// TIA Portal project "整合" (V18)

(* hardware
DEVICE "S7-1200 station_2"  S7-1200 Station
   slot 0: "Rack_0"  S7-1200 Rack  Rack  V1.0
   slot 1: "PLC_1"  CPU 1214C DC/DC/DC  6ES7 214-1AG40-0XB0  V4.1
DEVICE "PC-System_1"  SIMATIC PC station
   slot 0: "SIMATIC PC station"  Rail  SIMATIC PC-Station  V1.0
      slot 125: "Stationmanager"  Station_Manager  V6.0.4
   slot 1: "HMI_RT_1"  WinCC RT Advanced  6AV2 104-0xxxx-xxxx  17.0.0.0
      slot 33792: "主机接口"  Host interface
   slot 2: "IE general_1"  IE General  IE_CP  V8.2.0
      slot 1: "PROFINET interface"  IEGeneral.Interface.8.2.0
*)

// ===== PLC "PLC_1"  CPU 1214C DC/DC/DC =====

DATA_BLOCK "初始化用"   // DB2
{ S7_Optimized_Access := 'TRUE' }
VERSION : 0.1
// stored: InstanceOfName 初始化
"初始化"
BEGIN
END_DATA_BLOCK

DATA_BLOCK "中间变量2"   // DB3
{ S7_Optimized_Access := 'FALSE' }
VERSION : 0.1
   VAR
      "1梯1层最终调度距离" : Int;
      "2梯1层最终调度距离" : Int;
      "3梯1层最终调度距离" : Int;
      "1层上呼分配1" : Bool;
      "1层上呼分配2" : Bool;
      "1层上呼分配3" : Bool;
      "1层上呼分配4" : Bool;
      "1层上呼分配5" : Bool;
      "1层上呼分配6" : Bool;
      "1梯2层最终调度距离上" : Int;
      "1梯2层最终调度距离下" : Int;
      "2层上呼分配1" : Bool;
      "2层上呼分配2" : Bool;
      "2层上呼分配3" : Bool;
      "2层上呼分配4" : Bool;
      "2层上呼分配5" : Bool;
      "2层上呼分配6" : Bool;
      "2梯2层最终调度距离上" : Int;
      "2梯2层最终调度距离下" : Int;
      "3梯2层最终调度距离上" : Int;
      "3梯2层最终调度距离下" : Int;
      "1梯3层最终调度距离上" : Int;
      "1梯3层最终调度距离下" : Int;
      "2梯3层最终调度距离上" : Int;
      "2梯3层最终调度距离下" : Int;
      "3梯3层最终调度距离上" : Int;
      "3梯3层最终调度距离下" : Int;
      "1梯4层最终调度距离上" : Int;
      "1梯4层最终调度距离下" : Int;
      "2梯4层最终调度距离上" : Int;
      "2梯4层最终调度距离下" : Int;
      "3梯4层最终调度距离上" : Int;
      "3梯4层最终调度距离下" : Int;
      "2层下呼分配1" : Bool;
      "2层下呼分配2" : Bool;
      "2层下呼分配3" : Bool;
      "2层下呼分配4" : Bool;
      "2层下呼分配5" : Bool;
      "2层下呼分配6" : Bool;
      "3层上呼分配1" : Bool;
      "3层上呼分配2" : Bool;
      "3层上呼分配3" : Bool;
      "3层上呼分配4" : Bool;
      "3层上呼分配5" : Bool;
      "3层上呼分配6" : Bool;
      "3层下呼分配1" : Bool;
      "3层下呼分配2" : Bool;
      "3层下呼分配3" : Bool;
      "3层下呼分配4" : Bool;
      "3层下呼分配5" : Bool;
      "3层下呼分配6" : Bool;
      "4层上呼分配1" : Bool;
      "4层上呼分配2" : Bool;
      "4层上呼分配3" : Bool;
      "4层上呼分配4" : Bool;
      "4层上呼分配5" : Bool;
      "4层上呼分配6" : Bool;
      "4层下呼分配1" : Bool;
      "4层下呼分配2" : Bool;
      "4层下呼分配3" : Bool;
      "4层下呼分配4" : Bool;
      "4层下呼分配5" : Bool;
      "4层下呼分配6" : Bool;
      "1梯5层最终调度距离上" : Int;
      "1梯5层最终调度距离下" : Int;
      "2梯5层最终调度距离上" : Int;
      "2梯5层最终调度距离下" : Int;
      "3梯5层最终调度距离上" : Int;
      "3梯5层最终调度距离下" : Int;
      "5层上呼分配1" : Bool;
      "5层上呼分配2" : Bool;
      "5层上呼分配3" : Bool;
      "5层上呼分配4" : Bool;
      "5层上呼分配5" : Bool;
      "5层上呼分配6" : Bool;
      "5层下呼分配1" : Bool;
      "5层下呼分配2" : Bool;
      "5层下呼分配3" : Bool;
      "5层下呼分配4" : Bool;
      "5层下呼分配5" : Bool;
      "5层下呼分配6" : Bool;
      "1梯6层最终调度距离上" : Int;
      "1梯6层最终调度距离下" : Int;
      "2梯6层最终调度距离上" : Int;
      "2梯6层最终调度距离下" : Int;
      "3梯6层最终调度距离上" : Int;
      "3梯6层最终调度距离下" : Int;
      "6层上呼分配1" : Bool;
      "6层上呼分配2" : Bool;
      "6层上呼分配3" : Bool;
      "6层上呼分配4" : Bool;
      "6层上呼分配5" : Bool;
      "6层上呼分配6" : Bool;
      "6层下呼分配1" : Bool;
      "6层下呼分配2" : Bool;
      "6层下呼分配3" : Bool;
      "6层下呼分配4" : Bool;
      "6层下呼分配5" : Bool;
      "6层下呼分配6" : Bool;
      "1梯7层最终调度距离上" : Int;
      "1梯7层最终调度距离下" : Int;
      "2梯7层最终调度距离上" : Int;
      "2梯7层最终调度距离下" : Int;
      "3梯7层最终调度距离上" : Int;
      "3梯7层最终调度距离下" : Int;
      "7层上呼分配1" : Bool;
      "7层上呼分配2" : Bool;
      "7层上呼分配3" : Bool;
      "7层上呼分配4" : Bool;
      "7层上呼分配5" : Bool;
      "7层上呼分配6" : Bool;
      "7层下呼分配1" : Bool;
      "7层下呼分配2" : Bool;
      "7层下呼分配3" : Bool;
      "7层下呼分配4" : Bool;
      "7层下呼分配5" : Bool;
      "7层下呼分配6" : Bool;
      "1梯8层最终调度距离上" : Int;
      "1梯8层最终调度距离下" : Int;
      "2梯8层最终调度距离上" : Int;
      "2梯8层最终调度距离下" : Int;
      "3梯8层最终调度距离上" : Int;
      "3梯8层最终调度距离下" : Int;
      "8层上呼分配1" : Bool;
      "8层上呼分配2" : Bool;
      "8层上呼分配3" : Bool;
      "8层上呼分配4" : Bool;
      "8层上呼分配5" : Bool;
      "8层上呼分配6" : Bool;
      "8层下呼分配1" : Bool;
      "8层下呼分配2" : Bool;
      "8层下呼分配3" : Bool;
      "8层下呼分配4" : Bool;
      "8层下呼分配5" : Bool;
      "8层下呼分配6" : Bool;
      "1梯9层最终调度距离上" : Int;
      "1梯9层最终调度距离下" : Int;
      "2梯9层最终调度距离上" : Int;
      "2梯9层最终调度距离下" : Int;
      "3梯9层最终调度距离上" : Int;
      "3梯9层最终调度距离下" : Int;
      "9层上呼分配1" : Bool;
      "9层上呼分配2" : Bool;
      "9层上呼分配3" : Bool;
      "9层上呼分配4" : Bool;
      "9层上呼分配5" : Bool;
      "9层上呼分配6" : Bool;
      "9层下呼分配1" : Bool;
      "9层下呼分配2" : Bool;
      "9层下呼分配3" : Bool;
      "9层下呼分配4" : Bool;
      "9层下呼分配5" : Bool;
      "9层下呼分配6" : Bool;
      "1梯10层最终调度距离" : Int;
      "2梯10层最终调度距离" : Int;
      "3梯10层最终调度距离" : Int;
      "10层下呼分配1" : Bool;
      "10层下呼分配2" : Bool;
      "10层下呼分配3" : Bool;
      "10层下呼分配4" : Bool;
      "10层下呼分配5" : Bool;
      "10层下呼分配6" : Bool;
      "1号梯外呼上面无目标2" : Bool;
      "1号梯外呼上面无目标3" : Bool;
      "1号梯外呼上面无目标4" : Bool;
      "1号梯外呼上面无目标5" : Bool;
      "1号梯外呼上面无目标6" : Bool;
      "1号梯外呼上面无目标7" : Bool;
      "1号梯外呼上面无目标8" : Bool;
      "1号梯外呼上面无目标9" : Bool;
      "1号梯外呼下面无目标2" : Bool;
      "1号梯外呼下面无目标3" : Bool;
      "1号梯外呼下面无目标4" : Bool;
      "1号梯外呼下面无目标5" : Bool;
      "1号梯外呼下面无目标6" : Bool;
      "1号梯外呼下面无目标7" : Bool;
      "1号梯外呼下面无目标8" : Bool;
      "1号梯外呼下面无目标9" : Bool;
      "2号梯外呼上面无目标2" : Bool;
      "2号梯外呼上面无目标3" : Bool;
      "2号梯外呼上面无目标4" : Bool;
      "2号梯外呼上面无目标5" : Bool;
      "2号梯外呼上面无目标6" : Bool;
      "2号梯外呼上面无目标7" : Bool;
      "2号梯外呼上面无目标8" : Bool;
      "2号梯外呼上面无目标9" : Bool;
      "2号梯外呼下面无目标2" : Bool;
      "2号梯外呼下面无目标3" : Bool;
      "2号梯外呼下面无目标4" : Bool;
      "2号梯外呼下面无目标5" : Bool;
      "2号梯外呼下面无目标6" : Bool;
      "2号梯外呼下面无目标7" : Bool;
      "2号梯外呼下面无目标8" : Bool;
      "2号梯外呼下面无目标9" : Bool;
      "3号梯外呼上面无目标2" : Bool;
      "3号梯外呼上面无目标3" : Bool;
      "3号梯外呼上面无目标4" : Bool;
      "3号梯外呼上面无目标5" : Bool;
      "3号梯外呼上面无目标6" : Bool;
      "3号梯外呼上面无目标7" : Bool;
      "3号梯外呼上面无目标8" : Bool;
      "3号梯外呼上面无目标9" : Bool;
      "3号梯外呼下面无目标2" : Bool;
      "3号梯外呼下面无目标3" : Bool;
      "3号梯外呼下面无目标4" : Bool;
      "3号梯外呼下面无目标5" : Bool;
      "3号梯外呼下面无目标6" : Bool;
      "3号梯外呼下面无目标7" : Bool;
      "3号梯外呼下面无目标8" : Bool;
      "3号梯外呼下面无目标9" : Bool;
      "1号梯外呼上面有目标最大数1" : Int;
      "1号梯外呼上面有目标最大数2" : Int;
      "1号梯外呼上面有目标最大数3" : Int;
      "1号梯外呼上面有目标最大数4" : Int;
      "1号梯外呼上面有目标最大数5" : Int;
      "1号梯外呼上面有目标最大数6" : Int;
      "1号梯外呼上面有目标最大数7" : Int;
      "1号梯外呼上面有目标最大数8" : Int;
      "1号梯外呼上面有目标最大数9" : Int;
      "1号梯外呼下面有目标最小数2" : Int;
      "1号梯外呼下面有目标最小数3" : Int;
      "1号梯外呼下面有目标最小数4" : Int;
      "1号梯外呼下面有目标最小数5" : Int;
      "1号梯外呼下面有目标最小数6" : Int;
      "1号梯外呼下面有目标最小数7" : Int;
      "1号梯外呼下面有目标最小数8" : Int;
      "1号梯外呼下面有目标最小数9" : Int;
      "1号梯外呼下面有目标最小数10" : Int;
      "2号梯外呼上面有目标最大数1" : Int;
      "2号梯外呼上面有目标最大数2" : Int;
      "2号梯外呼上面有目标最大数3" : Int;
      "2号梯外呼上面有目标最大数4" : Int;
      "2号梯外呼上面有目标最大数5" : Int;
      "2号梯外呼上面有目标最大数6" : Int;
      "2号梯外呼上面有目标最大数7" : Int;
      "2号梯外呼上面有目标最大数8" : Int;
      "2号梯外呼上面有目标最大数9" : Int;
      "2号梯外呼下面有目标最小数2" : Int;
      "2号梯外呼下面有目标最小数3" : Int;
      "2号梯外呼下面有目标最小数4" : Int;
      "2号梯外呼下面有目标最小数5" : Int;
      "2号梯外呼下面有目标最小数6" : Int;
      "2号梯外呼下面有目标最小数7" : Int;
      "2号梯外呼下面有目标最小数8" : Int;
      "2号梯外呼下面有目标最小数9" : Int;
      "2号梯外呼下面有目标最小数10" : Int;
      "3号梯外呼上面有目标最大数1" : Int;
      "3号梯外呼上面有目标最大数2" : Int;
      "3号梯外呼上面有目标最大数3" : Int;
      "3号梯外呼上面有目标最大数4" : Int;
      "3号梯外呼上面有目标最大数5" : Int;
      "3号梯外呼上面有目标最大数6" : Int;
      "3号梯外呼上面有目标最大数7" : Int;
      "3号梯外呼上面有目标最大数8" : Int;
      "3号梯外呼上面有目标最大数9" : Int;
      "3号梯外呼下面有目标最小数2" : Int;
      "3号梯外呼下面有目标最小数3" : Int;
      "3号梯外呼下面有目标最小数4" : Int;
      "3号梯外呼下面有目标最小数5" : Int;
      "3号梯外呼下面有目标最小数6" : Int;
      "3号梯外呼下面有目标最小数7" : Int;
      "3号梯外呼下面有目标最小数8" : Int;
      "3号梯外呼下面有目标最小数9" : Int;
      "3号梯外呼下面有目标最小数10" : Int;
      "1号梯外呼上面有目标1" : Bool;
      "1号梯外呼上面有目标2" : Bool;
      "1号梯外呼上面有目标3" : Bool;
      "1号梯外呼上面有目标4" : Bool;
      "1号梯外呼上面有目标5" : Bool;
      "1号梯外呼上面有目标6" : Bool;
      "1号梯外呼上面有目标7" : Bool;
      "1号梯外呼上面有目标8" : Bool;
      "1号梯外呼上面有目标9" : Bool;
      "1号梯外呼下面有目标2" : Bool;
      "1号梯外呼下面有目标3" : Bool;
      "1号梯外呼下面有目标4" : Bool;
      "1号梯外呼下面有目标5" : Bool;
      "1号梯外呼下面有目标6" : Bool;
      "1号梯外呼下面有目标7" : Bool;
      "1号梯外呼下面有目标8" : Bool;
      "1号梯外呼下面有目标9" : Bool;
      "1号梯外呼下面有目标10" : Bool;
      "2号梯外呼上面有目标1" : Bool;
      "2号梯外呼上面有目标2" : Bool;
      "2号梯外呼上面有目标3" : Bool;
      "2号梯外呼上面有目标4" : Bool;
      "2号梯外呼上面有目标5" : Bool;
      "2号梯外呼上面有目标6" : Bool;
      "2号梯外呼上面有目标7" : Bool;
      "2号梯外呼上面有目标8" : Bool;
      "2号梯外呼上面有目标9" : Bool;
      "2号梯外呼下面有目标2" : Bool;
      "2号梯外呼下面有目标3" : Bool;
      "2号梯外呼下面有目标4" : Bool;
      "2号梯外呼下面有目标5" : Bool;
      "2号梯外呼下面有目标6" : Bool;
      "2号梯外呼下面有目标7" : Bool;
      "2号梯外呼下面有目标8" : Bool;
      "2号梯外呼下面有目标9" : Bool;
      "2号梯外呼下面有目标10" : Bool;
      "3号梯外呼上面有目标1" : Bool;
      "3号梯外呼上面有目标2" : Bool;
      "3号梯外呼上面有目标3" : Bool;
      "3号梯外呼上面有目标4" : Bool;
      "3号梯外呼上面有目标5" : Bool;
      "3号梯外呼上面有目标6" : Bool;
      "3号梯外呼上面有目标7" : Bool;
      "3号梯外呼上面有目标8" : Bool;
      "3号梯外呼上面有目标9" : Bool;
      "3号梯外呼下面有目标2" : Bool;
      "3号梯外呼下面有目标3" : Bool;
      "3号梯外呼下面有目标4" : Bool;
      "3号梯外呼下面有目标5" : Bool;
      "3号梯外呼下面有目标6" : Bool;
      "3号梯外呼下面有目标7" : Bool;
      "3号梯外呼下面有目标8" : Bool;
      "3号梯外呼下面有目标9" : Bool;
      "3号梯外呼下面有目标10" : Bool;
      "1号梯上行停站次数3" : Int;
      "1号梯上行停站次数4" : Int;
      "1号梯上行停站次数5" : Int;
      "1号梯上行停站次数6" : Int;
      "1号梯上行停站次数7" : Int;
      "1号梯上行停站次数8" : Int;
      "1号梯上行停站次数9" : Int;
      "1号梯上行停站次数10" : Int;
      "1号梯下行停站次数1" : Int;
      "1号梯下行停站次数2" : Int;
      "1号梯下行停站次数3" : Int;
      "1号梯下行停站次数4" : Int;
      "1号梯下行停站次数5" : Int;
      "1号梯下行停站次数6" : Int;
      "1号梯下行停站次数7" : Int;
      "1号梯下行停站次数8" : Int;
      "2号梯上行停站次数3" : Int;
      "2号梯上行停站次数4" : Int;
      "2号梯上行停站次数5" : Int;
      "2号梯上行停站次数6" : Int;
      "2号梯上行停站次数7" : Int;
      "2号梯上行停站次数8" : Int;
      "2号梯上行停站次数9" : Int;
      "2号梯上行停站次数10" : Int;
      "2号梯下行停站次数1" : Int;
      "2号梯下行停站次数2" : Int;
      "2号梯下行停站次数3" : Int;
      "2号梯下行停站次数4" : Int;
      "2号梯下行停站次数5" : Int;
      "2号梯下行停站次数6" : Int;
      "2号梯下行停站次数7" : Int;
      "2号梯下行停站次数8" : Int;
      "3号梯上行停站次数3" : Int;
      "3号梯上行停站次数4" : Int;
      "3号梯上行停站次数5" : Int;
      "3号梯上行停站次数6" : Int;
      "3号梯上行停站次数7" : Int;
      "3号梯上行停站次数8" : Int;
      "3号梯上行停站次数9" : Int;
      "3号梯上行停站次数10" : Int;
      "3号梯下行停站次数1" : Int;
      "3号梯下行停站次数2" : Int;
      "3号梯下行停站次数3" : Int;
      "3号梯下行停站次数4" : Int;
      "3号梯下行停站次数5" : Int;
      "3号梯下行停站次数6" : Int;
      "3号梯下行停站次数7" : Int;
      "3号梯下行停站次数8" : Int;
      "1号梯上行需折返停站次数10" : Int;
      "2号梯上行需折返停站次数10" : Int;
      "3号梯上行需折返停站次数10" : Int;
      "1号梯下行需折返停站次数1" : Int;
      "2号梯下行需折返停站次数1" : Int;
      "3号梯下行需折返停站次数1" : Int;
      "1号梯当前楼层数" : Int;
      "2号梯当前楼层数" : Int;
      "3号梯当前楼层数" : Int;
      "4号梯当前楼层数" : Int;
      "5号梯当前楼层数" : Int;
      "6号梯当前楼层数" : Int;
      "4梯1层最终调度距离" : Int;
      "4梯10层最终调度距离" : Int;
      "4梯2层最终调度距离上" : Int;
      "4梯2层最终调度距离下" : Int;
      "4梯3层最终调度距离上" : Int;
      "4梯3层最终调度距离下" : Int;
      "4梯4层最终调度距离上" : Int;
      "4梯4层最终调度距离下" : Int;
      "4梯5层最终调度距离上" : Int;
      "4梯5层最终调度距离下" : Int;
      "4梯6层最终调度距离上" : Int;
      "4梯6层最终调度距离下" : Int;
      "4梯7层最终调度距离上" : Int;
      "4梯7层最终调度距离下" : Int;
      "4梯8层最终调度距离上" : Int;
      "4梯8层最终调度距离下" : Int;
      "4梯9层最终调度距离上" : Int;
      "4梯9层最终调度距离下" : Int;
      "4号梯外呼上面无目标2" : Bool;
      "4号梯外呼上面无目标3" : Bool;
      "4号梯外呼上面无目标4" : Bool;
      "4号梯外呼上面无目标5" : Bool;
      "4号梯外呼上面无目标6" : Bool;
      "4号梯外呼上面无目标7" : Bool;
      "4号梯外呼上面无目标8" : Bool;
      "4号梯外呼上面无目标9" : Bool;
      "4号梯外呼下面无目标2" : Bool;
      "4号梯外呼下面无目标3" : Bool;
      "4号梯外呼下面无目标4" : Bool;
      "4号梯外呼下面无目标5" : Bool;
      "4号梯外呼下面无目标6" : Bool;
      "4号梯外呼下面无目标7" : Bool;
      "4号梯外呼下面无目标8" : Bool;
      "4号梯外呼下面无目标9" : Bool;
      "4号梯外呼上面有目标最大数1" : Int;
      "4号梯外呼上面有目标最大数2" : Int;
      "4号梯外呼上面有目标最大数3" : Int;
      "4号梯外呼上面有目标最大数4" : Int;
      "4号梯外呼上面有目标最大数5" : Int;
      "4号梯外呼上面有目标最大数6" : Int;
      "4号梯外呼上面有目标最大数7" : Int;
      "4号梯外呼上面有目标最大数8" : Int;
      "4号梯外呼上面有目标最大数9" : Int;
      "4号梯外呼下面有目标最小数2" : Int;
      "4号梯外呼下面有目标最小数3" : Int;
      "4号梯外呼下面有目标最小数4" : Int;
      "4号梯外呼下面有目标最小数5" : Int;
      "4号梯外呼下面有目标最小数6" : Int;
      "4号梯外呼下面有目标最小数7" : Int;
      "4号梯外呼下面有目标最小数8" : Int;
      "4号梯外呼下面有目标最小数9" : Int;
      "4号梯外呼下面有目标最小数10" : Int;
      "4号梯外呼上面有目标1" : Bool;
      "4号梯外呼上面有目标2" : Bool;
      "4号梯外呼上面有目标3" : Bool;
      "4号梯外呼上面有目标4" : Bool;
      "4号梯外呼上面有目标5" : Bool;
      "4号梯外呼上面有目标6" : Bool;
      "4号梯外呼上面有目标7" : Bool;
      "4号梯外呼上面有目标8" : Bool;
      "4号梯外呼上面有目标9" : Bool;
      "4号梯外呼下面有目标2" : Bool;
      "4号梯外呼下面有目标3" : Bool;
      "4号梯外呼下面有目标4" : Bool;
      "4号梯外呼下面有目标5" : Bool;
      "4号梯外呼下面有目标6" : Bool;
      "4号梯外呼下面有目标7" : Bool;
      "4号梯外呼下面有目标8" : Bool;
      "4号梯外呼下面有目标9" : Bool;
      "4号梯外呼下面有目标10" : Bool;
      "4号梯上行停站次数3" : Int;
      "4号梯上行停站次数4" : Int;
      "4号梯上行停站次数5" : Int;
      "4号梯上行停站次数6" : Int;
      "4号梯上行停站次数7" : Int;
      "4号梯上行停站次数8" : Int;
      "4号梯上行停站次数9" : Int;
      "4号梯上行停站次数10" : Int;
      "4号梯下行停站次数1" : Int;
      "4号梯下行停站次数2" : Int;
      "4号梯下行停站次数3" : Int;
      "4号梯下行停站次数4" : Int;
      "4号梯下行停站次数5" : Int;
      "4号梯下行停站次数6" : Int;
      "4号梯下行停站次数7" : Int;
      "4号梯下行停站次数8" : Int;
      "4号梯上行需折返停站次数10" : Int;
      "4号梯下行需折返停站次数1" : Int;
      "5梯1层最终调度距离" : Int;
      "5梯10层最终调度距离" : Int;
      "5梯2层最终调度距离上" : Int;
      "5梯2层最终调度距离下" : Int;
      "5梯3层最终调度距离上" : Int;
      "5梯3层最终调度距离下" : Int;
      "5梯4层最终调度距离上" : Int;
      "5梯4层最终调度距离下" : Int;
      "5梯5层最终调度距离上" : Int;
      "5梯5层最终调度距离下" : Int;
      "5梯6层最终调度距离上" : Int;
      "5梯6层最终调度距离下" : Int;
      "5梯7层最终调度距离上" : Int;
      "5梯7层最终调度距离下" : Int;
      "5梯8层最终调度距离上" : Int;
      "5梯8层最终调度距离下" : Int;
      "5梯9层最终调度距离上" : Int;
      "5梯9层最终调度距离下" : Int;
      "5号梯外呼上面无目标2" : Bool;
      "5号梯外呼上面无目标3" : Bool;
      "5号梯外呼上面无目标4" : Bool;
      "5号梯外呼上面无目标5" : Bool;
      "5号梯外呼上面无目标6" : Bool;
      "5号梯外呼上面无目标7" : Bool;
      "5号梯外呼上面无目标8" : Bool;
      "5号梯外呼上面无目标9" : Bool;
      "5号梯外呼下面无目标2" : Bool;
      "5号梯外呼下面无目标3" : Bool;
      "5号梯外呼下面无目标4" : Bool;
      "5号梯外呼下面无目标5" : Bool;
      "5号梯外呼下面无目标6" : Bool;
      "5号梯外呼下面无目标7" : Bool;
      "5号梯外呼下面无目标8" : Bool;
      "5号梯外呼下面无目标9" : Bool;
      "5号梯外呼上面有目标最大数1" : Int;
      "5号梯外呼上面有目标最大数2" : Int;
      "5号梯外呼上面有目标最大数3" : Int;
      "5号梯外呼上面有目标最大数4" : Int;
      "5号梯外呼上面有目标最大数5" : Int;
      "5号梯外呼上面有目标最大数6" : Int;
      "5号梯外呼上面有目标最大数7" : Int;
      "5号梯外呼上面有目标最大数8" : Int;
      "5号梯外呼上面有目标最大数9" : Int;
      "5号梯外呼下面有目标最小数2" : Int;
      "5号梯外呼下面有目标最小数3" : Int;
      "5号梯外呼下面有目标最小数4" : Int;
      "5号梯外呼下面有目标最小数5" : Int;
      "5号梯外呼下面有目标最小数6" : Int;
      "5号梯外呼下面有目标最小数7" : Int;
      "5号梯外呼下面有目标最小数8" : Int;
      "5号梯外呼下面有目标最小数9" : Int;
      "5号梯外呼下面有目标最小数10" : Int;
      "5号梯外呼上面有目标1" : Bool;
      "5号梯外呼上面有目标2" : Bool;
      "5号梯外呼上面有目标3" : Bool;
      "5号梯外呼上面有目标4" : Bool;
      "5号梯外呼上面有目标5" : Bool;
      "5号梯外呼上面有目标6" : Bool;
      "5号梯外呼上面有目标7" : Bool;
      "5号梯外呼上面有目标8" : Bool;
      "5号梯外呼上面有目标9" : Bool;
      "5号梯外呼下面有目标2" : Bool;
      "5号梯外呼下面有目标3" : Bool;
      "5号梯外呼下面有目标4" : Bool;
      "5号梯外呼下面有目标5" : Bool;
      "5号梯外呼下面有目标6" : Bool;
      "5号梯外呼下面有目标7" : Bool;
      "5号梯外呼下面有目标8" : Bool;
      "5号梯外呼下面有目标9" : Bool;
      "5号梯外呼下面有目标10" : Bool;
      "5号梯上行停站次数3" : Int;
      "5号梯上行停站次数4" : Int;
      "5号梯上行停站次数5" : Int;
      "5号梯上行停站次数6" : Int;
      "5号梯上行停站次数7" : Int;
      "5号梯上行停站次数8" : Int;
      "5号梯上行停站次数9" : Int;
      "5号梯上行停站次数10" : Int;
      "5号梯下行停站次数1" : Int;
      "5号梯下行停站次数2" : Int;
      "5号梯下行停站次数3" : Int;
      "5号梯下行停站次数4" : Int;
      "5号梯下行停站次数5" : Int;
      "5号梯下行停站次数6" : Int;
      "5号梯下行停站次数7" : Int;
      "5号梯下行停站次数8" : Int;
      "5号梯上行需折返停站次数10" : Int;
      "5号梯下行需折返停站次数1" : Int;
      "6梯1层最终调度距离" : Int;
      "6梯10层最终调度距离" : Int;
      "6梯2层最终调度距离上" : Int;
      "6梯2层最终调度距离下" : Int;
      "6梯3层最终调度距离上" : Int;
      "6梯3层最终调度距离下" : Int;
      "6梯4层最终调度距离上" : Int;
      "6梯4层最终调度距离下" : Int;
      "6梯5层最终调度距离上" : Int;
      "6梯5层最终调度距离下" : Int;
      "6梯6层最终调度距离上" : Int;
      "6梯6层最终调度距离下" : Int;
      "6梯7层最终调度距离上" : Int;
      "6梯7层最终调度距离下" : Int;
      "6梯8层最终调度距离上" : Int;
      "6梯8层最终调度距离下" : Int;
      "6梯9层最终调度距离上" : Int;
      "6梯9层最终调度距离下" : Int;
      "6号梯外呼上面无目标2" : Bool;
      "6号梯外呼上面无目标3" : Bool;
      "6号梯外呼上面无目标4" : Bool;
      "6号梯外呼上面无目标5" : Bool;
      "6号梯外呼上面无目标6" : Bool;
      "6号梯外呼上面无目标7" : Bool;
      "6号梯外呼上面无目标8" : Bool;
      "6号梯外呼上面无目标9" : Bool;
      "6号梯外呼下面无目标2" : Bool;
      "6号梯外呼下面无目标3" : Bool;
      "6号梯外呼下面无目标4" : Bool;
      "6号梯外呼下面无目标5" : Bool;
      "6号梯外呼下面无目标6" : Bool;
      "6号梯外呼下面无目标7" : Bool;
      "6号梯外呼下面无目标8" : Bool;
      "6号梯外呼下面无目标9" : Bool;
      "6号梯外呼上面有目标最大数1" : Int;
      "6号梯外呼上面有目标最大数2" : Int;
      "6号梯外呼上面有目标最大数3" : Int;
      "6号梯外呼上面有目标最大数4" : Int;
      "6号梯外呼上面有目标最大数5" : Int;
      "6号梯外呼上面有目标最大数6" : Int;
      "6号梯外呼上面有目标最大数7" : Int;
      "6号梯外呼上面有目标最大数8" : Int;
      "6号梯外呼上面有目标最大数9" : Int;
      "6号梯外呼下面有目标最小数2" : Int;
      "6号梯外呼下面有目标最小数3" : Int;
      "6号梯外呼下面有目标最小数4" : Int;
      "6号梯外呼下面有目标最小数5" : Int;
      "6号梯外呼下面有目标最小数6" : Int;
      "6号梯外呼下面有目标最小数7" : Int;
      "6号梯外呼下面有目标最小数8" : Int;
      "6号梯外呼下面有目标最小数9" : Int;
      "6号梯外呼下面有目标最小数10" : Int;
      "6号梯外呼上面有目标1" : Bool;
      "6号梯外呼上面有目标2" : Bool;
      "6号梯外呼上面有目标3" : Bool;
      "6号梯外呼上面有目标4" : Bool;
      "6号梯外呼上面有目标5" : Bool;
      "6号梯外呼上面有目标6" : Bool;
      "6号梯外呼上面有目标7" : Bool;
      "6号梯外呼上面有目标8" : Bool;
      "6号梯外呼上面有目标9" : Bool;
      "6号梯外呼下面有目标2" : Bool;
      "6号梯外呼下面有目标3" : Bool;
      "6号梯外呼下面有目标4" : Bool;
      "6号梯外呼下面有目标5" : Bool;
      "6号梯外呼下面有目标6" : Bool;
      "6号梯外呼下面有目标7" : Bool;
      "6号梯外呼下面有目标8" : Bool;
      "6号梯外呼下面有目标9" : Bool;
      "6号梯外呼下面有目标10" : Bool;
      "6号梯上行停站次数3" : Int;
      "6号梯上行停站次数4" : Int;
      "6号梯上行停站次数5" : Int;
      "6号梯上行停站次数6" : Int;
      "6号梯上行停站次数7" : Int;
      "6号梯上行停站次数8" : Int;
      "6号梯上行停站次数9" : Int;
      "6号梯上行停站次数10" : Int;
      "6号梯下行停站次数1" : Int;
      "6号梯下行停站次数2" : Int;
      "6号梯下行停站次数3" : Int;
      "6号梯下行停站次数4" : Int;
      "6号梯下行停站次数5" : Int;
      "6号梯下行停站次数6" : Int;
      "6号梯下行停站次数7" : Int;
      "6号梯下行停站次数8" : Int;
      "6号梯上行需折返停站次数10" : Int;
      "6号梯下行需折返停站次数1" : Int;
      "1号梯转换后载重量" : Int;
      "2号梯转换后载重量" : Int;
      "3号梯转换后载重量" : Int;
      "4号梯转换后载重量" : Int;
      "5号梯转换后载重量" : Int;
      "6号梯转换后载重量" : Int;
      限重分配1 : Int := 900;
      限重分配2 : Int := 1200;
      限重分配3 : Int := 1200;
      限重分配4 : Int := 1200;
      限重分配5 : Int := 1650;
      限重分配6 : Int := 1850;
      就近运动电梯1 : Bool;
      就近运动电梯2 : Bool;
      就近运动电梯3 : Bool;
      就近运动电梯4 : Bool;
      就近运动电梯5 : Bool;
      就近运动电梯6 : Bool;
   END_VAR
BEGIN
END_DATA_BLOCK

DATA_BLOCK "输入"   // DB10
{ S7_Optimized_Access := 'FALSE' }
VERSION : 0.1
   VAR
      "1层上行呼梯按钮" : Bool;
      "2层上行呼梯按钮" : Bool;
      "3层上行呼梯按钮" : Bool;
      "4层上行呼梯按钮" : Bool;
      "5层上行呼梯按钮" : Bool;
      "6层上行呼梯按钮" : Bool;
      "7层上行呼梯按钮" : Bool;
      "8层上行呼梯按钮" : Bool;
      "9层上行呼梯按钮" : Bool;
      "2层下行呼梯按钮" : Bool;
      "3层下行呼梯按钮" : Bool;
      "4层下行呼梯按钮" : Bool;
      "5层下行呼梯按钮" : Bool;
      "6层下行呼梯按钮" : Bool;
      "7层下行呼梯按钮" : Bool;
      "8层下行呼梯按钮" : Bool;
      "9层下行呼梯按钮" : Bool;
      "10层下行呼梯按钮" : Bool;
      "1号梯轿内选层按钮1" : Bool;
      "1号梯轿内选层按钮2" : Bool;
      "1号梯轿内选层按钮3" : Bool;
      "1号梯轿内选层按钮4" : Bool;
      "1号梯轿内选层按钮5" : Bool;
      "1号梯轿内选层按钮6" : Bool;
      "1号梯轿内选层按钮7" : Bool;
      "1号梯轿内选层按钮8" : Bool;
      "1号梯轿内选层按钮9" : Bool;
      "1号梯轿内选层按钮10" : Bool;
      "1号梯轿内开门按钮" : Bool;
      "1号梯轿内关门按钮" : Bool;
      "1号梯光幕信号" : Bool;
      "1号梯检修信号" : Bool;
      "1号梯轿厢门锁信号" : Bool;
      "1号梯1楼层门锁信号" : Bool;
      "1号梯2楼层门锁信号" : Bool;
      "1号梯3楼层门锁信号" : Bool;
      "1号梯4楼层门锁信号" : Bool;
      "1号梯5楼层门锁信号" : Bool;
      "1号梯6楼层门锁信号" : Bool;
      "1号梯7楼层门锁信号" : Bool;
      "1号梯8楼层门锁信号" : Bool;
      "1号梯9楼层门锁信号" : Bool;
      "1号梯10楼层门锁信号" : Bool;
      "1号梯开门到位" : Bool;
      "1号梯关门到位" : Bool;
      "1号梯上平层信号" : Bool;
      "1号梯下平层信号" : Bool;
      "1号梯上端站第1限位" : Bool;
      "1号梯上端站第2限位" : Bool;
      "1号梯下端站第1限位" : Bool;
      "1号梯下端站第2限位" : Bool;
      "2号梯轿内选层按钮1" : Bool;
      "2号梯轿内选层按钮2" : Bool;
      "2号梯轿内选层按钮3" : Bool;
      "2号梯轿内选层按钮4" : Bool;
      "2号梯轿内选层按钮5" : Bool;
      "2号梯轿内选层按钮6" : Bool;
      "2号梯轿内选层按钮7" : Bool;
      "2号梯轿内选层按钮8" : Bool;
      "2号梯轿内选层按钮9" : Bool;
      "2号梯轿内选层按钮10" : Bool;
      "2号梯轿内开门按钮" : Bool;
      "2号梯轿内关门按钮" : Bool;
      "2号梯光幕信号" : Bool;
      "2号梯检修信号" : Bool;
      "2号梯轿厢门锁信号" : Bool;
      "2号梯1楼层门锁信号" : Bool;
      "2号梯2楼层门锁信号" : Bool;
      "2号梯3楼层门锁信号" : Bool;
      "2号梯4楼层门锁信号" : Bool;
      "2号梯5楼层门锁信号" : Bool;
      "2号梯6楼层门锁信号" : Bool;
      "2号梯7楼层门锁信号" : Bool;
      "2号梯8楼层门锁信号" : Bool;
      "2号梯9楼层门锁信号" : Bool;
      "2号梯10楼层门锁信号" : Bool;
      "2号梯开门到位" : Bool;
      "2号梯关门到位" : Bool;
      "2号梯上平层信号" : Bool;
      "2号梯下平层信号" : Bool;
      "2号梯上端站第1限位" : Bool;
      "2号梯上端站第2限位" : Bool;
      "2号梯下端站第1限位" : Bool;
      "2号梯下端站第2限位" : Bool;
      "3号梯轿内选层按钮1" : Bool;
      "3号梯轿内选层按钮2" : Bool;
      "3号梯轿内选层按钮3" : Bool;
      "3号梯轿内选层按钮4" : Bool;
      "3号梯轿内选层按钮5" : Bool;
      "3号梯轿内选层按钮6" : Bool;
      "3号梯轿内选层按钮7" : Bool;
      "3号梯轿内选层按钮8" : Bool;
      "3号梯轿内选层按钮9" : Bool;
      "3号梯轿内选层按钮10" : Bool;
      "3号梯轿内开门按钮" : Bool;
      "3号梯轿内关门按钮" : Bool;
      "3号梯光幕信号" : Bool;
      "3号梯检修信号" : Bool;
      "3号梯轿厢门锁信号" : Bool;
      "3号梯1楼层门锁信号" : Bool;
      "3号梯2楼层门锁信号" : Bool;
      "3号梯3楼层门锁信号" : Bool;
      "3号梯4楼层门锁信号" : Bool;
      "3号梯5楼层门锁信号" : Bool;
      "3号梯6楼层门锁信号" : Bool;
      "3号梯7楼层门锁信号" : Bool;
      "3号梯8楼层门锁信号" : Bool;
      "3号梯9楼层门锁信号" : Bool;
      "3号梯10楼层门锁信号" : Bool;
      "3号梯开门到位" : Bool;
      "3号梯关门到位" : Bool;
      "3号梯上平层信号" : Bool;
      "3号梯下平层信号" : Bool;
      "3号梯上端站第1限位" : Bool;
      "3号梯上端站第2限位" : Bool;
      "3号梯下端站第1限位" : Bool;
      "3号梯下端站第2限位" : Bool;
      "4号梯轿内选层按钮1" : Bool;
      "4号梯轿内选层按钮2" : Bool;
      "4号梯轿内选层按钮3" : Bool;
      "4号梯轿内选层按钮4" : Bool;
      "4号梯轿内选层按钮5" : Bool;
      "4号梯轿内选层按钮6" : Bool;
      "4号梯轿内选层按钮7" : Bool;
      "4号梯轿内选层按钮8" : Bool;
      "4号梯轿内选层按钮9" : Bool;
      "4号梯轿内选层按钮10" : Bool;
      "4号梯轿内开门按钮" : Bool;
      "4号梯轿内关门按钮" : Bool;
      "4号梯光幕信号" : Bool;
      "4号梯检修信号" : Bool;
      "4号梯轿厢门锁信号" : Bool;
      "4号梯1楼层门锁信号" : Bool;
      "4号梯2楼层门锁信号" : Bool;
      "4号梯3楼层门锁信号" : Bool;
      "4号梯4楼层门锁信号" : Bool;
      "4号梯5楼层门锁信号" : Bool;
      "4号梯6楼层门锁信号" : Bool;
      "4号梯7楼层门锁信号" : Bool;
      "4号梯8楼层门锁信号" : Bool;
      "4号梯9楼层门锁信号" : Bool;
      "4号梯10楼层门锁信号" : Bool;
      "4号梯开门到位" : Bool;
      "4号梯关门到位" : Bool;
      "4号梯上平层信号" : Bool;
      "4号梯下平层信号" : Bool;
      "4号梯上端站第1限位" : Bool;
      "4号梯上端站第2限位" : Bool;
      "4号梯下端站第1限位" : Bool;
      "4号梯下端站第2限位" : Bool;
      "5号梯轿内选层按钮1" : Bool;
      "5号梯轿内选层按钮2" : Bool;
      "5号梯轿内选层按钮3" : Bool;
      "5号梯轿内选层按钮4" : Bool;
      "5号梯轿内选层按钮5" : Bool;
      "5号梯轿内选层按钮6" : Bool;
      "5号梯轿内选层按钮7" : Bool;
      "5号梯轿内选层按钮8" : Bool;
      "5号梯轿内选层按钮9" : Bool;
      "5号梯轿内选层按钮10" : Bool;
      "5号梯轿内开门按钮" : Bool;
      "5号梯轿内关门按钮" : Bool;
      "5号梯光幕信号" : Bool;
      "5号梯检修信号" : Bool;
      "5号梯轿厢门锁信号" : Bool;
      "5号梯1楼层门锁信号" : Bool;
      "5号梯2楼层门锁信号" : Bool;
      "5号梯3楼层门锁信号" : Bool;
      "5号梯4楼层门锁信号" : Bool;
      "5号梯5楼层门锁信号" : Bool;
      "5号梯6楼层门锁信号" : Bool;
      "5号梯7楼层门锁信号" : Bool;
      "5号梯8楼层门锁信号" : Bool;
      "5号梯9楼层门锁信号" : Bool;
      "5号梯10楼层门锁信号" : Bool;
      "5号梯开门到位" : Bool;
      "5号梯关门到位" : Bool;
      "5号梯上平层信号" : Bool;
      "5号梯下平层信号" : Bool;
      "5号梯上端站第1限位" : Bool;
      "5号梯上端站第2限位" : Bool;
      "5号梯下端站第1限位" : Bool;
      "5号梯下端站第2限位" : Bool;
      "6号梯轿内选层按钮1" : Bool;
      "6号梯轿内选层按钮2" : Bool;
      "6号梯轿内选层按钮3" : Bool;
      "6号梯轿内选层按钮4" : Bool;
      "6号梯轿内选层按钮5" : Bool;
      "6号梯轿内选层按钮6" : Bool;
      "6号梯轿内选层按钮7" : Bool;
      "6号梯轿内选层按钮8" : Bool;
      "6号梯轿内选层按钮9" : Bool;
      "6号梯轿内选层按钮10" : Bool;
      "6号梯轿内开门按钮" : Bool;
      "6号梯轿内关门按钮" : Bool;
      "6号梯光幕信号" : Bool;
      "6号梯检修信号" : Bool;
      "6号梯轿厢门锁信号" : Bool;
      "6号梯1楼层门锁信号" : Bool;
      "6号梯2楼层门锁信号" : Bool;
      "6号梯3楼层门锁信号" : Bool;
      "6号梯4楼层门锁信号" : Bool;
      "6号梯5楼层门锁信号" : Bool;
      "6号梯6楼层门锁信号" : Bool;
      "6号梯7楼层门锁信号" : Bool;
      "6号梯8楼层门锁信号" : Bool;
      "6号梯9楼层门锁信号" : Bool;
      "6号梯10楼层门锁信号" : Bool;
      "6号梯开门到位" : Bool;
      "6号梯关门到位" : Bool;
      "6号梯上平层信号" : Bool;
      "6号梯下平层信号" : Bool;
      "6号梯上端站第1限位" : Bool;
      "6号梯上端站第2限位" : Bool;
      "6号梯下端站第1限位" : Bool;
      "6号梯下端站第2限位" : Bool;
      自动运行信号 : Bool;
      "1号梯当前载重量" : Word;
      "2号梯当前载重量" : Word;
      "3号梯当前载重量" : Word;
      "4号梯当前载重量" : Word;
      "5号梯当前载重量" : Word;
      "6号梯当前载重量" : Word;
   END_VAR
BEGIN
END_DATA_BLOCK

DATA_BLOCK "输出"   // DB11
{ S7_Optimized_Access := 'FALSE' }
VERSION : 0.1
   VAR
      "1层上行呼梯按钮指示灯" : Bool;
      "2层上行呼梯按钮指示灯" : Bool;
      "3层上行呼梯按钮指示灯" : Bool;
      "4层上行呼梯按钮指示灯" : Bool;
      "5层上行呼梯按钮指示灯" : Bool;
      "6层上行呼梯按钮指示灯" : Bool;
      "7层上行呼梯按钮指示灯" : Bool;
      "8层上行呼梯按钮指示灯" : Bool;
      "9层上行呼梯按钮指示灯" : Bool;
      "2层下行呼梯按钮指示灯" : Bool;
      "3层下行呼梯按钮指示灯" : Bool;
      "4层下行呼梯按钮指示灯" : Bool;
      "5层下行呼梯按钮指示灯" : Bool;
      "6层下行呼梯按钮指示灯" : Bool;
      "7层下行呼梯按钮指示灯" : Bool;
      "8层下行呼梯按钮指示灯" : Bool;
      "9层下行呼梯按钮指示灯" : Bool;
      "10层下行呼梯按钮指示灯" : Bool;
      "1号梯1层按钮指示灯" : Bool;
      "1号梯2层按钮指示灯" : Bool;
      "1号梯3层按钮指示灯" : Bool;
      "1号梯4层按钮指示灯" : Bool;
      "1号梯5层按钮指示灯" : Bool;
      "1号梯6层按钮指示灯" : Bool;
      "1号梯7层按钮指示灯" : Bool;
      "1号梯8层按钮指示灯" : Bool;
      "1号梯9层按钮指示灯" : Bool;
      "1号梯10层按钮指示灯" : Bool;
      "1号梯LEDa" : Bool;
      "1号梯LEDb" : Bool;
      "1号梯LEDc" : Bool;
      "1号梯LEDd" : Bool;
      "1号梯LEDe" : Bool;
      "1号梯LEDf" : Bool;
      "1号梯LEDg" : Bool;
      "1号梯LEDh" : Bool;
      "1号梯LEDi" : Bool;
      "1号梯LEDj" : Bool;
      "1号梯LEDk" : Bool;
      "1号梯LEDl" : Bool;
      "1号梯LEDm" : Bool;
      "1号梯LEDn" : Bool;
      "1号梯上行指示" : Bool;
      "1号梯下行指示" : Bool;
      "1号梯故障指示" : Bool;
      "1号梯照明指示" : Bool;
      "1号梯风扇指示" : Bool;
      "1号梯满载指示" : Bool;
      "1号梯电机启动信号" : Bool;
      "1号梯上行接触器" : Bool;
      "1号梯下行接触器" : Bool;
      "1号梯高速接触器" : Bool;
      "1号梯低速接触器" : Bool;
      "1号梯开门继电器" : Bool;
      "1号梯关门继电器" : Bool;
      "1号梯1级减速制动" : Bool;
      "1号梯2级减速制动" : Bool;
      "1号梯3级减速制动" : Bool;
      "2号梯1层按钮指示灯" : Bool;
      "2号梯2层按钮指示灯" : Bool;
      "2号梯3层按钮指示灯" : Bool;
      "2号梯4层按钮指示灯" : Bool;
      "2号梯5层按钮指示灯" : Bool;
      "2号梯6层按钮指示灯" : Bool;
      "2号梯7层按钮指示灯" : Bool;
      "2号梯8层按钮指示灯" : Bool;
      "2号梯9层按钮指示灯" : Bool;
      "2号梯10层按钮指示灯" : Bool;
      "2号梯LEDa" : Bool;
      "2号梯LEDb" : Bool;
      "2号梯LEDc" : Bool;
      "2号梯LEDd" : Bool;
      "2号梯LEDe" : Bool;
      "2号梯LEDf" : Bool;
      "2号梯LEDg" : Bool;
      "2号梯LEDh" : Bool;
      "2号梯LEDi" : Bool;
      "2号梯LEDj" : Bool;
      "2号梯LEDk" : Bool;
      "2号梯LEDl" : Bool;
      "2号梯LEDm" : Bool;
      "2号梯LEDn" : Bool;
      "2号梯上行指示" : Bool;
      "2号梯下行指示" : Bool;
      "2号梯故障指示" : Bool;
      "2号梯照明指示" : Bool;
      "2号梯风扇指示" : Bool;
      "2号梯满载指示" : Bool;
      "2号梯电机启动信号" : Bool;
      "2号梯上行接触器" : Bool;
      "2号梯下行接触器" : Bool;
      "2号梯高速接触器" : Bool;
      "2号梯低速接触器" : Bool;
      "2号梯开门继电器" : Bool;
      "2号梯关门继电器" : Bool;
      "2号梯1级减速制动" : Bool;
      "2号梯2级减速制动" : Bool;
      "2号梯3级减速制动" : Bool;
      "3号梯1层按钮指示灯" : Bool;
      "3号梯2层按钮指示灯" : Bool;
      "3号梯3层按钮指示灯" : Bool;
      "3号梯4层按钮指示灯" : Bool;
      "3号梯5层按钮指示灯" : Bool;
      "3号梯6层按钮指示灯" : Bool;
      "3号梯7层按钮指示灯" : Bool;
      "3号梯8层按钮指示灯" : Bool;
      "3号梯9层按钮指示灯" : Bool;
      "3号梯10层按钮指示灯" : Bool;
      "3号梯LEDa" : Bool;
      "3号梯LEDb" : Bool;
      "3号梯LEDc" : Bool;
      "3号梯LEDd" : Bool;
      "3号梯LEDe" : Bool;
      "3号梯LEDf" : Bool;
      "3号梯LEDg" : Bool;
      "3号梯LEDh" : Bool;
      "3号梯LEDi" : Bool;
      "3号梯LEDj" : Bool;
      "3号梯LEDk" : Bool;
      "3号梯LEDl" : Bool;
      "3号梯LEDm" : Bool;
      "3号梯LEDn" : Bool;
      "3号梯上行指示" : Bool;
      "3号梯下行指示" : Bool;
      "3号梯故障指示" : Bool;
      "3号梯照明指示" : Bool;
      "3号梯风扇指示" : Bool;
      "3号梯满载指示" : Bool;
      "3号梯电机启动信号" : Bool;
      "3号梯上行接触器" : Bool;
      "3号梯下行接触器" : Bool;
      "3号梯高速接触器" : Bool;
      "3号梯低速接触器" : Bool;
      "3号梯开门继电器" : Bool;
      "3号梯关门继电器" : Bool;
      "3号梯1级减速制动" : Bool;
      "3号梯2级减速制动" : Bool;
      "3号梯3级减速制动" : Bool;
      "4号梯1层按钮指示灯" : Bool;
      "4号梯2层按钮指示灯" : Bool;
      "4号梯3层按钮指示灯" : Bool;
      "4号梯4层按钮指示灯" : Bool;
      "4号梯5层按钮指示灯" : Bool;
      "4号梯6层按钮指示灯" : Bool;
      "4号梯7层按钮指示灯" : Bool;
      "4号梯8层按钮指示灯" : Bool;
      "4号梯9层按钮指示灯" : Bool;
      "4号梯10层按钮指示灯" : Bool;
      "4号梯LEDa" : Bool;
      "4号梯LEDb" : Bool;
      "4号梯LEDc" : Bool;
      "4号梯LEDd" : Bool;
      "4号梯LEDe" : Bool;
      "4号梯LEDf" : Bool;
      "4号梯LEDg" : Bool;
      "4号梯LEDh" : Bool;
      "4号梯LEDi" : Bool;
      "4号梯LEDj" : Bool;
      "4号梯LEDk" : Bool;
      "4号梯LEDl" : Bool;
      "4号梯LEDm" : Bool;
      "4号梯LEDn" : Bool;
      "4号梯上行指示" : Bool;
      "4号梯下行指示" : Bool;
      "4号梯故障指示" : Bool;
      "4号梯照明指示" : Bool;
      "4号梯风扇指示" : Bool;
      "4号梯满载指示" : Bool;
      "4号梯电机启动信号" : Bool;
      "4号梯上行接触器" : Bool;
      "4号梯下行接触器" : Bool;
      "4号梯高速接触器" : Bool;
      "4号梯低速接触器" : Bool;
      "4号梯开门继电器" : Bool;
      "4号梯关门继电器" : Bool;
      "4号梯1级减速制动" : Bool;
      "4号梯2级减速制动" : Bool;
      "4号梯3级减速制动" : Bool;
      "5号梯1层按钮指示灯" : Bool;
      "5号梯2层按钮指示灯" : Bool;
      "5号梯3层按钮指示灯" : Bool;
      "5号梯4层按钮指示灯" : Bool;
      "5号梯5层按钮指示灯" : Bool;
      "5号梯6层按钮指示灯" : Bool;
      "5号梯7层按钮指示灯" : Bool;
      "5号梯8层按钮指示灯" : Bool;
      "5号梯9层按钮指示灯" : Bool;
      "5号梯10层按钮指示灯" : Bool;
      "5号梯LEDa" : Bool;
      "5号梯LEDb" : Bool;
      "5号梯LEDc" : Bool;
      "5号梯LEDd" : Bool;
      "5号梯LEDe" : Bool;
      "5号梯LEDf" : Bool;
      "5号梯LEDg" : Bool;
      "5号梯LEDh" : Bool;
      "5号梯LEDi" : Bool;
      "5号梯LEDj" : Bool;
      "5号梯LEDk" : Bool;
      "5号梯LEDl" : Bool;
      "5号梯LEDm" : Bool;
      "5号梯LEDn" : Bool;
      "5号梯上行指示" : Bool;
      "5号梯下行指示" : Bool;
      "5号梯故障指示" : Bool;
      "5号梯照明指示" : Bool;
      "5号梯风扇指示" : Bool;
      "5号梯满载指示" : Bool;
      "5号梯电机启动信号" : Bool;
      "5号梯上行接触器" : Bool;
      "5号梯下行接触器" : Bool;
      "5号梯高速接触器" : Bool;
      "5号梯低速接触器" : Bool;
      "5号梯开门继电器" : Bool;
      "5号梯关门继电器" : Bool;
      "5号梯1级减速制动" : Bool;
      "5号梯2级减速制动" : Bool;
      "5号梯3级减速制动" : Bool;
      "6号梯1层按钮指示灯" : Bool;
      "6号梯2层按钮指示灯" : Bool;
      "6号梯3层按钮指示灯" : Bool;
      "6号梯4层按钮指示灯" : Bool;
      "6号梯5层按钮指示灯" : Bool;
      "6号梯6层按钮指示灯" : Bool;
      "6号梯7层按钮指示灯" : Bool;
      "6号梯8层按钮指示灯" : Bool;
      "6号梯9层按钮指示灯" : Bool;
      "6号梯10层按钮指示灯" : Bool;
      "6号梯LEDa" : Bool;
      "6号梯LEDb" : Bool;
      "6号梯LEDc" : Bool;
      "6号梯LEDd" : Bool;
      "6号梯LEDe" : Bool;
      "6号梯LEDf" : Bool;
      "6号梯LEDg" : Bool;
      "6号梯LEDh" : Bool;
      "6号梯LEDi" : Bool;
      "6号梯LEDj" : Bool;
      "6号梯LEDk" : Bool;
      "6号梯LEDl" : Bool;
      "6号梯LEDm" : Bool;
      "6号梯LEDn" : Bool;
      "6号梯上行指示" : Bool;
      "6号梯下行指示" : Bool;
      "6号梯故障指示" : Bool;
      "6号梯照明指示" : Bool;
      "6号梯风扇指示" : Bool;
      "6号梯满载指示" : Bool;
      "6号梯电机启动信号" : Bool;
      "6号梯上行接触器" : Bool;
      "6号梯下行接触器" : Bool;
      "6号梯高速接触器" : Bool;
      "6号梯低速接触器" : Bool;
      "6号梯开门继电器" : Bool;
      "6号梯关门继电器" : Bool;
      "6号梯1级减速制动" : Bool;
      "6号梯2级减速制动" : Bool;
      "6号梯3级减速制动" : Bool;
      准备就绪信号 : Bool;
   END_VAR
BEGIN
END_DATA_BLOCK

DATA_BLOCK "中间变量1"   // DB13
{ S7_Optimized_Access := 'FALSE' }
VERSION : 0.1
   VAR
      "1号梯高速初始化" : Bool;
      "2号梯高速初始化" : Bool;
      "3号梯高速初始化" : Bool;
      "4号梯高速初始化" : Bool;
      "5号梯高速初始化" : Bool;
      "6号梯高速初始化" : Bool;
      是否高速1 : Bool;
      是否高速2 : Bool;
      是否高速3 : Bool;
      是否高速4 : Bool;
      是否高速5 : Bool;
      是否高速6 : Bool;
      高速延时1 : Time;
      高速延时2 : Time;
      高速延时3 : Time;
      高速延时4 : Time;
      高速延时5 : Time;
      高速延时6 : Time;
      上下平层同时为1梯1 : Bool;
      上下平层同时为1梯2 : Bool;
      上下平层同时为1梯3 : Bool;
      上下平层同时为1梯4 : Bool;
      上下平层同时为1梯5 : Bool;
      上下平层同时为1梯6 : Bool;
      特殊上行将要停梯1 : Bool;
      特殊上行将要停梯2 : Bool;
      特殊上行将要停梯3 : Bool;
      特殊上行将要停梯4 : Bool;
      特殊上行将要停梯5 : Bool;
      特殊上行将要停梯6 : Bool;
      特殊下行将要停梯1 : Bool;
      特殊下行将要停梯2 : Bool;
      特殊下行将要停梯3 : Bool;
      特殊下行将要停梯4 : Bool;
      特殊下行将要停梯5 : Bool;
      特殊下行将要停梯6 : Bool;
      "1号梯正处于故障中" : Bool;
      "2号梯正处于故障中" : Bool;
      "3号梯正处于故障中" : Bool;
      "4号梯正处于故障中" : Bool;
      "5号梯正处于故障中" : Bool;
      "6号梯正处于故障中" : Bool;
      "1号梯存在安全隐患（光幕）" : Bool;
      "2号梯存在安全隐患（光幕）" : Bool;
      "3号梯存在安全隐患（光幕）" : Bool;
      "4号梯存在安全隐患（光幕）" : Bool;
      "5号梯存在安全隐患（光幕）" : Bool;
      "6号梯存在安全隐患（光幕）" : Bool;
      "1号梯当前楼层数" : Int;
      "2号梯当前楼层数" : Int;
      "3号梯当前楼层数" : Int;
      "4号梯当前楼层数" : Int;
      "5号梯当前楼层数" : Int;
      "6号梯当前楼层数" : Int;
      "1号梯初始化楼层数" : Int := 1;
      "2号梯初始化楼层数" : Int := 1;
      "3号梯初始化楼层数" : Int := 10;
      "4号梯初始化楼层数" : Int := 10;
      "5号梯初始化楼层数" : Int := 10;
      "6号梯初始化楼层数" : Int := 10;
      "1号梯是否到达端限" : Bool;
      "2号梯是否到达端限" : Bool;
      "3号梯是否到达端限" : Bool;
      "4号梯是否到达端限" : Bool;
      "5号梯是否到达端限" : Bool;
      "6号梯是否到达端限" : Bool;
      "1号梯初始化方向上行" : Bool;
      "2号梯初始化方向上行" : Bool;
      "3号梯初始化方向上行" : Bool;
      "4号梯初始化方向上行" : Bool;
      "5号梯初始化方向上行" : Bool;
      "6号梯初始化方向上行" : Bool;
      "1号梯初始化方向下行" : Bool;
      "2号梯初始化方向下行" : Bool;
      "3号梯初始化方向下行" : Bool;
      "4号梯初始化方向下行" : Bool;
      "5号梯初始化方向下行" : Bool;
      "6号梯初始化方向下行" : Bool;
      检修方向上行1 : Bool;
      检修方向上行2 : Bool;
      检修方向上行3 : Bool;
      检修方向上行4 : Bool;
      检修方向上行5 : Bool;
      检修方向上行6 : Bool;
      检修方向下行1 : Bool;
      检修方向下行2 : Bool;
      检修方向下行3 : Bool;
      检修方向下行4 : Bool;
      检修方向下行5 : Bool;
      检修方向下行6 : Bool;
      "1号梯初始化低速运行" : Bool;
      "2号梯初始化低速运行" : Bool;
      "3号梯初始化低速运行" : Bool;
      "4号梯初始化低速运行" : Bool;
      "5号梯初始化低速运行" : Bool;
      "6号梯初始化低速运行" : Bool;
      "1号梯初始化上行接触器" : Bool;
      "2号梯初始化上行接触器" : Bool;
      "3号梯初始化上行接触器" : Bool;
      "4号梯初始化上行接触器" : Bool;
      "5号梯初始化上行接触器" : Bool;
      "6号梯初始化上行接触器" : Bool;
      "1号梯初始化下行接触器" : Bool;
      "2号梯初始化下行接触器" : Bool;
      "3号梯初始化下行接触器" : Bool;
      "4号梯初始化下行接触器" : Bool;
      "5号梯初始化下行接触器" : Bool;
      "6号梯初始化下行接触器" : Bool;
      "1号梯停梯截断(置0完成关门）" : Bool;
      "2号梯停梯截断(置0完成关门）" : Bool;
      "3号梯停梯截断(置0完成关门）" : Bool;
      "4号梯停梯截断(置0完成关门）" : Bool;
      "5号梯停梯截断(置0完成关门）" : Bool;
      "6号梯停梯截断(置0完成关门）" : Bool;
      "1号梯停梯截断(置0完成开门）" : Bool;
      "2号梯停梯截断(置0完成开门）" : Bool;
      "3号梯停梯截断(置0完成开门）" : Bool;
      "4号梯停梯截断(置0完成开门）" : Bool;
      "5号梯停梯截断(置0完成开门）" : Bool;
      "6号梯停梯截断(置0完成开门）" : Bool;
      "1号梯置0为完成开门" : Bool;
      "2号梯置0为完成开门" : Bool;
      "3号梯置0为完成开门" : Bool;
      "4号梯置0为完成开门" : Bool;
      "5号梯置0为完成开门" : Bool;
      "6号梯置0为完成开门" : Bool;
      "1号梯置0为完成关门" : Bool;
      "2号梯置0为完成关门" : Bool;
      "3号梯置0为完成关门" : Bool;
      "4号梯置0为完成关门" : Bool;
      "5号梯置0为完成关门" : Bool;
      "6号梯置0为完成关门" : Bool;
      "1号梯转换" : Real;
      "2号梯转换" : Real;
      "3号梯转换" : Real;
      "4号梯转换" : Real;
      "5号梯转换" : Real;
      "6号梯转换" : Real;
      "1号梯载重限额" : Int := 1050;
      "2号梯载重限额" : Int := 1350;
      "3号梯载重限额" : Int := 1350;
      "4号梯载重限额" : Int := 1350;
      "5号梯载重限额" : Int := 1800;
      "6号梯载重限额" : Int := 2000;
      "1号梯准备就绪" : Bool;
      "2号梯准备就绪" : Bool;
      "3号梯准备就绪" : Bool;
      "4号梯准备就绪" : Bool;
      "5号梯准备就绪" : Bool;
      "6号梯准备就绪" : Bool;
      "1号梯将要停梯" : Bool;
      "2号梯将要停梯" : Bool;
      "3号梯将要停梯" : Bool;
      "4号梯将要停梯" : Bool;
      "5号梯将要停梯" : Bool;
      "6号梯将要停梯" : Bool;
      "1号梯初始化将要停梯" : Bool;
      "2号梯初始化将要停梯" : Bool;
      "3号梯初始化将要停梯" : Bool;
      "4号梯初始化将要停梯" : Bool;
      "5号梯初始化将要停梯" : Bool;
      "6号梯初始化将要停梯" : Bool;
      初始化1级制动 : Bool;
      初始化2级制动 : Bool;
      初始化3级制动 : Bool;
      卡顿上行1 : Bool;
      卡顿上行2 : Bool;
      卡顿上行3 : Bool;
      卡顿上行4 : Bool;
      卡顿上行5 : Bool;
      卡顿上行6 : Bool;
      卡顿下行1 : Bool;
      卡顿下行2 : Bool;
      卡顿下行3 : Bool;
      卡顿下行4 : Bool;
      卡顿下行5 : Bool;
      卡顿下行6 : Bool;
      卡顿制速1 : Bool;
      卡顿制速2 : Bool;
      卡顿制速3 : Bool;
      卡顿制速4 : Bool;
      卡顿制速5 : Bool;
      卡顿制速6 : Bool;
      到达初始化楼层1号梯 : Bool;
      到达初始化楼层2号梯 : Bool;
      到达初始化楼层3号梯 : Bool;
      到达初始化楼层4号梯 : Bool;
      到达初始化楼层5号梯 : Bool;
      到达初始化楼层6号梯 : Bool;
      死机1 : Bool;
      死机2 : Bool;
      死机3 : Bool;
      死机4 : Bool;
      死机5 : Bool;
      死机6 : Bool;
      截下 : Bool;
      截上 : Bool;
      疑似满载1 : Int;
      疑似满载2 : Int;
      疑似满载3 : Int;
      疑似满载4 : Int;
      疑似满载5 : Int;
      "1号梯初始化方向位" : Int;
      "2号梯初始化方向位" : Int;
      "3号梯初始化方向位" : Int;
      "4号梯初始化方向位" : Int;
      "5号梯初始化方向位" : Int;
      "6号梯初始化方向位" : Int;
      "1号梯初始化方向位选择" : Bool;
      "2号梯初始化方向位选择" : Bool;
      "3号梯初始化方向位选择" : Bool;
      "4号梯初始化方向位选择" : Bool;
      "5号梯初始化方向位选择" : Bool;
      "6号梯初始化方向位选择" : Bool;
      疑似满载6 : Int;
      "1号梯正确楼层数" : Int;
      "2号梯正确楼层数" : Int;
      "3号梯正确楼层数" : Int;
      "4号梯正确楼层数" : Int;
      "5号梯正确楼层数" : Int;
      "6号梯正确楼层数" : Int;
      程序运行时长秒 : Int;
      程序运行时长分钟 : Int;
      程序运行时长小时 : Int;
      程序运行时长 : Time_Of_Day;
      程序运行时长初始量 : Time_Of_Day;
      时间累加器最长时长 : Time := T#99999999ms;
      小时复位 : Bool;
      分钟复位 : Bool;
      秒复位 : Bool;
   END_VAR
BEGIN
END_DATA_BLOCK

// folder: 1号梯

DATA_BLOCK "1号梯初始化"   // DB1
{ S7_Optimized_Access := 'TRUE' }
VERSION : 0.1
// stored: InstanceOfName 初始化
"初始化"
BEGIN
END_DATA_BLOCK

DATA_BLOCK "1号梯距离调度"   // DB4
{ S7_Optimized_Access := 'TRUE' }
VERSION : 0.1
// stored: InstanceOfName 距离调度
"距离调度"
BEGIN
END_DATA_BLOCK

DATA_BLOCK "1号梯指示灯"   // DB6
{ S7_Optimized_Access := 'TRUE' }
VERSION : 0.1
// stored: InstanceOfName 照明，风扇，数码管
"照明，风扇，数码管"
BEGIN
END_DATA_BLOCK

DATA_BLOCK "1号梯停层次数"   // DB7
{ S7_Optimized_Access := 'TRUE' }
VERSION : 0.1
// stored: InstanceOfName 停层次数判断
"停层次数判断"
BEGIN
END_DATA_BLOCK

DATA_BLOCK "1号梯高低速转换"   // DB9
{ S7_Optimized_Access := 'TRUE' }
VERSION : 0.1
// stored: InstanceOfName 高低速转换
"高低速转换"
BEGIN
END_DATA_BLOCK

DATA_BLOCK "1号梯上下行与制动"   // DB16
{ S7_Optimized_Access := 'TRUE' }
VERSION : 0.1
// stored: InstanceOfName 上下行和制动
"上下行和制动"
BEGIN
END_DATA_BLOCK

DATA_BLOCK "1号梯优先级"   // DB18
{ S7_Optimized_Access := 'TRUE' }
VERSION : 0.1
// stored: InstanceOfName 优先级响应开关门
"优先级响应开关门"
BEGIN
END_DATA_BLOCK

DATA_BLOCK "1号梯楼层计算"   // DB20
{ S7_Optimized_Access := 'TRUE' }
VERSION : 0.1
// stored: InstanceOfName 楼层计算
"楼层计算"
BEGIN
END_DATA_BLOCK

DATA_BLOCK "1号梯有无目标判断"   // DB24
{ S7_Optimized_Access := 'TRUE' }
VERSION : 0.1
// stored: InstanceOfName 目标判断
"目标判断"
BEGIN
END_DATA_BLOCK

// folder: 2号梯

DATA_BLOCK "2号梯初始化"   // DB14
{ S7_Optimized_Access := 'TRUE' }
VERSION : 0.1
// stored: InstanceOfName 初始化
"初始化"
BEGIN
END_DATA_BLOCK

DATA_BLOCK "2号梯高低速转换"   // DB15
{ S7_Optimized_Access := 'TRUE' }
VERSION : 0.1
// stored: InstanceOfName 高低速转换
"高低速转换"
BEGIN
END_DATA_BLOCK

DATA_BLOCK "2号梯上下行与制动"   // DB44
{ S7_Optimized_Access := 'TRUE' }
VERSION : 0.1
// stored: InstanceOfName 上下行和制动
"上下行和制动"
BEGIN
END_DATA_BLOCK

DATA_BLOCK "2号梯距离调度"   // DB49
{ S7_Optimized_Access := 'TRUE' }
VERSION : 0.1
// stored: InstanceOfName 距离调度
"距离调度"
BEGIN
END_DATA_BLOCK

DATA_BLOCK "2号梯停层次数"   // DB54
{ S7_Optimized_Access := 'TRUE' }
VERSION : 0.1
// stored: InstanceOfName 停层次数判断
"停层次数判断"
BEGIN
END_DATA_BLOCK

DATA_BLOCK "2号梯楼层计算"   // DB59
{ S7_Optimized_Access := 'TRUE' }
VERSION : 0.1
// stored: InstanceOfName 楼层计算
"楼层计算"
BEGIN
END_DATA_BLOCK

DATA_BLOCK "2号梯优先级"   // DB64
{ S7_Optimized_Access := 'TRUE' }
VERSION : 0.1
// stored: InstanceOfName 优先级响应开关门
"优先级响应开关门"
BEGIN
END_DATA_BLOCK

DATA_BLOCK "2号梯指示灯"   // DB69
{ S7_Optimized_Access := 'TRUE' }
VERSION : 0.1
// stored: InstanceOfName 照明，风扇，数码管
"照明，风扇，数码管"
BEGIN
END_DATA_BLOCK

DATA_BLOCK "2号梯有无目标判断"   // DB74
{ S7_Optimized_Access := 'TRUE' }
VERSION : 0.1
// stored: InstanceOfName 目标判断
"目标判断"
BEGIN
END_DATA_BLOCK

// folder: 3号梯

DATA_BLOCK "3号梯初始化"   // DB17
{ S7_Optimized_Access := 'TRUE' }
VERSION : 0.1
// stored: InstanceOfName 初始化
"初始化"
BEGIN
END_DATA_BLOCK

DATA_BLOCK "3号梯高低速转换"   // DB40
{ S7_Optimized_Access := 'TRUE' }
VERSION : 0.1
// stored: InstanceOfName 高低速转换
"高低速转换"
BEGIN
END_DATA_BLOCK

DATA_BLOCK "3号梯上下行与制动"   // DB45
{ S7_Optimized_Access := 'TRUE' }
VERSION : 0.1
// stored: InstanceOfName 上下行和制动
"上下行和制动"
BEGIN
END_DATA_BLOCK

DATA_BLOCK "3号梯距离调度"   // DB50
{ S7_Optimized_Access := 'TRUE' }
VERSION : 0.1
// stored: InstanceOfName 距离调度
"距离调度"
BEGIN
END_DATA_BLOCK

DATA_BLOCK "3号梯停层次数"   // DB55
{ S7_Optimized_Access := 'TRUE' }
VERSION : 0.1
// stored: InstanceOfName 停层次数判断
"停层次数判断"
BEGIN
END_DATA_BLOCK

DATA_BLOCK "3号梯楼层计算"   // DB60
{ S7_Optimized_Access := 'TRUE' }
VERSION : 0.1
// stored: InstanceOfName 楼层计算
"楼层计算"
BEGIN
END_DATA_BLOCK

DATA_BLOCK "3号梯优先级"   // DB65
{ S7_Optimized_Access := 'TRUE' }
VERSION : 0.1
// stored: InstanceOfName 优先级响应开关门
"优先级响应开关门"
BEGIN
END_DATA_BLOCK

DATA_BLOCK "3号梯指示灯"   // DB70
{ S7_Optimized_Access := 'TRUE' }
VERSION : 0.1
// stored: InstanceOfName 照明，风扇，数码管
"照明，风扇，数码管"
BEGIN
END_DATA_BLOCK

DATA_BLOCK "3号梯有无目标判断"   // DB75
{ S7_Optimized_Access := 'TRUE' }
VERSION : 0.1
// stored: InstanceOfName 目标判断
"目标判断"
BEGIN
END_DATA_BLOCK

// folder: 4号梯

DATA_BLOCK "4号梯初始化"   // DB19
{ S7_Optimized_Access := 'TRUE' }
VERSION : 0.1
// stored: InstanceOfName 初始化
"初始化"
BEGIN
END_DATA_BLOCK

DATA_BLOCK "4号梯高低速转换"   // DB41
{ S7_Optimized_Access := 'TRUE' }
VERSION : 0.1
// stored: InstanceOfName 高低速转换
"高低速转换"
BEGIN
END_DATA_BLOCK

DATA_BLOCK "4号梯上下行与制动"   // DB46
{ S7_Optimized_Access := 'TRUE' }
VERSION : 0.1
// stored: InstanceOfName 上下行和制动
"上下行和制动"
BEGIN
END_DATA_BLOCK

DATA_BLOCK "4号梯距离调度"   // DB51
{ S7_Optimized_Access := 'TRUE' }
VERSION : 0.1
// stored: InstanceOfName 距离调度
"距离调度"
BEGIN
END_DATA_BLOCK

DATA_BLOCK "4号梯停层次数"   // DB56
{ S7_Optimized_Access := 'TRUE' }
VERSION : 0.1
// stored: InstanceOfName 停层次数判断
"停层次数判断"
BEGIN
END_DATA_BLOCK

DATA_BLOCK "4号梯楼层计算"   // DB61
{ S7_Optimized_Access := 'TRUE' }
VERSION : 0.1
// stored: InstanceOfName 楼层计算
"楼层计算"
BEGIN
END_DATA_BLOCK

DATA_BLOCK "4号梯优先级"   // DB66
{ S7_Optimized_Access := 'TRUE' }
VERSION : 0.1
// stored: InstanceOfName 优先级响应开关门
"优先级响应开关门"
BEGIN
END_DATA_BLOCK

DATA_BLOCK "4号梯指示灯"   // DB71
{ S7_Optimized_Access := 'TRUE' }
VERSION : 0.1
// stored: InstanceOfName 照明，风扇，数码管
"照明，风扇，数码管"
BEGIN
END_DATA_BLOCK

DATA_BLOCK "4号梯有无目标判断"   // DB76
{ S7_Optimized_Access := 'TRUE' }
VERSION : 0.1
// stored: InstanceOfName 目标判断
"目标判断"
BEGIN
END_DATA_BLOCK

// folder: 5号梯

DATA_BLOCK "5号梯初始化"   // DB22
{ S7_Optimized_Access := 'TRUE' }
VERSION : 0.1
// stored: InstanceOfName 初始化
"初始化"
BEGIN
END_DATA_BLOCK

DATA_BLOCK "5号梯高低速转换"   // DB42
{ S7_Optimized_Access := 'TRUE' }
VERSION : 0.1
// stored: InstanceOfName 初始化低速模式
"初始化低速模式"
BEGIN
END_DATA_BLOCK

DATA_BLOCK "5号梯上下行与制动"   // DB47
{ S7_Optimized_Access := 'TRUE' }
VERSION : 0.1
// stored: InstanceOfName 上下行和制动
"上下行和制动"
BEGIN
END_DATA_BLOCK

DATA_BLOCK "5号梯距离调度"   // DB52
{ S7_Optimized_Access := 'TRUE' }
VERSION : 0.1
// stored: InstanceOfName 距离调度
"距离调度"
BEGIN
END_DATA_BLOCK

DATA_BLOCK "5号梯停层次数"   // DB57
{ S7_Optimized_Access := 'TRUE' }
VERSION : 0.1
// stored: InstanceOfName 停层次数判断
"停层次数判断"
BEGIN
END_DATA_BLOCK

DATA_BLOCK "5号梯楼层计算"   // DB62
{ S7_Optimized_Access := 'TRUE' }
VERSION : 0.1
// stored: InstanceOfName 楼层计算
"楼层计算"
BEGIN
END_DATA_BLOCK

DATA_BLOCK "5号梯优先级"   // DB67
{ S7_Optimized_Access := 'TRUE' }
VERSION : 0.1
// stored: InstanceOfName 优先级响应开关门
"优先级响应开关门"
BEGIN
END_DATA_BLOCK

DATA_BLOCK "5号梯指示灯"   // DB72
{ S7_Optimized_Access := 'TRUE' }
VERSION : 0.1
// stored: InstanceOfName 照明，风扇，数码管
"照明，风扇，数码管"
BEGIN
END_DATA_BLOCK

DATA_BLOCK "5号梯有无目标判断"   // DB77
{ S7_Optimized_Access := 'TRUE' }
VERSION : 0.1
// stored: InstanceOfName 目标判断
"目标判断"
BEGIN
END_DATA_BLOCK

DATA_BLOCK "5号梯高低速切换"   // DB80
{ S7_Optimized_Access := 'TRUE' }
VERSION : 0.1
// stored: InstanceOfName 高低速转换
"高低速转换"
BEGIN
END_DATA_BLOCK

// folder: 6号梯

DATA_BLOCK "6号梯初始化"   // DB23
{ S7_Optimized_Access := 'TRUE' }
VERSION : 0.1
// stored: InstanceOfName 初始化
"初始化"
BEGIN
END_DATA_BLOCK

DATA_BLOCK "6号梯高低速转换"   // DB43
{ S7_Optimized_Access := 'TRUE' }
VERSION : 0.1
// stored: InstanceOfName 初始化低速模式
"初始化低速模式"
BEGIN
END_DATA_BLOCK

DATA_BLOCK "6号梯上下行与制动"   // DB48
{ S7_Optimized_Access := 'TRUE' }
VERSION : 0.1
// stored: InstanceOfName 上下行和制动
"上下行和制动"
BEGIN
END_DATA_BLOCK

DATA_BLOCK "6号梯距离调度"   // DB53
{ S7_Optimized_Access := 'TRUE' }
VERSION : 0.1
// stored: InstanceOfName 距离调度
"距离调度"
BEGIN
END_DATA_BLOCK

DATA_BLOCK "6号梯停层次数"   // DB58
{ S7_Optimized_Access := 'TRUE' }
VERSION : 0.1
// stored: InstanceOfName 停层次数判断
"停层次数判断"
BEGIN
END_DATA_BLOCK

DATA_BLOCK "6号梯楼层计算"   // DB63
{ S7_Optimized_Access := 'TRUE' }
VERSION : 0.1
// stored: InstanceOfName 楼层计算
"楼层计算"
BEGIN
END_DATA_BLOCK

DATA_BLOCK "6号梯优先级"   // DB68
{ S7_Optimized_Access := 'TRUE' }
VERSION : 0.1
// stored: InstanceOfName 优先级响应开关门
"优先级响应开关门"
BEGIN
END_DATA_BLOCK

DATA_BLOCK "6号梯指示灯"   // DB73
{ S7_Optimized_Access := 'TRUE' }
VERSION : 0.1
// stored: InstanceOfName 照明，风扇，数码管
"照明，风扇，数码管"
BEGIN
END_DATA_BLOCK

DATA_BLOCK "6号梯有无目标判断"   // DB78
{ S7_Optimized_Access := 'TRUE' }
VERSION : 0.1
// stored: InstanceOfName 目标判断
"目标判断"
BEGIN
END_DATA_BLOCK

DATA_BLOCK "6号梯高低速切换"   // DB82
{ S7_Optimized_Access := 'TRUE' }
VERSION : 0.1
// stored: InstanceOfName 高低速转换
"高低速转换"
BEGIN
END_DATA_BLOCK

// folder: System blocks/Program resources

DATA_BLOCK "1号梯初始化置位延时"   // DB21
{ S7_Optimized_Access := 'TRUE' }
AUTHOR : Simatic
FAMILY : IEC
NAME : IEC_TMR
VERSION : 1.0
// stored: InstanceOfName IEC_TIMER
"IEC_TIMER"
BEGIN
END_DATA_BLOCK

DATA_BLOCK "2号梯初始化置位延时"   // DB79
{ S7_Optimized_Access := 'TRUE' }
AUTHOR : Simatic
FAMILY : IEC
NAME : IEC_TMR
VERSION : 1.0
// stored: InstanceOfName IEC_TIMER
"IEC_TIMER"
BEGIN
END_DATA_BLOCK

DATA_BLOCK "3号梯初始化置位延时"   // DB81
{ S7_Optimized_Access := 'TRUE' }
AUTHOR : Simatic
FAMILY : IEC
NAME : IEC_TMR
VERSION : 1.0
// stored: InstanceOfName IEC_TIMER
"IEC_TIMER"
BEGIN
END_DATA_BLOCK

DATA_BLOCK "4号梯初始化置位延时"   // DB83
{ S7_Optimized_Access := 'TRUE' }
AUTHOR : Simatic
FAMILY : IEC
NAME : IEC_TMR
VERSION : 1.0
// stored: InstanceOfName IEC_TIMER
"IEC_TIMER"
BEGIN
END_DATA_BLOCK

DATA_BLOCK "接通延时"   // DB84
{ S7_Optimized_Access := 'TRUE' }
AUTHOR : Simatic
FAMILY : IEC
NAME : IEC_TMR
VERSION : 1.0
// stored: InstanceOfName IEC_TIMER
"IEC_TIMER"
BEGIN
END_DATA_BLOCK

DATA_BLOCK "5号梯初始化置位延时"   // DB85
{ S7_Optimized_Access := 'TRUE' }
AUTHOR : Simatic
FAMILY : IEC
NAME : IEC_TMR
VERSION : 1.0
// stored: InstanceOfName IEC_TIMER
"IEC_TIMER"
BEGIN
END_DATA_BLOCK

DATA_BLOCK "6号梯初始化置位延时"   // DB87
{ S7_Optimized_Access := 'TRUE' }
AUTHOR : Simatic
FAMILY : IEC
NAME : IEC_TMR
VERSION : 1.0
// stored: InstanceOfName IEC_TIMER
"IEC_TIMER"
BEGIN
END_DATA_BLOCK

DATA_BLOCK "每秒脉冲生成器"   // DB91
{ S7_Optimized_Access := 'TRUE' }
AUTHOR : Simatic
FAMILY : IEC
NAME : IEC_TMR
VERSION : 1.0
// stored: InstanceOfName IEC_TIMER
"IEC_TIMER"
BEGIN
END_DATA_BLOCK

DATA_BLOCK "脉冲计数小时"   // DB93
{ S7_Optimized_Access := 'TRUE' }
AUTHOR : Simatic
FAMILY : IEC
NAME : CNTR
VERSION : 1.0
// stored: InstanceOfName IEC_COUNTER
"IEC_COUNTER"
BEGIN
END_DATA_BLOCK

DATA_BLOCK "脉冲计数秒"   // DB94
{ S7_Optimized_Access := 'TRUE' }
AUTHOR : Simatic
FAMILY : IEC
NAME : CNTR
VERSION : 1.0
// stored: InstanceOfName IEC_COUNTER
"IEC_COUNTER"
BEGIN
END_DATA_BLOCK

DATA_BLOCK "脉冲计数分钟"   // DB95
{ S7_Optimized_Access := 'TRUE' }
AUTHOR : Simatic
FAMILY : IEC
NAME : CNTR
VERSION : 1.0
// stored: InstanceOfName IEC_COUNTER
"IEC_COUNTER"
BEGIN
END_DATA_BLOCK

// folder: 距离比较

DATA_BLOCK "1层上呼距离比较"   // DB5
{ S7_Optimized_Access := 'TRUE' }
VERSION : 0.1
// stored: InstanceOfName 距离比较
"距离比较"
BEGIN
END_DATA_BLOCK

DATA_BLOCK "2层上呼距离比较"   // DB8
{ S7_Optimized_Access := 'TRUE' }
VERSION : 0.1
// stored: InstanceOfName 距离比较
"距离比较"
BEGIN
END_DATA_BLOCK

DATA_BLOCK "2层下呼距离比较"   // DB12
{ S7_Optimized_Access := 'TRUE' }
VERSION : 0.1
// stored: InstanceOfName 距离比较
"距离比较"
BEGIN
END_DATA_BLOCK

DATA_BLOCK "3层上呼距离比较"   // DB25
{ S7_Optimized_Access := 'TRUE' }
VERSION : 0.1
// stored: InstanceOfName 距离比较
"距离比较"
BEGIN
END_DATA_BLOCK

DATA_BLOCK "3层下呼距离比较"   // DB26
{ S7_Optimized_Access := 'TRUE' }
VERSION : 0.1
// stored: InstanceOfName 距离比较
"距离比较"
BEGIN
END_DATA_BLOCK

DATA_BLOCK "4层上呼距离比较"   // DB27
{ S7_Optimized_Access := 'TRUE' }
VERSION : 0.1
// stored: InstanceOfName 距离比较
"距离比较"
BEGIN
END_DATA_BLOCK

DATA_BLOCK "4层下呼距离比较"   // DB28
{ S7_Optimized_Access := 'TRUE' }
VERSION : 0.1
// stored: InstanceOfName 距离比较
"距离比较"
BEGIN
END_DATA_BLOCK

DATA_BLOCK "5层上呼距离比较"   // DB29
{ S7_Optimized_Access := 'TRUE' }
VERSION : 0.1
// stored: InstanceOfName 距离比较
"距离比较"
BEGIN
END_DATA_BLOCK

DATA_BLOCK "5层下呼距离比较"   // DB30
{ S7_Optimized_Access := 'TRUE' }
VERSION : 0.1
// stored: InstanceOfName 距离比较
"距离比较"
BEGIN
END_DATA_BLOCK

DATA_BLOCK "6层上呼距离比较"   // DB31
{ S7_Optimized_Access := 'TRUE' }
VERSION : 0.1
// stored: InstanceOfName 距离比较
"距离比较"
BEGIN
END_DATA_BLOCK

DATA_BLOCK "6层下呼距离比较"   // DB32
{ S7_Optimized_Access := 'TRUE' }
VERSION : 0.1
// stored: InstanceOfName 距离比较
"距离比较"
BEGIN
END_DATA_BLOCK

DATA_BLOCK "7层上呼距离比较"   // DB33
{ S7_Optimized_Access := 'TRUE' }
VERSION : 0.1
// stored: InstanceOfName 距离比较
"距离比较"
BEGIN
END_DATA_BLOCK

DATA_BLOCK "7层下呼距离比较"   // DB34
{ S7_Optimized_Access := 'TRUE' }
VERSION : 0.1
// stored: InstanceOfName 距离比较
"距离比较"
BEGIN
END_DATA_BLOCK

DATA_BLOCK "8层上呼距离比较"   // DB35
{ S7_Optimized_Access := 'TRUE' }
VERSION : 0.1
// stored: InstanceOfName 距离比较
"距离比较"
BEGIN
END_DATA_BLOCK

DATA_BLOCK "8层下行距离比较"   // DB36
{ S7_Optimized_Access := 'TRUE' }
VERSION : 0.1
// stored: InstanceOfName 距离比较
"距离比较"
BEGIN
END_DATA_BLOCK

DATA_BLOCK "9层上呼距离比较"   // DB37
{ S7_Optimized_Access := 'TRUE' }
VERSION : 0.1
// stored: InstanceOfName 距离比较
"距离比较"
BEGIN
END_DATA_BLOCK

DATA_BLOCK "9层下呼距离比较"   // DB38
{ S7_Optimized_Access := 'TRUE' }
VERSION : 0.1
// stored: InstanceOfName 距离比较
"距离比较"
BEGIN
END_DATA_BLOCK

DATA_BLOCK "10层下行距离比较"   // DB39
{ S7_Optimized_Access := 'TRUE' }
VERSION : 0.1
// stored: InstanceOfName 距离比较
"距离比较"
BEGIN
END_DATA_BLOCK

// folder: (top level)

FUNCTION_BLOCK "距离比较"   // FB1, LAD
{ S7_Optimized_Access := 'TRUE' }
VERSION : 0.1
   VAR_INPUT
      上下平层同时为1梯1 : Bool;
      上下平层同时为1梯2 : Bool;
      上下平层同时为1梯3 : Bool;
      上下平层同时为1梯4 : Bool;
      上下平层同时为1梯5 : Bool;
      上下平层同时为1梯6 : Bool;
      有外呼楼层内选1 : Bool;
      有外呼楼层内选2 : Bool;
      有外呼楼层内选3 : Bool;
      有外呼楼层内选4 : Bool;
      有外呼楼层内选5 : Bool;
      有外呼楼层内选6 : Bool;
      就近运动电梯1 : Bool;
      就近运动电梯2 : Bool;
      就近运动电梯3 : Bool;
      就近运动电梯4 : Bool;
      就近运动电梯5 : Bool;
      就近运动电梯6 : Bool;
      呼灯 : Bool;
      调度距离1 : Int;
      调度距离2 : Int;
      调度距离3 : Int;
      调度距离4 : Int;
      调度距离5 : Int;
      调度距离6 : Int;
   END_VAR
   VAR_OUTPUT
      最小调度距离 : Int;
      分配给1 : Bool;
      分配给2 : Bool;
      分配给3 : Bool;
      分配给4 : Bool;
      分配给5 : Bool;
      分配给6 : Bool;
   END_VAR
   VAR
      追击1 : Bool;
      追击2 : Bool;
      追击3 : Bool;
      追击4 : Bool;
      追击5 : Bool;
      追击6 : Bool;
      中间分配1 : Bool;
      中间分配2 : Bool;
      中间分配3 : Bool;
      中间分配4 : Bool;
      中间分配5 : Bool;
      中间分配6 : Bool;
      内外呼重合1 : Bool;
      内外呼重合2 : Bool;
      内外呼重合3 : Bool;
      内外呼重合4 : Bool;
      内外呼重合5 : Bool;
      内外呼重合6 : Bool;
      与最小调度距离差值1 : Int;
      与最小调度距离差值2 : Int;
      与最小调度距离差值3 : Int;
      与最小调度距离差值4 : Int;
      与最小调度距离差值5 : Int;
      与最小调度距离差值6 : Int;
      IEC_Timer_0_Instance : TON_TIME;
      IEC_Timer_0_Instance_1 : TOF_TIME;
      "IEC_Ti me_0_Instance_3" : TOF_TIME;
      IEC_Timer_0_Instance_2 : TON_TIME;
      "IEC_Timer_0_Instance 5" : TOF_TIME;
      IEC_Timer_0_Instance_4 : TON_TIME;
      "IEC_Timer_0_Instance 7" : TOF_TIME;
      IEC_Timer_0_Instance_6 : TON_TIME;
      IEC_Timer_0_Instance_9 : TON_TIME;
      IEC_Timer_0_Instance11 : TON_TIME;
      "IEC_Timer_0_Instance 8" : TOF_TIME;
      IEC_Timer_0_Instance10 : TOF_TIME;
      IEC_Timer_0_Instance_3 : TOF_TIME;
      IEC_Timer_0_Instance_44 : TOF_TIME;
      IEC_Timer_0_Instance_45 : TOF_TIME;
      IEC_Timer_0_Instance_46 : TOF_TIME;
      IEC_Timer_0_Instance_47 : TOF_TIME;
   END_VAR
BEGIN

REGION Network 1: 比较计算
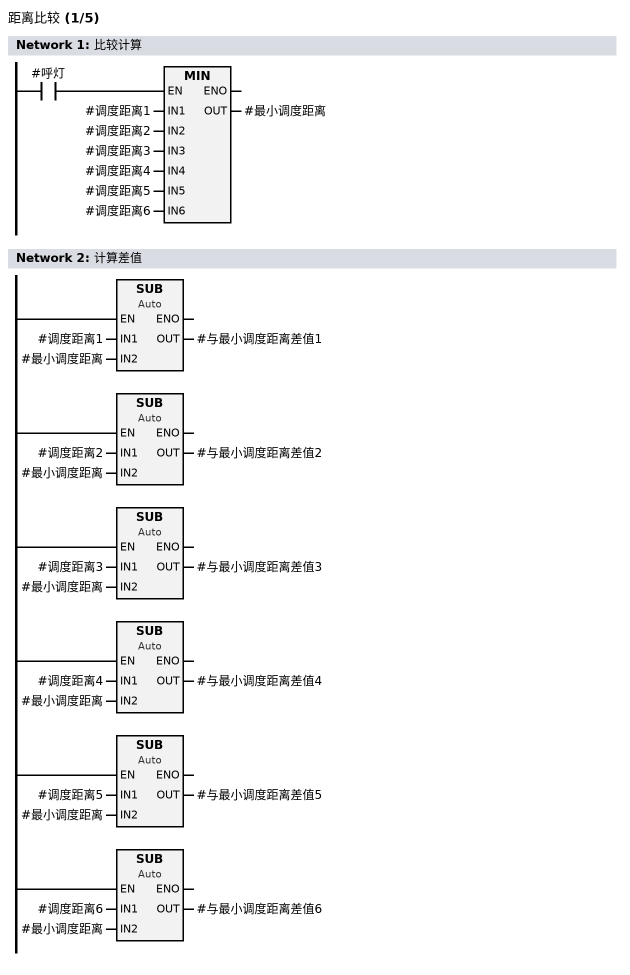
   IF #呼灯 THEN
       #最小调度距离 := MIN(IN1 := #调度距离1, IN2 := #调度距离2, IN3 := #调度距离3, IN4 := #调度距离4, IN5 := #调度距离5, IN6 := #调度距离6);
   END_IF;
END_REGION

REGION Network 2: 计算差值
   RUNG wire#powerrail
      Sub(in1 := #调度距离1, in2 := #最小调度距离, out => #与最小调度距离差值1)
   END_RUNG
   RUNG wire#powerrail
      Sub(in1 := #调度距离2, in2 := #最小调度距离, out => #与最小调度距离差值2)
   END_RUNG
   RUNG wire#powerrail
      Sub(in1 := #调度距离3, in2 := #最小调度距离, out => #与最小调度距离差值3)
   END_RUNG
   RUNG wire#powerrail
      Sub(in1 := #调度距离4, in2 := #最小调度距离, out => #与最小调度距离差值4)
   END_RUNG
   RUNG wire#powerrail
      Sub(in1 := #调度距离5, in2 := #最小调度距离, out => #与最小调度距离差值5)
   END_RUNG
   RUNG wire#powerrail
      Sub(in1 := #调度距离6, in2 := #最小调度距离, out => #与最小调度距离差值6)
   END_RUNG
   // the same network as SCL:
   #与最小调度距离差值1 := #调度距离1 - #最小调度距离;
   #与最小调度距离差值2 := #调度距离2 - #最小调度距离;
   #与最小调度距离差值3 := #调度距离3 - #最小调度距离;
   #与最小调度距离差值4 := #调度距离4 - #最小调度距离;
   #与最小调度距离差值5 := #调度距离5 - #最小调度距离;
   #与最小调度距离差值6 := #调度距离6 - #最小调度距离;
END_REGION

REGION Network 3: 追击
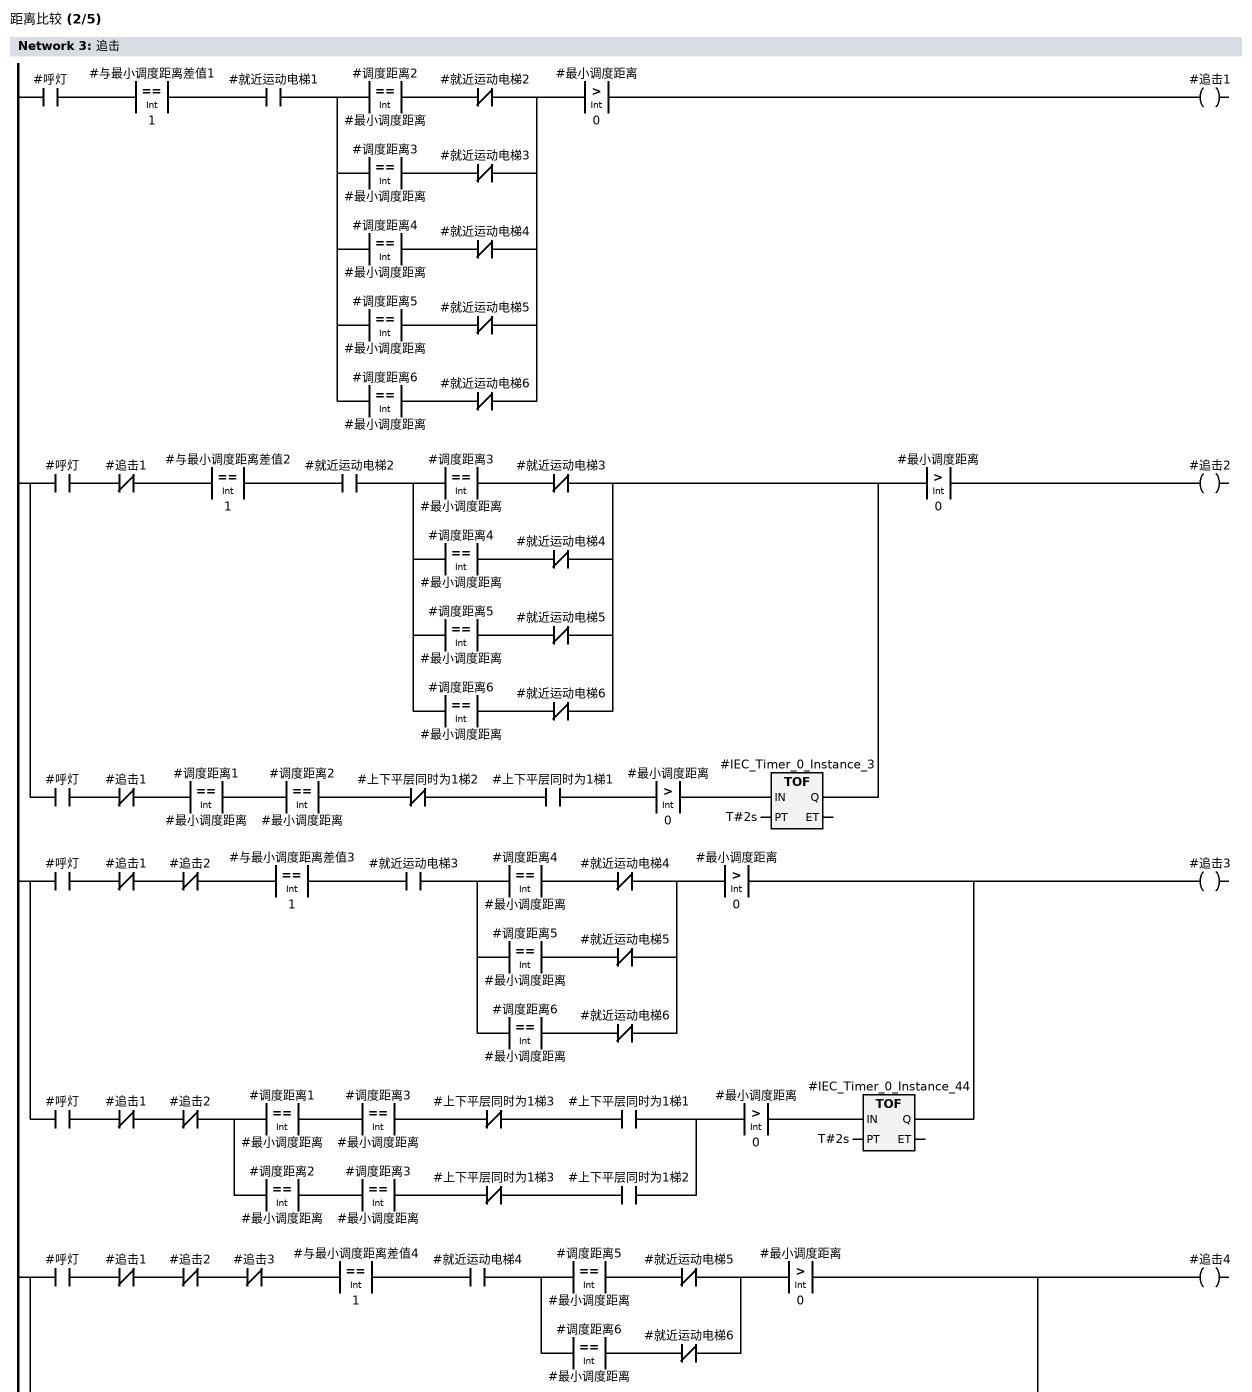
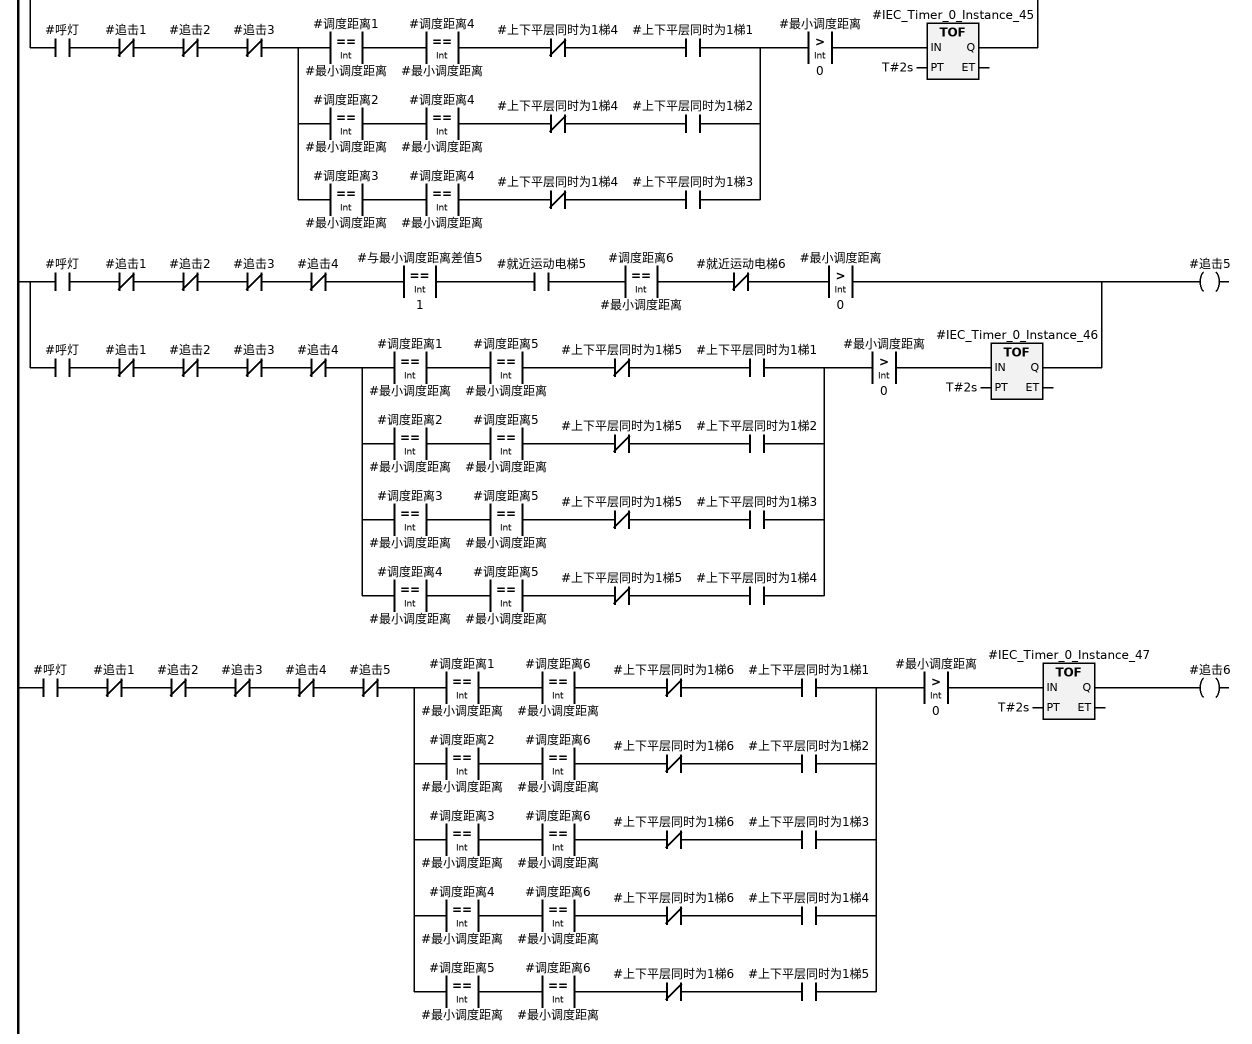
   #追击1 := #呼灯 AND (#与最小调度距离差值1 = 1) AND #就近运动电梯1 AND (((#调度距离2 = #最小调度距离) AND NOT #就近运动电梯2) OR ((#调度距离3 = #最小调度距离) AND NOT #就近运动电梯3) OR ((#调度距离4 = #最小调度距离) AND NOT #就近运动电梯4) OR ((#调度距离5 = #最小调度距离) AND NOT #就近运动电梯5) OR ((#调度距离6 = #最小调度距离) AND NOT #就近运动电梯6)) AND (#最小调度距离 > 0);
   #IEC_Timer_0_Instance_3(IN := #呼灯 AND NOT #追击1 AND (#调度距离1 = #最小调度距离) AND (#调度距离2 = #最小调度距离) AND NOT #上下平层同时为1梯2 AND #上下平层同时为1梯1 AND (#最小调度距离 > 0),   // TOF
                           PT := T#2s);
   #追击2 := ((#呼灯 AND NOT #追击1 AND (#与最小调度距离差值2 = 1) AND #就近运动电梯2 AND (((#调度距离3 = #最小调度距离) AND NOT #就近运动电梯3) OR ((#调度距离4 = #最小调度距离) AND NOT #就近运动电梯4) OR ((#调度距离5 = #最小调度距离) AND NOT #就近运动电梯5) OR ((#调度距离6 = #最小调度距离) AND NOT #就近运动电梯6))) OR #IEC_Timer_0_Instance_3.Q) AND (#最小调度距离 > 0);
   #IEC_Timer_0_Instance_44(IN := #呼灯 AND NOT #追击1 AND NOT #追击2 AND (((#调度距离1 = #最小调度距离) AND (#调度距离3 = #最小调度距离) AND NOT #上下平层同时为1梯3 AND #上下平层同时为1梯1) OR ((#调度距离2 = #最小调度距离) AND (#调度距离3 = #最小调度距离) AND NOT #上下平层同时为1梯3 AND #上下平层同时为1梯2)) AND (#最小调度距离 > 0),   // TOF
                           PT := T#2s);
   #追击3 := (#呼灯 AND NOT #追击1 AND NOT #追击2 AND (#与最小调度距离差值3 = 1) AND #就近运动电梯3 AND (((#调度距离4 = #最小调度距离) AND NOT #就近运动电梯4) OR ((#调度距离5 = #最小调度距离) AND NOT #就近运动电梯5) OR ((#调度距离6 = #最小调度距离) AND NOT #就近运动电梯6)) AND (#最小调度距离 > 0)) OR #IEC_Timer_0_Instance_44.Q;
   #IEC_Timer_0_Instance_45(IN := #呼灯 AND NOT #追击1 AND NOT #追击2 AND NOT #追击3 AND (((#调度距离1 = #最小调度距离) AND (#调度距离4 = #最小调度距离) AND NOT #上下平层同时为1梯4 AND #上下平层同时为1梯1) OR ((#调度距离2 = #最小调度距离) AND (#调度距离4 = #最小调度距离) AND NOT #上下平层同时为1梯4 AND #上下平层同时为1梯2) OR ((#调度距离3 = #最小调度距离) AND (#调度距离4 = #最小调度距离) AND NOT #上下平层同时为1梯4 AND #上下平层同时为1梯3)) AND (#最小调度距离 > 0),   // TOF
                           PT := T#2s);
   #追击4 := (#呼灯 AND NOT #追击1 AND NOT #追击2 AND NOT #追击3 AND (#与最小调度距离差值4 = 1) AND #就近运动电梯4 AND (((#调度距离5 = #最小调度距离) AND NOT #就近运动电梯5) OR ((#调度距离6 = #最小调度距离) AND NOT #就近运动电梯6)) AND (#最小调度距离 > 0)) OR #IEC_Timer_0_Instance_45.Q;
   #IEC_Timer_0_Instance_46(IN := #呼灯 AND NOT #追击1 AND NOT #追击2 AND NOT #追击3 AND NOT #追击4 AND (((#调度距离1 = #最小调度距离) AND (#调度距离5 = #最小调度距离) AND NOT #上下平层同时为1梯5 AND #上下平层同时为1梯1) OR ((#调度距离2 = #最小调度距离) AND (#调度距离5 = #最小调度距离) AND NOT #上下平层同时为1梯5 AND #上下平层同时为1梯2) OR ((#调度距离3 = #最小调度距离) AND (#调度距离5 = #最小调度距离) AND NOT #上下平层同时为1梯5 AND #上下平层同时为1梯3) OR ((#调度距离4 = #最小调度距离) AND (#调度距离5 = #最小调度距离) AND NOT #上下平层同时为1梯5 AND #上下平层同时为1梯4)) AND (#最小调度距离 > 0),   // TOF
                           PT := T#2s);
   #追击5 := (#呼灯 AND NOT #追击1 AND NOT #追击2 AND NOT #追击3 AND NOT #追击4 AND (#与最小调度距离差值5 = 1) AND #就近运动电梯5 AND (#调度距离6 = #最小调度距离) AND NOT #就近运动电梯6 AND (#最小调度距离 > 0)) OR #IEC_Timer_0_Instance_46.Q;
   #IEC_Timer_0_Instance_47(IN := #呼灯 AND NOT #追击1 AND NOT #追击2 AND NOT #追击3 AND NOT #追击4 AND NOT #追击5 AND (((#调度距离1 = #最小调度距离) AND (#调度距离6 = #最小调度距离) AND NOT #上下平层同时为1梯6 AND #上下平层同时为1梯1) OR ((#调度距离2 = #最小调度距离) AND (#调度距离6 = #最小调度距离) AND NOT #上下平层同时为1梯6 AND #上下平层同时为1梯2) OR ((#调度距离3 = #最小调度距离) AND (#调度距离6 = #最小调度距离) AND NOT #上下平层同时为1梯6 AND #上下平层同时为1梯3) OR ((#调度距离4 = #最小调度距离) AND (#调度距离6 = #最小调度距离) AND NOT #上下平层同时为1梯6 AND #上下平层同时为1梯4) OR ((#调度距离5 = #最小调度距离) AND (#调度距离6 = #最小调度距离) AND NOT #上下平层同时为1梯6 AND #上下平层同时为1梯5)) AND (#最小调度距离 > 0),   // TOF
                           PT := T#2s);
   #追击6 := #IEC_Timer_0_Instance_47.Q;
END_REGION

REGION Network 4: 判断内外呼是否重合
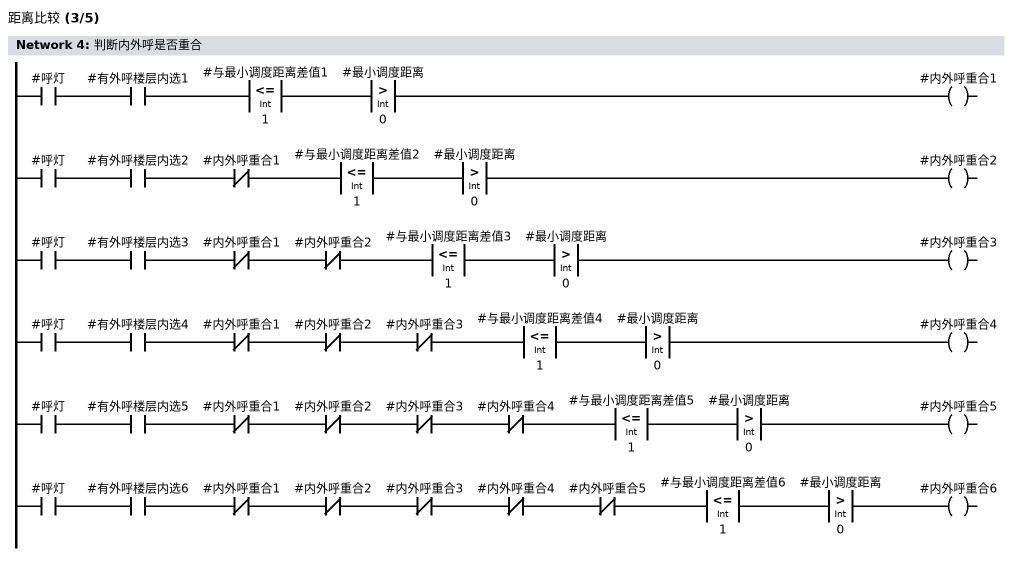
   RUNG wire#powerrail
      Contact( #呼灯 )
      Contact( #有外呼楼层内选1 )
      { S7_Templates := "SrcType := Int" } LE_Contact(in1 := #与最小调度距离差值1, in2 := 1)
      { S7_Templates := "SrcType := Int" } GT_Contact(in1 := #最小调度距离, in2 := 0)
      Coil( #内外呼重合1 )
   END_RUNG
   RUNG wire#powerrail
      Contact( #呼灯 )
      Contact( #有外呼楼层内选2 )
      I_Contact( #内外呼重合1 )
      { S7_Templates := "SrcType := Int" } LE_Contact(in1 := #与最小调度距离差值2, in2 := 1)
      { S7_Templates := "SrcType := Int" } GT_Contact(in1 := #最小调度距离, in2 := 0)
      Coil( #内外呼重合2 )
   END_RUNG
   RUNG wire#powerrail
      Contact( #呼灯 )
      Contact( #有外呼楼层内选3 )
      I_Contact( #内外呼重合1 )
      I_Contact( #内外呼重合2 )
      { S7_Templates := "SrcType := Int" } LE_Contact(in1 := #与最小调度距离差值3, in2 := 1)
      { S7_Templates := "SrcType := Int" } GT_Contact(in1 := #最小调度距离, in2 := 0)
      Coil( #内外呼重合3 )
   END_RUNG
   RUNG wire#powerrail
      Contact( #呼灯 )
      Contact( #有外呼楼层内选4 )
      I_Contact( #内外呼重合1 )
      I_Contact( #内外呼重合2 )
      I_Contact( #内外呼重合3 )
      { S7_Templates := "SrcType := Int" } LE_Contact(in1 := #与最小调度距离差值4, in2 := 1)
      { S7_Templates := "SrcType := Int" } GT_Contact(in1 := #最小调度距离, in2 := 0)
      Coil( #内外呼重合4 )
   END_RUNG
   RUNG wire#powerrail
      Contact( #呼灯 )
      Contact( #有外呼楼层内选5 )
      I_Contact( #内外呼重合1 )
      I_Contact( #内外呼重合2 )
      I_Contact( #内外呼重合3 )
      I_Contact( #内外呼重合4 )
      { S7_Templates := "SrcType := Int" } LE_Contact(in1 := #与最小调度距离差值5, in2 := 1)
      { S7_Templates := "SrcType := Int" } GT_Contact(in1 := #最小调度距离, in2 := 0)
      Coil( #内外呼重合5 )
   END_RUNG
   RUNG wire#powerrail
      Contact( #呼灯 )
      Contact( #有外呼楼层内选6 )
      I_Contact( #内外呼重合1 )
      I_Contact( #内外呼重合2 )
      I_Contact( #内外呼重合3 )
      I_Contact( #内外呼重合4 )
      I_Contact( #内外呼重合5 )
      { S7_Templates := "SrcType := Int" } LE_Contact(in1 := #与最小调度距离差值6, in2 := 1)
      { S7_Templates := "SrcType := Int" } GT_Contact(in1 := #最小调度距离, in2 := 0)
      Coil( #内外呼重合6 )
   END_RUNG
   // the same network as SCL:
   #内外呼重合1 := #呼灯 AND #有外呼楼层内选1 AND (#与最小调度距离差值1 <= 1) AND (#最小调度距离 > 0);
   #内外呼重合2 := #呼灯 AND #有外呼楼层内选2 AND NOT #内外呼重合1 AND (#与最小调度距离差值2 <= 1) AND (#最小调度距离 > 0);
   #内外呼重合3 := #呼灯 AND #有外呼楼层内选3 AND NOT #内外呼重合1 AND NOT #内外呼重合2 AND (#与最小调度距离差值3 <= 1) AND (#最小调度距离 > 0);
   #内外呼重合4 := #呼灯 AND #有外呼楼层内选4 AND NOT #内外呼重合1 AND NOT #内外呼重合2 AND NOT #内外呼重合3 AND (#与最小调度距离差值4 <= 1) AND (#最小调度距离 > 0);
   #内外呼重合5 := #呼灯 AND #有外呼楼层内选5 AND NOT #内外呼重合1 AND NOT #内外呼重合2 AND NOT #内外呼重合3 AND NOT #内外呼重合4 AND (#与最小调度距离差值5 <= 1) AND (#最小调度距离 > 0);
   #内外呼重合6 := #呼灯 AND #有外呼楼层内选6 AND NOT #内外呼重合1 AND NOT #内外呼重合2 AND NOT #内外呼重合3 AND NOT #内外呼重合4 AND NOT #内外呼重合5 AND (#与最小调度距离差值6 <= 1) AND (#最小调度距离 > 0);
END_REGION

REGION Network 5: 中间分配123456
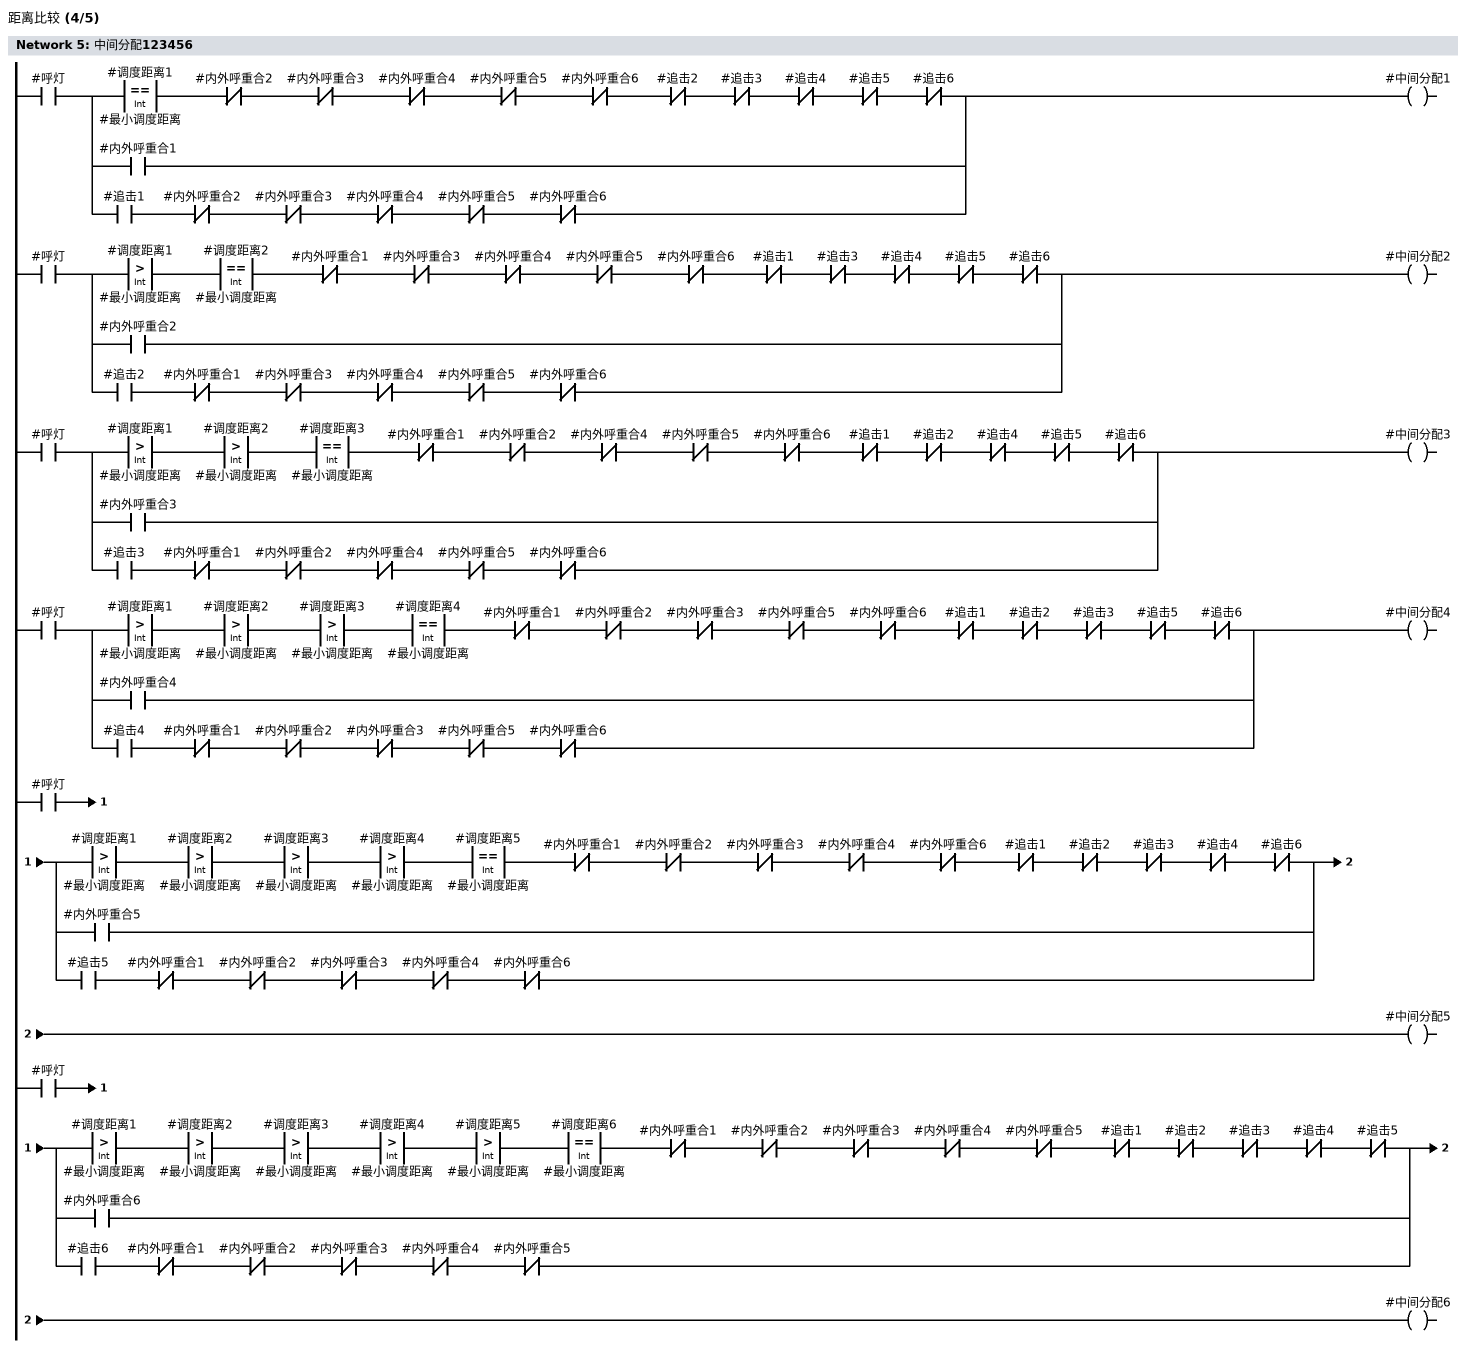
   RUNG wire#powerrail
      Contact( #呼灯 )
      wire#w1
      { S7_Templates := "SrcType := Int" } EQ_Contact(in1 := #调度距离1, in2 := #最小调度距离)
      I_Contact( #内外呼重合2 )
      I_Contact( #内外呼重合3 )
      I_Contact( #内外呼重合4 )
      I_Contact( #内外呼重合5 )
      I_Contact( #内外呼重合6 )
      I_Contact( #追击2 )
      I_Contact( #追击3 )
      I_Contact( #追击4 )
      I_Contact( #追击5 )
      I_Contact( #追击6 )
      wire#w2
      Coil( #中间分配1 )
   END_RUNG
   RUNG wire#w1
      Contact( #内外呼重合1 )
   END_RUNG wire#w2
   RUNG wire#w1
      Contact( #追击1 )
      I_Contact( #内外呼重合2 )
      I_Contact( #内外呼重合3 )
      I_Contact( #内外呼重合4 )
      I_Contact( #内外呼重合5 )
      I_Contact( #内外呼重合6 )
   END_RUNG wire#w2
   RUNG wire#powerrail
      Contact( #呼灯 )
      wire#w3
      { S7_Templates := "SrcType := Int" } GT_Contact(in1 := #调度距离1, in2 := #最小调度距离)
      { S7_Templates := "SrcType := Int" } EQ_Contact(in1 := #调度距离2, in2 := #最小调度距离)
      I_Contact( #内外呼重合1 )
      I_Contact( #内外呼重合3 )
      I_Contact( #内外呼重合4 )
      I_Contact( #内外呼重合5 )
      I_Contact( #内外呼重合6 )
      I_Contact( #追击1 )
      I_Contact( #追击3 )
      I_Contact( #追击4 )
      I_Contact( #追击5 )
      I_Contact( #追击6 )
      wire#w4
      Coil( #中间分配2 )
   END_RUNG
   RUNG wire#w3
      Contact( #内外呼重合2 )
   END_RUNG wire#w4
   RUNG wire#w3
      Contact( #追击2 )
      I_Contact( #内外呼重合1 )
      I_Contact( #内外呼重合3 )
      I_Contact( #内外呼重合4 )
      I_Contact( #内外呼重合5 )
      I_Contact( #内外呼重合6 )
   END_RUNG wire#w4
   RUNG wire#powerrail
      Contact( #呼灯 )
      wire#w5
      { S7_Templates := "SrcType := Int" } GT_Contact(in1 := #调度距离1, in2 := #最小调度距离)
      { S7_Templates := "SrcType := Int" } GT_Contact(in1 := #调度距离2, in2 := #最小调度距离)
      { S7_Templates := "SrcType := Int" } EQ_Contact(in1 := #调度距离3, in2 := #最小调度距离)
      I_Contact( #内外呼重合1 )
      I_Contact( #内外呼重合2 )
      I_Contact( #内外呼重合4 )
      I_Contact( #内外呼重合5 )
      I_Contact( #内外呼重合6 )
      I_Contact( #追击1 )
      I_Contact( #追击2 )
      I_Contact( #追击4 )
      I_Contact( #追击5 )
      I_Contact( #追击6 )
      wire#w6
      Coil( #中间分配3 )
   END_RUNG
   RUNG wire#w5
      Contact( #内外呼重合3 )
   END_RUNG wire#w6
   RUNG wire#w5
      Contact( #追击3 )
      I_Contact( #内外呼重合1 )
      I_Contact( #内外呼重合2 )
      I_Contact( #内外呼重合4 )
      I_Contact( #内外呼重合5 )
      I_Contact( #内外呼重合6 )
   END_RUNG wire#w6
   RUNG wire#powerrail
      Contact( #呼灯 )
      wire#w7
      { S7_Templates := "SrcType := Int" } GT_Contact(in1 := #调度距离1, in2 := #最小调度距离)
      { S7_Templates := "SrcType := Int" } GT_Contact(in1 := #调度距离2, in2 := #最小调度距离)
      { S7_Templates := "SrcType := Int" } GT_Contact(in1 := #调度距离3, in2 := #最小调度距离)
      { S7_Templates := "SrcType := Int" } EQ_Contact(in1 := #调度距离4, in2 := #最小调度距离)
      I_Contact( #内外呼重合1 )
      I_Contact( #内外呼重合2 )
      I_Contact( #内外呼重合3 )
      I_Contact( #内外呼重合5 )
      I_Contact( #内外呼重合6 )
      I_Contact( #追击1 )
      I_Contact( #追击2 )
      I_Contact( #追击3 )
      I_Contact( #追击5 )
      I_Contact( #追击6 )
      wire#w8
      Coil( #中间分配4 )
   END_RUNG
   RUNG wire#w7
      Contact( #内外呼重合4 )
   END_RUNG wire#w8
   RUNG wire#w7
      Contact( #追击4 )
      I_Contact( #内外呼重合1 )
      I_Contact( #内外呼重合2 )
      I_Contact( #内外呼重合3 )
      I_Contact( #内外呼重合5 )
      I_Contact( #内外呼重合6 )
   END_RUNG wire#w8
   RUNG wire#powerrail
      Contact( #呼灯 )
      wire#w9
      { S7_Templates := "SrcType := Int" } GT_Contact(in1 := #调度距离1, in2 := #最小调度距离)
      { S7_Templates := "SrcType := Int" } GT_Contact(in1 := #调度距离2, in2 := #最小调度距离)
      { S7_Templates := "SrcType := Int" } GT_Contact(in1 := #调度距离3, in2 := #最小调度距离)
      { S7_Templates := "SrcType := Int" } GT_Contact(in1 := #调度距离4, in2 := #最小调度距离)
      { S7_Templates := "SrcType := Int" } EQ_Contact(in1 := #调度距离5, in2 := #最小调度距离)
      I_Contact( #内外呼重合1 )
      I_Contact( #内外呼重合2 )
      I_Contact( #内外呼重合3 )
      I_Contact( #内外呼重合4 )
      I_Contact( #内外呼重合6 )
      I_Contact( #追击1 )
      I_Contact( #追击2 )
      I_Contact( #追击3 )
      I_Contact( #追击4 )
      I_Contact( #追击6 )
      wire#w10
      Coil( #中间分配5 )
   END_RUNG
   RUNG wire#w9
      Contact( #内外呼重合5 )
   END_RUNG wire#w10
   RUNG wire#w9
      Contact( #追击5 )
      I_Contact( #内外呼重合1 )
      I_Contact( #内外呼重合2 )
      I_Contact( #内外呼重合3 )
      I_Contact( #内外呼重合4 )
      I_Contact( #内外呼重合6 )
   END_RUNG wire#w10
   RUNG wire#powerrail
      Contact( #呼灯 )
      wire#w11
      { S7_Templates := "SrcType := Int" } GT_Contact(in1 := #调度距离1, in2 := #最小调度距离)
      { S7_Templates := "SrcType := Int" } GT_Contact(in1 := #调度距离2, in2 := #最小调度距离)
      { S7_Templates := "SrcType := Int" } GT_Contact(in1 := #调度距离3, in2 := #最小调度距离)
      { S7_Templates := "SrcType := Int" } GT_Contact(in1 := #调度距离4, in2 := #最小调度距离)
      { S7_Templates := "SrcType := Int" } GT_Contact(in1 := #调度距离5, in2 := #最小调度距离)
      { S7_Templates := "SrcType := Int" } EQ_Contact(in1 := #调度距离6, in2 := #最小调度距离)
      I_Contact( #内外呼重合1 )
      I_Contact( #内外呼重合2 )
      I_Contact( #内外呼重合3 )
      I_Contact( #内外呼重合4 )
      I_Contact( #内外呼重合5 )
      I_Contact( #追击1 )
      I_Contact( #追击2 )
      I_Contact( #追击3 )
      I_Contact( #追击4 )
      I_Contact( #追击5 )
      wire#w12
      Coil( #中间分配6 )
   END_RUNG
   RUNG wire#w11
      Contact( #内外呼重合6 )
   END_RUNG wire#w12
   RUNG wire#w11
      Contact( #追击6 )
      I_Contact( #内外呼重合1 )
      I_Contact( #内外呼重合2 )
      I_Contact( #内外呼重合3 )
      I_Contact( #内外呼重合4 )
      I_Contact( #内外呼重合5 )
   END_RUNG wire#w12
   // the same network as SCL:
   #中间分配1 := #呼灯 AND (((#调度距离1 = #最小调度距离) AND NOT #内外呼重合2 AND NOT #内外呼重合3 AND NOT #内外呼重合4 AND NOT #内外呼重合5 AND NOT #内外呼重合6 AND NOT #追击2 AND NOT #追击3 AND NOT #追击4 AND NOT #追击5 AND NOT #追击6) OR #内外呼重合1 OR (#追击1 AND NOT #内外呼重合2 AND NOT #内外呼重合3 AND NOT #内外呼重合4 AND NOT #内外呼重合5 AND NOT #内外呼重合6));
   #中间分配2 := #呼灯 AND (((#调度距离1 > #最小调度距离) AND (#调度距离2 = #最小调度距离) AND NOT #内外呼重合1 AND NOT #内外呼重合3 AND NOT #内外呼重合4 AND NOT #内外呼重合5 AND NOT #内外呼重合6 AND NOT #追击1 AND NOT #追击3 AND NOT #追击4 AND NOT #追击5 AND NOT #追击6) OR #内外呼重合2 OR (#追击2 AND NOT #内外呼重合1 AND NOT #内外呼重合3 AND NOT #内外呼重合4 AND NOT #内外呼重合5 AND NOT #内外呼重合6));
   #中间分配3 := #呼灯 AND (((#调度距离1 > #最小调度距离) AND (#调度距离2 > #最小调度距离) AND (#调度距离3 = #最小调度距离) AND NOT #内外呼重合1 AND NOT #内外呼重合2 AND NOT #内外呼重合4 AND NOT #内外呼重合5 AND NOT #内外呼重合6 AND NOT #追击1 AND NOT #追击2 AND NOT #追击4 AND NOT #追击5 AND NOT #追击6) OR #内外呼重合3 OR (#追击3 AND NOT #内外呼重合1 AND NOT #内外呼重合2 AND NOT #内外呼重合4 AND NOT #内外呼重合5 AND NOT #内外呼重合6));
   #中间分配4 := #呼灯 AND (((#调度距离1 > #最小调度距离) AND (#调度距离2 > #最小调度距离) AND (#调度距离3 > #最小调度距离) AND (#调度距离4 = #最小调度距离) AND NOT #内外呼重合1 AND NOT #内外呼重合2 AND NOT #内外呼重合3 AND NOT #内外呼重合5 AND NOT #内外呼重合6 AND NOT #追击1 AND NOT #追击2 AND NOT #追击3 AND NOT #追击5 AND NOT #追击6) OR #内外呼重合4 OR (#追击4 AND NOT #内外呼重合1 AND NOT #内外呼重合2 AND NOT #内外呼重合3 AND NOT #内外呼重合5 AND NOT #内外呼重合6));
   #中间分配5 := #呼灯 AND (((#调度距离1 > #最小调度距离) AND (#调度距离2 > #最小调度距离) AND (#调度距离3 > #最小调度距离) AND (#调度距离4 > #最小调度距离) AND (#调度距离5 = #最小调度距离) AND NOT #内外呼重合1 AND NOT #内外呼重合2 AND NOT #内外呼重合3 AND NOT #内外呼重合4 AND NOT #内外呼重合6 AND NOT #追击1 AND NOT #追击2 AND NOT #追击3 AND NOT #追击4 AND NOT #追击6) OR #内外呼重合5 OR (#追击5 AND NOT #内外呼重合1 AND NOT #内外呼重合2 AND NOT #内外呼重合3 AND NOT #内外呼重合4 AND NOT #内外呼重合6));
   #中间分配6 := #呼灯 AND (((#调度距离1 > #最小调度距离) AND (#调度距离2 > #最小调度距离) AND (#调度距离3 > #最小调度距离) AND (#调度距离4 > #最小调度距离) AND (#调度距离5 > #最小调度距离) AND (#调度距离6 = #最小调度距离) AND NOT #内外呼重合1 AND NOT #内外呼重合2 AND NOT #内外呼重合3 AND NOT #内外呼重合4 AND NOT #内外呼重合5 AND NOT #追击1 AND NOT #追击2 AND NOT #追击3 AND NOT #追击4 AND NOT #追击5) OR #内外呼重合6 OR (#追击6 AND NOT #内外呼重合1 AND NOT #内外呼重合2 AND NOT #内外呼重合3 AND NOT #内外呼重合4 AND NOT #内外呼重合5));
END_REGION

REGION Network 6: 分配1梯
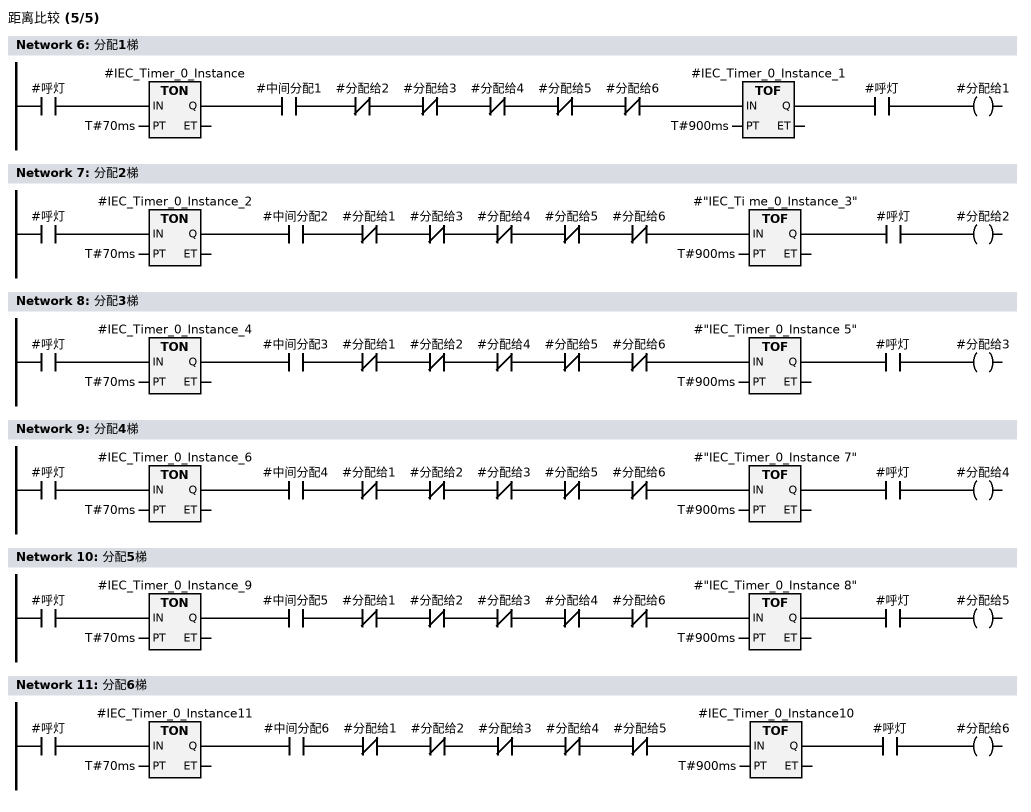
   #IEC_Timer_0_Instance(IN := #呼灯, PT := T#70ms);   // TON
   #IEC_Timer_0_Instance_1(IN := #IEC_Timer_0_Instance.Q AND #中间分配1 AND NOT #分配给2 AND NOT #分配给3 AND NOT #分配给4 AND NOT #分配给5 AND NOT #分配给6,   // TOF
                           PT := T#900ms);
   #分配给1 := #IEC_Timer_0_Instance_1.Q AND #呼灯;
END_REGION

REGION Network 7: 分配2梯
   #IEC_Timer_0_Instance_2(IN := #呼灯, PT := T#70ms);   // TON
   #"IEC_Ti me_0_Instance_3"(IN := #IEC_Timer_0_Instance_2.Q AND #中间分配2 AND NOT #分配给1 AND NOT #分配给3 AND NOT #分配给4 AND NOT #分配给5 AND NOT #分配给6,   // TOF
                           PT := T#900ms);
   #分配给2 := #"IEC_Ti me_0_Instance_3".Q AND #呼灯;
END_REGION

REGION Network 8: 分配3梯
   #IEC_Timer_0_Instance_4(IN := #呼灯, PT := T#70ms);   // TON
   #"IEC_Timer_0_Instance 5"(IN := #IEC_Timer_0_Instance_4.Q AND #中间分配3 AND NOT #分配给1 AND NOT #分配给2 AND NOT #分配给4 AND NOT #分配给5 AND NOT #分配给6,   // TOF
                           PT := T#900ms);
   #分配给3 := #"IEC_Timer_0_Instance 5".Q AND #呼灯;
END_REGION

REGION Network 9: 分配4梯
   #IEC_Timer_0_Instance_6(IN := #呼灯, PT := T#70ms);   // TON
   #"IEC_Timer_0_Instance 7"(IN := #IEC_Timer_0_Instance_6.Q AND #中间分配4 AND NOT #分配给1 AND NOT #分配给2 AND NOT #分配给3 AND NOT #分配给5 AND NOT #分配给6,   // TOF
                           PT := T#900ms);
   #分配给4 := #"IEC_Timer_0_Instance 7".Q AND #呼灯;
END_REGION

REGION Network 10: 分配5梯
   #IEC_Timer_0_Instance_9(IN := #呼灯, PT := T#70ms);   // TON
   #"IEC_Timer_0_Instance 8"(IN := #IEC_Timer_0_Instance_9.Q AND #中间分配5 AND NOT #分配给1 AND NOT #分配给2 AND NOT #分配给3 AND NOT #分配给4 AND NOT #分配给6,   // TOF
                           PT := T#900ms);
   #分配给5 := #"IEC_Timer_0_Instance 8".Q AND #呼灯;
END_REGION

REGION Network 11: 分配6梯
   #IEC_Timer_0_Instance11(IN := #呼灯, PT := T#70ms);   // TON
   #IEC_Timer_0_Instance10(IN := #IEC_Timer_0_Instance11.Q AND #中间分配6 AND NOT #分配给1 AND NOT #分配给2 AND NOT #分配给3 AND NOT #分配给4 AND NOT #分配给5,   // TOF
                           PT := T#900ms);
   #分配给6 := #IEC_Timer_0_Instance10.Q AND #呼灯;
END_REGION
END_FUNCTION_BLOCK

FUNCTION_BLOCK "目标判断"   // FB2, LAD
{ S7_Optimized_Access := 'TRUE' }
VERSION : 0.1
   VAR_INPUT
      "1层上呼分配" : Bool;
      "2层上呼分配" : Bool;
      "2层下呼分配" : Bool;
      "3层上呼分配" : Bool;
      "3层下呼分配" : Bool;
      "4层上呼分配" : Bool;
      "4层下呼分配" : Bool;
      "5层上呼分配" : Bool;
      "5层下呼分配" : Bool;
      "6层上呼分配" : Bool;
      "6层下呼分配" : Bool;
      "7层上呼分配" : Bool;
      "7层下呼分配" : Bool;
      "8层上呼分配" : Bool;
      "8层下呼分配" : Bool;
      "9层上呼分配" : Bool;
      "9层下呼分配" : Bool;
      "10层下呼分配" : Bool;
      内呼按钮1 : Bool;
      内呼按钮2 : Bool;
      内呼按钮3 : Bool;
      内呼按钮4 : Bool;
      内呼按钮5 : Bool;
      内呼按钮6 : Bool;
      内呼按钮7 : Bool;
      内呼按钮8 : Bool;
      内呼按钮9 : Bool;
      内呼按钮10 : Bool;
   END_VAR
   VAR_OUTPUT
      外呼下面无目标2 : Bool;
      外呼下面无目标3 : Bool;
      外呼下面无目标4 : Bool;
      外呼下面无目标5 : Bool;
      外呼下面无目标6 : Bool;
      外呼下面无目标7 : Bool;
      外呼下面无目标8 : Bool;
      外呼下面无目标9 : Bool;
      外呼上面无目标2 : Bool;
      外呼上面无目标3 : Bool;
      外呼上面无目标4 : Bool;
      外呼上面无目标5 : Bool;
      外呼上面无目标6 : Bool;
      外呼上面无目标7 : Bool;
      外呼上面无目标8 : Bool;
      外呼上面无目标9 : Bool;
      外呼上面有目标1 : Bool;
      外呼上面有目标2 : Bool;
      外呼上面有目标3 : Bool;
      外呼上面有目标4 : Bool;
      外呼上面有目标5 : Bool;
      外呼上面有目标6 : Bool;
      外呼上面有目标7 : Bool;
      外呼上面有目标8 : Bool;
      外呼上面有目标9 : Bool;
      外呼下面有目标2 : Bool;
      外呼下面有目标3 : Bool;
      外呼下面有目标4 : Bool;
      外呼下面有目标5 : Bool;
      外呼下面有目标6 : Bool;
      外呼下面有目标7 : Bool;
      外呼下面有目标8 : Bool;
      外呼下面有目标9 : Bool;
      外呼下面有目标10 : Bool;
      外呼上面有最大目标数1 : Int;
      外呼上面有最大目标数2 : Int;
      外呼上面有最大目标数3 : Int;
      外呼上面有最大目标数4 : Int;
      外呼上面有最大目标数5 : Int;
      外呼上面有最大目标数6 : Int;
      外呼上面有最大目标数7 : Int;
      外呼上面有最大目标数8 : Int;
      外呼上面有最大目标数9 : Int;
      外呼下面有最小目标数2 : Int;
      外呼下面有最小目标数3 : Int;
      外呼下面有最小目标数4 : Int;
      外呼下面有最小目标数5 : Int;
      外呼下面有最小目标数6 : Int;
      外呼下面有最小目标数7 : Int;
      外呼下面有最小目标数8 : Int;
      外呼下面有最小目标数9 : Int;
      外呼下面有最小目标数10 : Int;
   END_VAR
   VAR
      目标楼层数1 : Int;
      目标楼层数2 : Int;
      目标楼层数3 : Int;
      目标楼层数4 : Int;
      目标楼层数5 : Int;
      目标楼层数6 : Int;
      目标楼层数7 : Int;
      目标楼层数8 : Int;
      目标楼层数9 : Int;
      目标楼层数10 : Int;
      无目标 : Bool;
   END_VAR
BEGIN

REGION Network 1: 外呼下面无目标
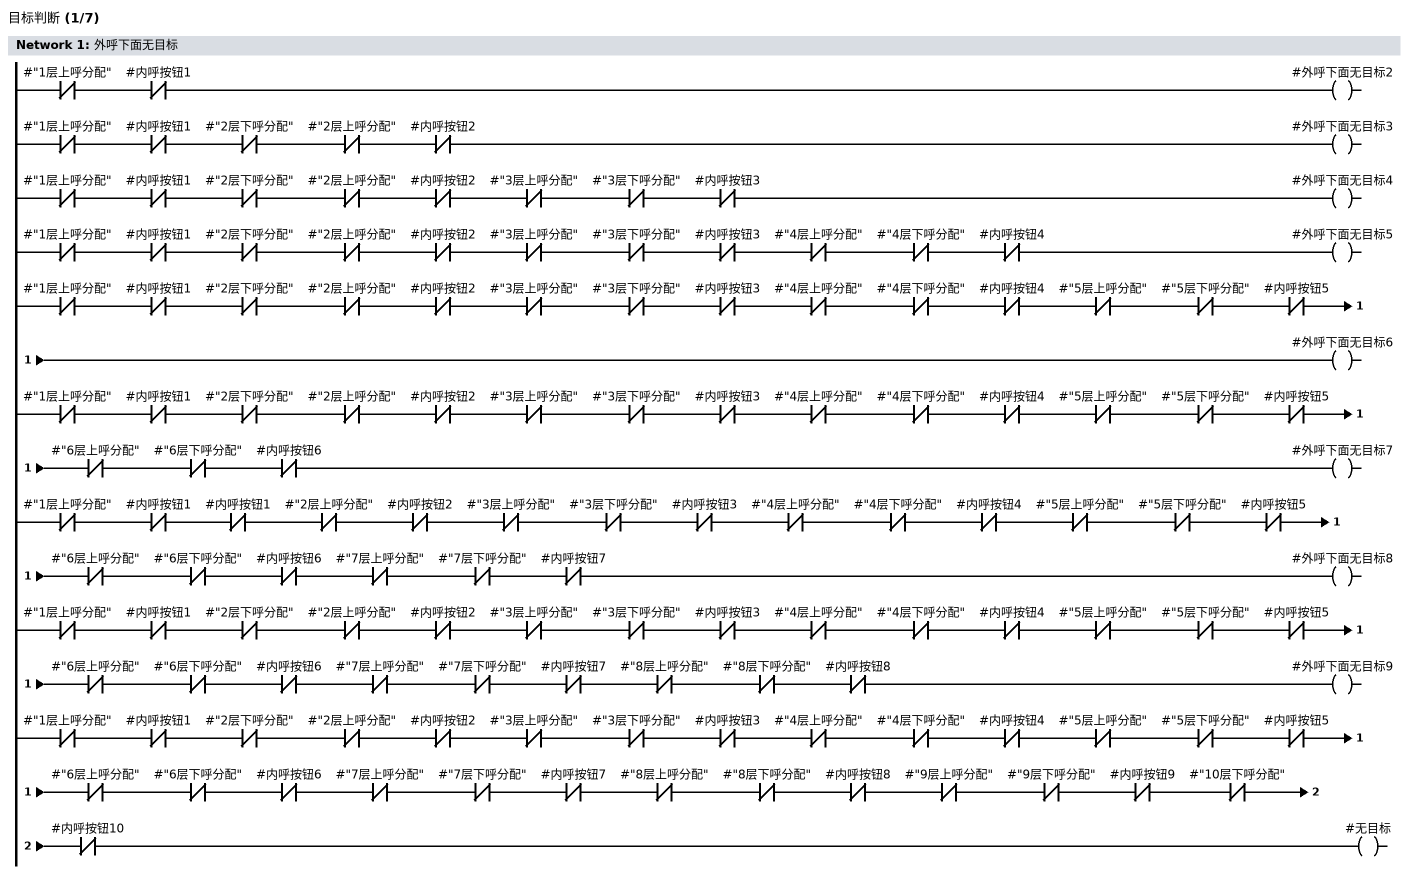
   RUNG wire#powerrail
      I_Contact( #"1层上呼分配" )
      I_Contact( #内呼按钮1 )
      Coil( #外呼下面无目标2 )
   END_RUNG
   RUNG wire#powerrail
      I_Contact( #"1层上呼分配" )
      I_Contact( #内呼按钮1 )
      I_Contact( #"2层下呼分配" )
      I_Contact( #"2层上呼分配" )
      I_Contact( #内呼按钮2 )
      Coil( #外呼下面无目标3 )
   END_RUNG
   RUNG wire#powerrail
      I_Contact( #"1层上呼分配" )
      I_Contact( #内呼按钮1 )
      I_Contact( #"2层下呼分配" )
      I_Contact( #"2层上呼分配" )
      I_Contact( #内呼按钮2 )
      I_Contact( #"3层上呼分配" )
      I_Contact( #"3层下呼分配" )
      I_Contact( #内呼按钮3 )
      Coil( #外呼下面无目标4 )
   END_RUNG
   RUNG wire#powerrail
      I_Contact( #"1层上呼分配" )
      I_Contact( #内呼按钮1 )
      I_Contact( #"2层下呼分配" )
      I_Contact( #"2层上呼分配" )
      I_Contact( #内呼按钮2 )
      I_Contact( #"3层上呼分配" )
      I_Contact( #"3层下呼分配" )
      I_Contact( #内呼按钮3 )
      I_Contact( #"4层上呼分配" )
      I_Contact( #"4层下呼分配" )
      I_Contact( #内呼按钮4 )
      Coil( #外呼下面无目标5 )
   END_RUNG
   RUNG wire#powerrail
      I_Contact( #"1层上呼分配" )
      I_Contact( #内呼按钮1 )
      I_Contact( #"2层下呼分配" )
      I_Contact( #"2层上呼分配" )
      I_Contact( #内呼按钮2 )
      I_Contact( #"3层上呼分配" )
      I_Contact( #"3层下呼分配" )
      I_Contact( #内呼按钮3 )
      I_Contact( #"4层上呼分配" )
      I_Contact( #"4层下呼分配" )
      I_Contact( #内呼按钮4 )
      I_Contact( #"5层上呼分配" )
      I_Contact( #"5层下呼分配" )
      I_Contact( #内呼按钮5 )
      Coil( #外呼下面无目标6 )
   END_RUNG
   RUNG wire#powerrail
      I_Contact( #"1层上呼分配" )
      I_Contact( #内呼按钮1 )
      I_Contact( #"2层下呼分配" )
      I_Contact( #"2层上呼分配" )
      I_Contact( #内呼按钮2 )
      I_Contact( #"3层上呼分配" )
      I_Contact( #"3层下呼分配" )
      I_Contact( #内呼按钮3 )
      I_Contact( #"4层上呼分配" )
      I_Contact( #"4层下呼分配" )
      I_Contact( #内呼按钮4 )
      I_Contact( #"5层上呼分配" )
      I_Contact( #"5层下呼分配" )
      I_Contact( #内呼按钮5 )
      I_Contact( #"6层上呼分配" )
      I_Contact( #"6层下呼分配" )
      I_Contact( #内呼按钮6 )
      Coil( #外呼下面无目标7 )
   END_RUNG
   RUNG wire#powerrail
      I_Contact( #"1层上呼分配" )
      I_Contact( #内呼按钮1 )
      I_Contact( #内呼按钮1 )
      I_Contact( #"2层上呼分配" )
      I_Contact( #内呼按钮2 )
      I_Contact( #"3层上呼分配" )
      I_Contact( #"3层下呼分配" )
      I_Contact( #内呼按钮3 )
      I_Contact( #"4层上呼分配" )
      I_Contact( #"4层下呼分配" )
      I_Contact( #内呼按钮4 )
      I_Contact( #"5层上呼分配" )
      I_Contact( #"5层下呼分配" )
      I_Contact( #内呼按钮5 )
      I_Contact( #"6层上呼分配" )
      I_Contact( #"6层下呼分配" )
      I_Contact( #内呼按钮6 )
      I_Contact( #"7层上呼分配" )
      I_Contact( #"7层下呼分配" )
      I_Contact( #内呼按钮7 )
      Coil( #外呼下面无目标8 )
   END_RUNG
   RUNG wire#powerrail
      I_Contact( #"1层上呼分配" )
      I_Contact( #内呼按钮1 )
      I_Contact( #"2层下呼分配" )
      I_Contact( #"2层上呼分配" )
      I_Contact( #内呼按钮2 )
      I_Contact( #"3层上呼分配" )
      I_Contact( #"3层下呼分配" )
      I_Contact( #内呼按钮3 )
      I_Contact( #"4层上呼分配" )
      I_Contact( #"4层下呼分配" )
      I_Contact( #内呼按钮4 )
      I_Contact( #"5层上呼分配" )
      I_Contact( #"5层下呼分配" )
      I_Contact( #内呼按钮5 )
      I_Contact( #"6层上呼分配" )
      I_Contact( #"6层下呼分配" )
      I_Contact( #内呼按钮6 )
      I_Contact( #"7层上呼分配" )
      I_Contact( #"7层下呼分配" )
      I_Contact( #内呼按钮7 )
      I_Contact( #"8层上呼分配" )
      I_Contact( #"8层下呼分配" )
      I_Contact( #内呼按钮8 )
      Coil( #外呼下面无目标9 )
   END_RUNG
   RUNG wire#powerrail
      I_Contact( #"1层上呼分配" )
      I_Contact( #内呼按钮1 )
      I_Contact( #"2层下呼分配" )
      I_Contact( #"2层上呼分配" )
      I_Contact( #内呼按钮2 )
      I_Contact( #"3层上呼分配" )
      I_Contact( #"3层下呼分配" )
      I_Contact( #内呼按钮3 )
      I_Contact( #"4层上呼分配" )
      I_Contact( #"4层下呼分配" )
      I_Contact( #内呼按钮4 )
      I_Contact( #"5层上呼分配" )
      I_Contact( #"5层下呼分配" )
      I_Contact( #内呼按钮5 )
      I_Contact( #"6层上呼分配" )
      I_Contact( #"6层下呼分配" )
      I_Contact( #内呼按钮6 )
      I_Contact( #"7层上呼分配" )
      I_Contact( #"7层下呼分配" )
      I_Contact( #内呼按钮7 )
      I_Contact( #"8层上呼分配" )
      I_Contact( #"8层下呼分配" )
      I_Contact( #内呼按钮8 )
      I_Contact( #"9层上呼分配" )
      I_Contact( #"9层下呼分配" )
      I_Contact( #内呼按钮9 )
      I_Contact( #"10层下呼分配" )
      I_Contact( #内呼按钮10 )
      Coil( #无目标 )
   END_RUNG
   // the same network as SCL:
   #外呼下面无目标2 := NOT #"1层上呼分配" AND NOT #内呼按钮1;
   #外呼下面无目标3 := NOT #"1层上呼分配" AND NOT #内呼按钮1 AND NOT #"2层下呼分配" AND NOT #"2层上呼分配" AND NOT #内呼按钮2;
   #外呼下面无目标4 := NOT #"1层上呼分配" AND NOT #内呼按钮1 AND NOT #"2层下呼分配" AND NOT #"2层上呼分配" AND NOT #内呼按钮2 AND NOT #"3层上呼分配" AND NOT #"3层下呼分配" AND NOT #内呼按钮3;
   #外呼下面无目标5 := NOT #"1层上呼分配" AND NOT #内呼按钮1 AND NOT #"2层下呼分配" AND NOT #"2层上呼分配" AND NOT #内呼按钮2 AND NOT #"3层上呼分配" AND NOT #"3层下呼分配" AND NOT #内呼按钮3 AND NOT #"4层上呼分配" AND NOT #"4层下呼分配" AND NOT #内呼按钮4;
   #外呼下面无目标6 := NOT #"1层上呼分配" AND NOT #内呼按钮1 AND NOT #"2层下呼分配" AND NOT #"2层上呼分配" AND NOT #内呼按钮2 AND NOT #"3层上呼分配" AND NOT #"3层下呼分配" AND NOT #内呼按钮3 AND NOT #"4层上呼分配" AND NOT #"4层下呼分配" AND NOT #内呼按钮4 AND NOT #"5层上呼分配" AND NOT #"5层下呼分配" AND NOT #内呼按钮5;
   #外呼下面无目标7 := NOT #"1层上呼分配" AND NOT #内呼按钮1 AND NOT #"2层下呼分配" AND NOT #"2层上呼分配" AND NOT #内呼按钮2 AND NOT #"3层上呼分配" AND NOT #"3层下呼分配" AND NOT #内呼按钮3 AND NOT #"4层上呼分配" AND NOT #"4层下呼分配" AND NOT #内呼按钮4 AND NOT #"5层上呼分配" AND NOT #"5层下呼分配" AND NOT #内呼按钮5 AND NOT #"6层上呼分配" AND NOT #"6层下呼分配" AND NOT #内呼按钮6;
   #外呼下面无目标8 := NOT #"1层上呼分配" AND NOT #内呼按钮1 AND NOT #内呼按钮1 AND NOT #"2层上呼分配" AND NOT #内呼按钮2 AND NOT #"3层上呼分配" AND NOT #"3层下呼分配" AND NOT #内呼按钮3 AND NOT #"4层上呼分配" AND NOT #"4层下呼分配" AND NOT #内呼按钮4 AND NOT #"5层上呼分配" AND NOT #"5层下呼分配" AND NOT #内呼按钮5 AND NOT #"6层上呼分配" AND NOT #"6层下呼分配" AND NOT #内呼按钮6 AND NOT #"7层上呼分配" AND NOT #"7层下呼分配" AND NOT #内呼按钮7;
   #外呼下面无目标9 := NOT #"1层上呼分配" AND NOT #内呼按钮1 AND NOT #"2层下呼分配" AND NOT #"2层上呼分配" AND NOT #内呼按钮2 AND NOT #"3层上呼分配" AND NOT #"3层下呼分配" AND NOT #内呼按钮3 AND NOT #"4层上呼分配" AND NOT #"4层下呼分配" AND NOT #内呼按钮4 AND NOT #"5层上呼分配" AND NOT #"5层下呼分配" AND NOT #内呼按钮5 AND NOT #"6层上呼分配" AND NOT #"6层下呼分配" AND NOT #内呼按钮6 AND NOT #"7层上呼分配" AND NOT #"7层下呼分配" AND NOT #内呼按钮7 AND NOT #"8层上呼分配" AND NOT #"8层下呼分配" AND NOT #内呼按钮8;
   #无目标 := NOT #"1层上呼分配" AND NOT #内呼按钮1 AND NOT #"2层下呼分配" AND NOT #"2层上呼分配" AND NOT #内呼按钮2 AND NOT #"3层上呼分配" AND NOT #"3层下呼分配" AND NOT #内呼按钮3 AND NOT #"4层上呼分配" AND NOT #"4层下呼分配" AND NOT #内呼按钮4 AND NOT #"5层上呼分配" AND NOT #"5层下呼分配" AND NOT #内呼按钮5 AND NOT #"6层上呼分配" AND NOT #"6层下呼分配" AND NOT #内呼按钮6 AND NOT #"7层上呼分配" AND NOT #"7层下呼分配" AND NOT #内呼按钮7 AND NOT #"8层上呼分配" AND NOT #"8层下呼分配" AND NOT #内呼按钮8 AND NOT #"9层上呼分配" AND NOT #"9层下呼分配" AND NOT #内呼按钮9 AND NOT #"10层下呼分配" AND NOT #内呼按钮10;
END_REGION

REGION Network 2: 外呼上面无目标
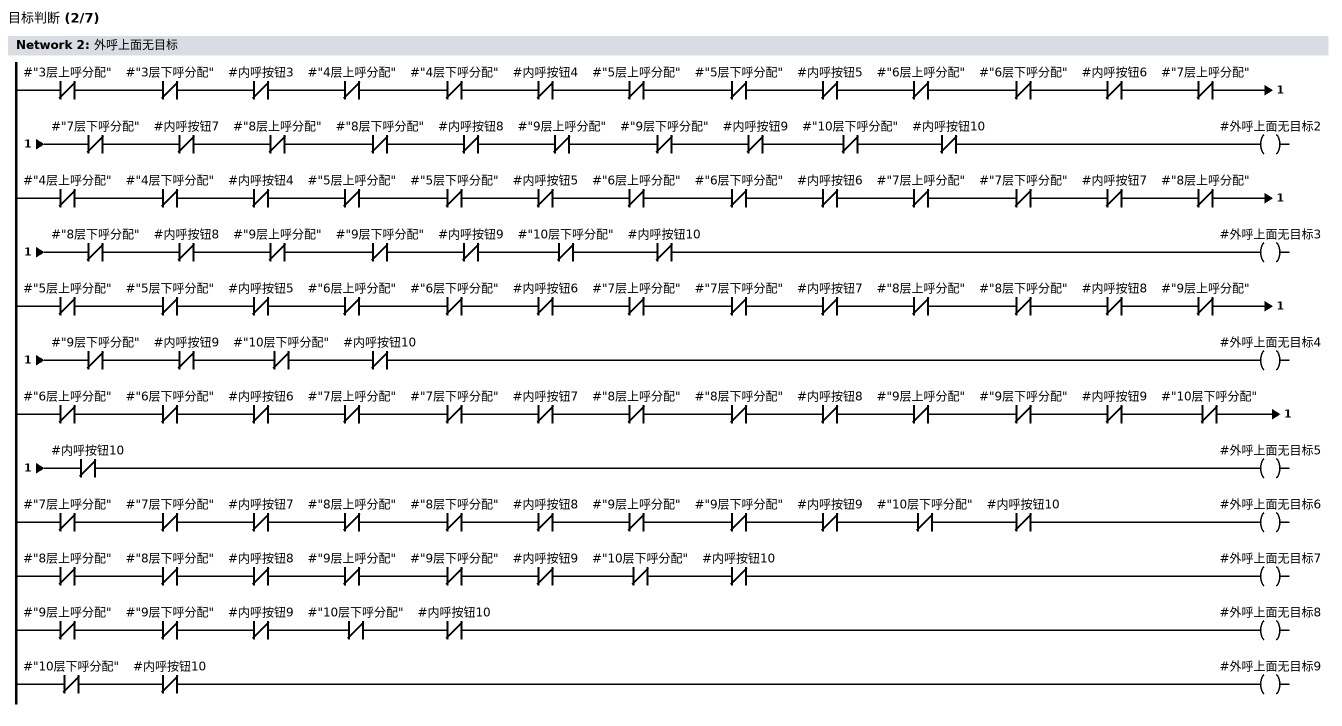
   RUNG wire#powerrail
      I_Contact( #"3层上呼分配" )
      I_Contact( #"3层下呼分配" )
      I_Contact( #内呼按钮3 )
      I_Contact( #"4层上呼分配" )
      I_Contact( #"4层下呼分配" )
      I_Contact( #内呼按钮4 )
      I_Contact( #"5层上呼分配" )
      I_Contact( #"5层下呼分配" )
      I_Contact( #内呼按钮5 )
      I_Contact( #"6层上呼分配" )
      I_Contact( #"6层下呼分配" )
      I_Contact( #内呼按钮6 )
      I_Contact( #"7层上呼分配" )
      I_Contact( #"7层下呼分配" )
      I_Contact( #内呼按钮7 )
      I_Contact( #"8层上呼分配" )
      I_Contact( #"8层下呼分配" )
      I_Contact( #内呼按钮8 )
      I_Contact( #"9层上呼分配" )
      I_Contact( #"9层下呼分配" )
      I_Contact( #内呼按钮9 )
      I_Contact( #"10层下呼分配" )
      I_Contact( #内呼按钮10 )
      Coil( #外呼上面无目标2 )
   END_RUNG
   RUNG wire#powerrail
      I_Contact( #"4层上呼分配" )
      I_Contact( #"4层下呼分配" )
      I_Contact( #内呼按钮4 )
      I_Contact( #"5层上呼分配" )
      I_Contact( #"5层下呼分配" )
      I_Contact( #内呼按钮5 )
      I_Contact( #"6层上呼分配" )
      I_Contact( #"6层下呼分配" )
      I_Contact( #内呼按钮6 )
      I_Contact( #"7层上呼分配" )
      I_Contact( #"7层下呼分配" )
      I_Contact( #内呼按钮7 )
      I_Contact( #"8层上呼分配" )
      I_Contact( #"8层下呼分配" )
      I_Contact( #内呼按钮8 )
      I_Contact( #"9层上呼分配" )
      I_Contact( #"9层下呼分配" )
      I_Contact( #内呼按钮9 )
      I_Contact( #"10层下呼分配" )
      I_Contact( #内呼按钮10 )
      Coil( #外呼上面无目标3 )
   END_RUNG
   RUNG wire#powerrail
      I_Contact( #"5层上呼分配" )
      I_Contact( #"5层下呼分配" )
      I_Contact( #内呼按钮5 )
      I_Contact( #"6层上呼分配" )
      I_Contact( #"6层下呼分配" )
      I_Contact( #内呼按钮6 )
      I_Contact( #"7层上呼分配" )
      I_Contact( #"7层下呼分配" )
      I_Contact( #内呼按钮7 )
      I_Contact( #"8层上呼分配" )
      I_Contact( #"8层下呼分配" )
      I_Contact( #内呼按钮8 )
      I_Contact( #"9层上呼分配" )
      I_Contact( #"9层下呼分配" )
      I_Contact( #内呼按钮9 )
      I_Contact( #"10层下呼分配" )
      I_Contact( #内呼按钮10 )
      Coil( #外呼上面无目标4 )
   END_RUNG
   RUNG wire#powerrail
      I_Contact( #"6层上呼分配" )
      I_Contact( #"6层下呼分配" )
      I_Contact( #内呼按钮6 )
      I_Contact( #"7层上呼分配" )
      I_Contact( #"7层下呼分配" )
      I_Contact( #内呼按钮7 )
      I_Contact( #"8层上呼分配" )
      I_Contact( #"8层下呼分配" )
      I_Contact( #内呼按钮8 )
      I_Contact( #"9层上呼分配" )
      I_Contact( #"9层下呼分配" )
      I_Contact( #内呼按钮9 )
      I_Contact( #"10层下呼分配" )
      I_Contact( #内呼按钮10 )
      Coil( #外呼上面无目标5 )
   END_RUNG
   RUNG wire#powerrail
      I_Contact( #"7层上呼分配" )
      I_Contact( #"7层下呼分配" )
      I_Contact( #内呼按钮7 )
      I_Contact( #"8层上呼分配" )
      I_Contact( #"8层下呼分配" )
      I_Contact( #内呼按钮8 )
      I_Contact( #"9层上呼分配" )
      I_Contact( #"9层下呼分配" )
      I_Contact( #内呼按钮9 )
      I_Contact( #"10层下呼分配" )
      I_Contact( #内呼按钮10 )
      Coil( #外呼上面无目标6 )
   END_RUNG
   RUNG wire#powerrail
      I_Contact( #"8层上呼分配" )
      I_Contact( #"8层下呼分配" )
      I_Contact( #内呼按钮8 )
      I_Contact( #"9层上呼分配" )
      I_Contact( #"9层下呼分配" )
      I_Contact( #内呼按钮9 )
      I_Contact( #"10层下呼分配" )
      I_Contact( #内呼按钮10 )
      Coil( #外呼上面无目标7 )
   END_RUNG
   RUNG wire#powerrail
      I_Contact( #"9层上呼分配" )
      I_Contact( #"9层下呼分配" )
      I_Contact( #内呼按钮9 )
      I_Contact( #"10层下呼分配" )
      I_Contact( #内呼按钮10 )
      Coil( #外呼上面无目标8 )
   END_RUNG
   RUNG wire#powerrail
      I_Contact( #"10层下呼分配" )
      I_Contact( #内呼按钮10 )
      Coil( #外呼上面无目标9 )
   END_RUNG
   // the same network as SCL:
   #外呼上面无目标2 := NOT #"3层上呼分配" AND NOT #"3层下呼分配" AND NOT #内呼按钮3 AND NOT #"4层上呼分配" AND NOT #"4层下呼分配" AND NOT #内呼按钮4 AND NOT #"5层上呼分配" AND NOT #"5层下呼分配" AND NOT #内呼按钮5 AND NOT #"6层上呼分配" AND NOT #"6层下呼分配" AND NOT #内呼按钮6 AND NOT #"7层上呼分配" AND NOT #"7层下呼分配" AND NOT #内呼按钮7 AND NOT #"8层上呼分配" AND NOT #"8层下呼分配" AND NOT #内呼按钮8 AND NOT #"9层上呼分配" AND NOT #"9层下呼分配" AND NOT #内呼按钮9 AND NOT #"10层下呼分配" AND NOT #内呼按钮10;
   #外呼上面无目标3 := NOT #"4层上呼分配" AND NOT #"4层下呼分配" AND NOT #内呼按钮4 AND NOT #"5层上呼分配" AND NOT #"5层下呼分配" AND NOT #内呼按钮5 AND NOT #"6层上呼分配" AND NOT #"6层下呼分配" AND NOT #内呼按钮6 AND NOT #"7层上呼分配" AND NOT #"7层下呼分配" AND NOT #内呼按钮7 AND NOT #"8层上呼分配" AND NOT #"8层下呼分配" AND NOT #内呼按钮8 AND NOT #"9层上呼分配" AND NOT #"9层下呼分配" AND NOT #内呼按钮9 AND NOT #"10层下呼分配" AND NOT #内呼按钮10;
   #外呼上面无目标4 := NOT #"5层上呼分配" AND NOT #"5层下呼分配" AND NOT #内呼按钮5 AND NOT #"6层上呼分配" AND NOT #"6层下呼分配" AND NOT #内呼按钮6 AND NOT #"7层上呼分配" AND NOT #"7层下呼分配" AND NOT #内呼按钮7 AND NOT #"8层上呼分配" AND NOT #"8层下呼分配" AND NOT #内呼按钮8 AND NOT #"9层上呼分配" AND NOT #"9层下呼分配" AND NOT #内呼按钮9 AND NOT #"10层下呼分配" AND NOT #内呼按钮10;
   #外呼上面无目标5 := NOT #"6层上呼分配" AND NOT #"6层下呼分配" AND NOT #内呼按钮6 AND NOT #"7层上呼分配" AND NOT #"7层下呼分配" AND NOT #内呼按钮7 AND NOT #"8层上呼分配" AND NOT #"8层下呼分配" AND NOT #内呼按钮8 AND NOT #"9层上呼分配" AND NOT #"9层下呼分配" AND NOT #内呼按钮9 AND NOT #"10层下呼分配" AND NOT #内呼按钮10;
   #外呼上面无目标6 := NOT #"7层上呼分配" AND NOT #"7层下呼分配" AND NOT #内呼按钮7 AND NOT #"8层上呼分配" AND NOT #"8层下呼分配" AND NOT #内呼按钮8 AND NOT #"9层上呼分配" AND NOT #"9层下呼分配" AND NOT #内呼按钮9 AND NOT #"10层下呼分配" AND NOT #内呼按钮10;
   #外呼上面无目标7 := NOT #"8层上呼分配" AND NOT #"8层下呼分配" AND NOT #内呼按钮8 AND NOT #"9层上呼分配" AND NOT #"9层下呼分配" AND NOT #内呼按钮9 AND NOT #"10层下呼分配" AND NOT #内呼按钮10;
   #外呼上面无目标8 := NOT #"9层上呼分配" AND NOT #"9层下呼分配" AND NOT #内呼按钮9 AND NOT #"10层下呼分配" AND NOT #内呼按钮10;
   #外呼上面无目标9 := NOT #"10层下呼分配" AND NOT #内呼按钮10;
END_REGION

REGION Network 3: 目标转数字
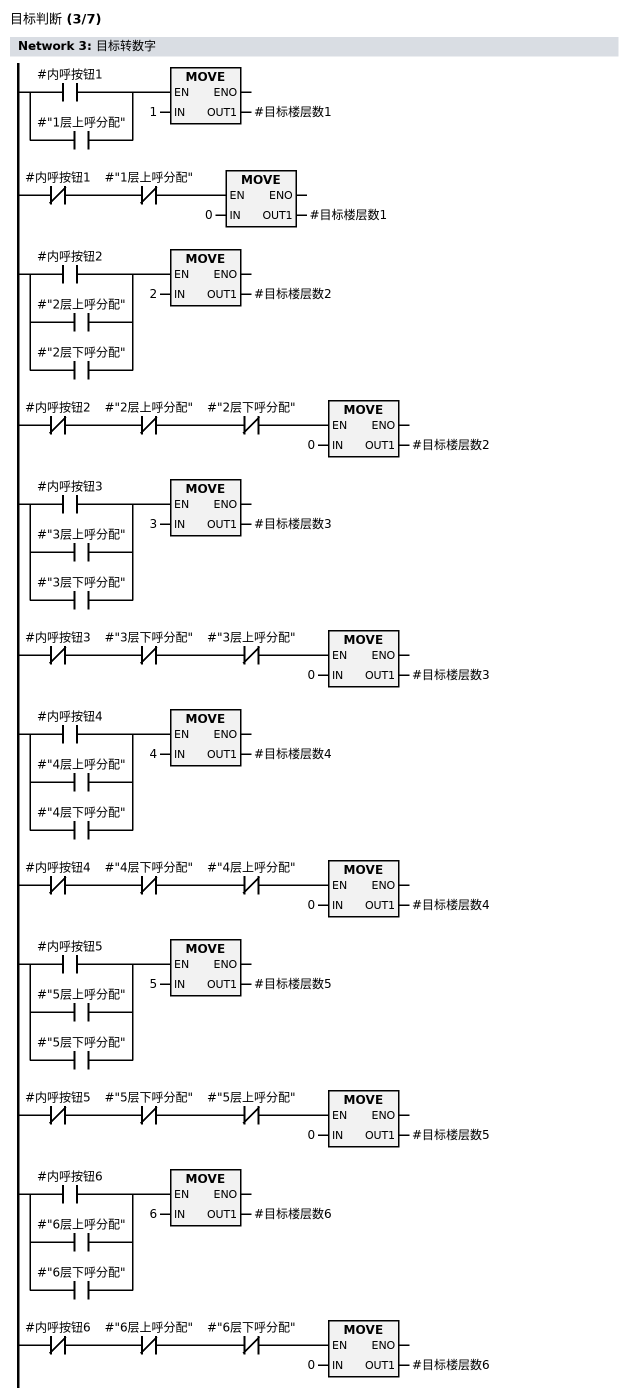
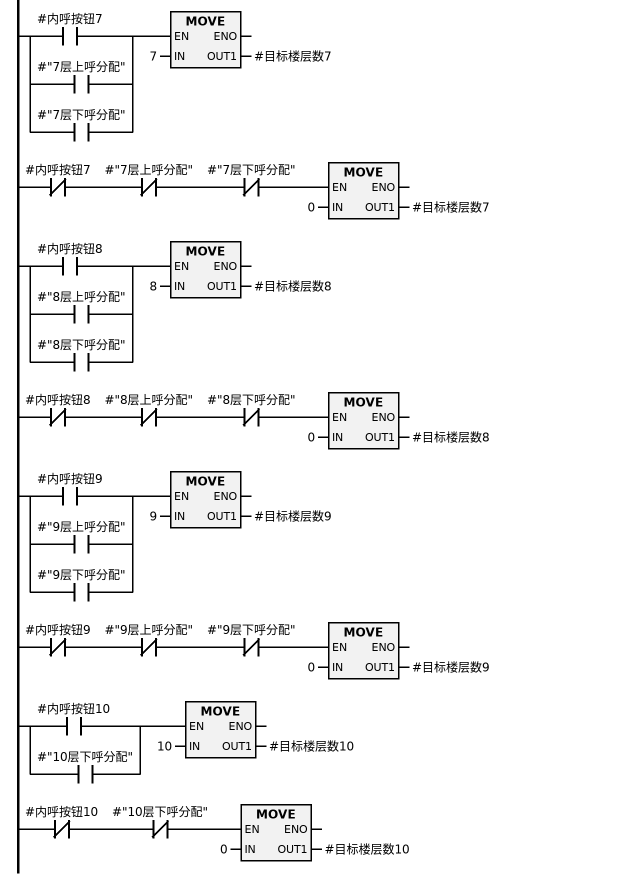
   RUNG wire#powerrail
      Contact( #内呼按钮1 )
      wire#w1
      Move(in := 1, out1 => #目标楼层数1)
   END_RUNG
   RUNG wire#powerrail
      Contact( #"1层上呼分配" )
   END_RUNG wire#w1
   RUNG wire#powerrail
      I_Contact( #内呼按钮1 )
      I_Contact( #"1层上呼分配" )
      Move(in := 0, out1 => #目标楼层数1)
   END_RUNG
   RUNG wire#powerrail
      Contact( #内呼按钮2 )
      wire#w2
      Move(in := 2, out1 => #目标楼层数2)
   END_RUNG
   RUNG wire#powerrail
      Contact( #"2层上呼分配" )
   END_RUNG wire#w2
   RUNG wire#powerrail
      Contact( #"2层下呼分配" )
   END_RUNG wire#w2
   RUNG wire#powerrail
      I_Contact( #内呼按钮2 )
      I_Contact( #"2层上呼分配" )
      I_Contact( #"2层下呼分配" )
      Move(in := 0, out1 => #目标楼层数2)
   END_RUNG
   RUNG wire#powerrail
      Contact( #内呼按钮3 )
      wire#w3
      Move(in := 3, out1 => #目标楼层数3)
   END_RUNG
   RUNG wire#powerrail
      Contact( #"3层上呼分配" )
   END_RUNG wire#w3
   RUNG wire#powerrail
      Contact( #"3层下呼分配" )
   END_RUNG wire#w3
   RUNG wire#powerrail
      I_Contact( #内呼按钮3 )
      I_Contact( #"3层下呼分配" )
      I_Contact( #"3层上呼分配" )
      Move(in := 0, out1 => #目标楼层数3)
   END_RUNG
   RUNG wire#powerrail
      Contact( #内呼按钮4 )
      wire#w4
      Move(in := 4, out1 => #目标楼层数4)
   END_RUNG
   RUNG wire#powerrail
      Contact( #"4层上呼分配" )
   END_RUNG wire#w4
   RUNG wire#powerrail
      Contact( #"4层下呼分配" )
   END_RUNG wire#w4
   RUNG wire#powerrail
      I_Contact( #内呼按钮4 )
      I_Contact( #"4层下呼分配" )
      I_Contact( #"4层上呼分配" )
      Move(in := 0, out1 => #目标楼层数4)
   END_RUNG
   RUNG wire#powerrail
      Contact( #内呼按钮5 )
      wire#w5
      Move(in := 5, out1 => #目标楼层数5)
   END_RUNG
   RUNG wire#powerrail
      Contact( #"5层上呼分配" )
   END_RUNG wire#w5
   RUNG wire#powerrail
      Contact( #"5层下呼分配" )
   END_RUNG wire#w5
   RUNG wire#powerrail
      I_Contact( #内呼按钮5 )
      I_Contact( #"5层下呼分配" )
      I_Contact( #"5层上呼分配" )
      Move(in := 0, out1 => #目标楼层数5)
   END_RUNG
   RUNG wire#powerrail
      Contact( #内呼按钮6 )
      wire#w6
      Move(in := 6, out1 => #目标楼层数6)
   END_RUNG
   RUNG wire#powerrail
      Contact( #"6层上呼分配" )
   END_RUNG wire#w6
   RUNG wire#powerrail
      Contact( #"6层下呼分配" )
   END_RUNG wire#w6
   RUNG wire#powerrail
      I_Contact( #内呼按钮6 )
      I_Contact( #"6层上呼分配" )
      I_Contact( #"6层下呼分配" )
      Move(in := 0, out1 => #目标楼层数6)
   END_RUNG
   RUNG wire#powerrail
      Contact( #内呼按钮7 )
      wire#w7
      Move(in := 7, out1 => #目标楼层数7)
   END_RUNG
   RUNG wire#powerrail
      Contact( #"7层上呼分配" )
   END_RUNG wire#w7
   RUNG wire#powerrail
      Contact( #"7层下呼分配" )
   END_RUNG wire#w7
   RUNG wire#powerrail
      I_Contact( #内呼按钮7 )
      I_Contact( #"7层上呼分配" )
      I_Contact( #"7层下呼分配" )
      Move(in := 0, out1 => #目标楼层数7)
   END_RUNG
   RUNG wire#powerrail
      Contact( #内呼按钮8 )
      wire#w8
      Move(in := 8, out1 => #目标楼层数8)
   END_RUNG
   RUNG wire#powerrail
      Contact( #"8层上呼分配" )
   END_RUNG wire#w8
   RUNG wire#powerrail
      Contact( #"8层下呼分配" )
   END_RUNG wire#w8
   RUNG wire#powerrail
      I_Contact( #内呼按钮8 )
      I_Contact( #"8层上呼分配" )
      I_Contact( #"8层下呼分配" )
      Move(in := 0, out1 => #目标楼层数8)
   END_RUNG
   RUNG wire#powerrail
      Contact( #内呼按钮9 )
      wire#w9
      Move(in := 9, out1 => #目标楼层数9)
   END_RUNG
   RUNG wire#powerrail
      Contact( #"9层上呼分配" )
   END_RUNG wire#w9
   RUNG wire#powerrail
      Contact( #"9层下呼分配" )
   END_RUNG wire#w9
   RUNG wire#powerrail
      I_Contact( #内呼按钮9 )
      I_Contact( #"9层上呼分配" )
      I_Contact( #"9层下呼分配" )
      Move(in := 0, out1 => #目标楼层数9)
   END_RUNG
   RUNG wire#powerrail
      Contact( #内呼按钮10 )
      wire#w10
      Move(in := 10, out1 => #目标楼层数10)
   END_RUNG
   RUNG wire#powerrail
      Contact( #"10层下呼分配" )
   END_RUNG wire#w10
   RUNG wire#powerrail
      I_Contact( #内呼按钮10 )
      I_Contact( #"10层下呼分配" )
      Move(in := 0, out1 => #目标楼层数10)
   END_RUNG
   // the same network as SCL:
   IF #内呼按钮1 OR #"1层上呼分配" THEN #目标楼层数1 := 1; END_IF;
   IF NOT #内呼按钮1 AND NOT #"1层上呼分配" THEN #目标楼层数1 := 0; END_IF;
   IF #内呼按钮2 OR #"2层上呼分配" OR #"2层下呼分配" THEN #目标楼层数2 := 2; END_IF;
   IF NOT #内呼按钮2 AND NOT #"2层上呼分配" AND NOT #"2层下呼分配" THEN #目标楼层数2 := 0; END_IF;
   IF #内呼按钮3 OR #"3层上呼分配" OR #"3层下呼分配" THEN #目标楼层数3 := 3; END_IF;
   IF NOT #内呼按钮3 AND NOT #"3层下呼分配" AND NOT #"3层上呼分配" THEN #目标楼层数3 := 0; END_IF;
   IF #内呼按钮4 OR #"4层上呼分配" OR #"4层下呼分配" THEN #目标楼层数4 := 4; END_IF;
   IF NOT #内呼按钮4 AND NOT #"4层下呼分配" AND NOT #"4层上呼分配" THEN #目标楼层数4 := 0; END_IF;
   IF #内呼按钮5 OR #"5层上呼分配" OR #"5层下呼分配" THEN #目标楼层数5 := 5; END_IF;
   IF NOT #内呼按钮5 AND NOT #"5层下呼分配" AND NOT #"5层上呼分配" THEN #目标楼层数5 := 0; END_IF;
   IF #内呼按钮6 OR #"6层上呼分配" OR #"6层下呼分配" THEN #目标楼层数6 := 6; END_IF;
   IF NOT #内呼按钮6 AND NOT #"6层上呼分配" AND NOT #"6层下呼分配" THEN #目标楼层数6 := 0; END_IF;
   IF #内呼按钮7 OR #"7层上呼分配" OR #"7层下呼分配" THEN #目标楼层数7 := 7; END_IF;
   IF NOT #内呼按钮7 AND NOT #"7层上呼分配" AND NOT #"7层下呼分配" THEN #目标楼层数7 := 0; END_IF;
   IF #内呼按钮8 OR #"8层上呼分配" OR #"8层下呼分配" THEN #目标楼层数8 := 8; END_IF;
   IF NOT #内呼按钮8 AND NOT #"8层上呼分配" AND NOT #"8层下呼分配" THEN #目标楼层数8 := 0; END_IF;
   IF #内呼按钮9 OR #"9层上呼分配" OR #"9层下呼分配" THEN #目标楼层数9 := 9; END_IF;
   IF NOT #内呼按钮9 AND NOT #"9层上呼分配" AND NOT #"9层下呼分配" THEN #目标楼层数9 := 0; END_IF;
   IF #内呼按钮10 OR #"10层下呼分配" THEN #目标楼层数10 := 10; END_IF;
   IF NOT #内呼按钮10 AND NOT #"10层下呼分配" THEN #目标楼层数10 := 0; END_IF;
END_REGION

REGION Network 4: 外呼上面有目标
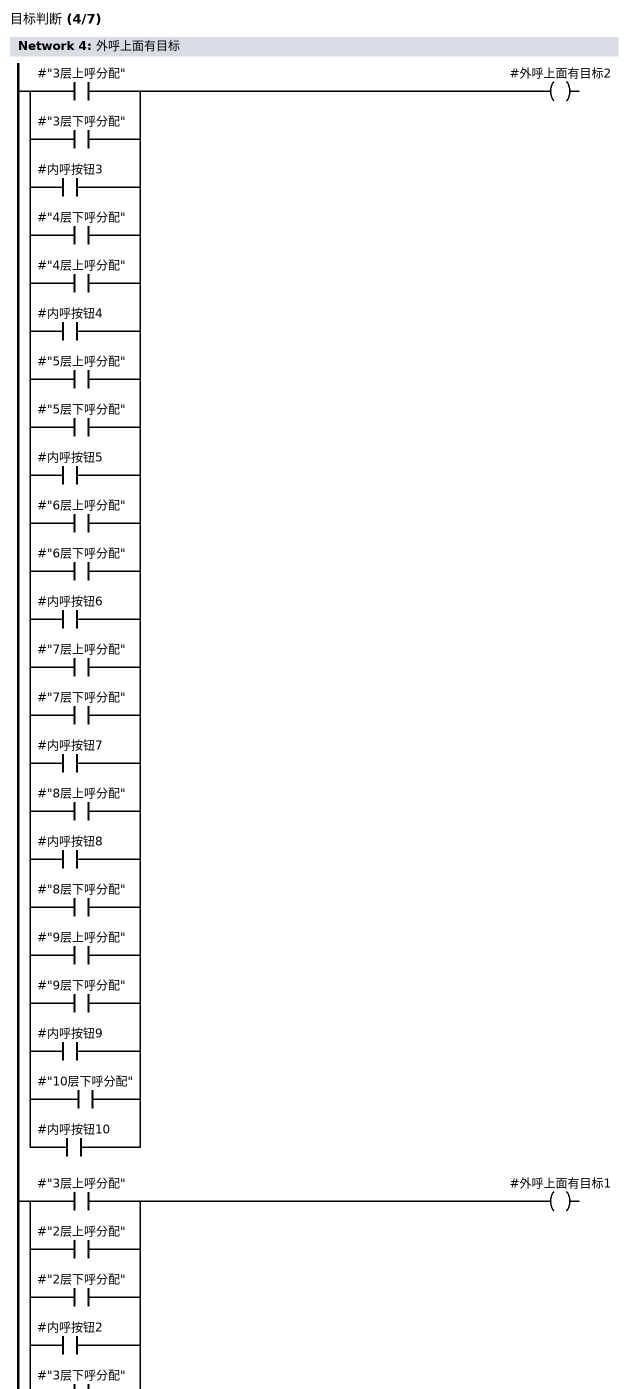
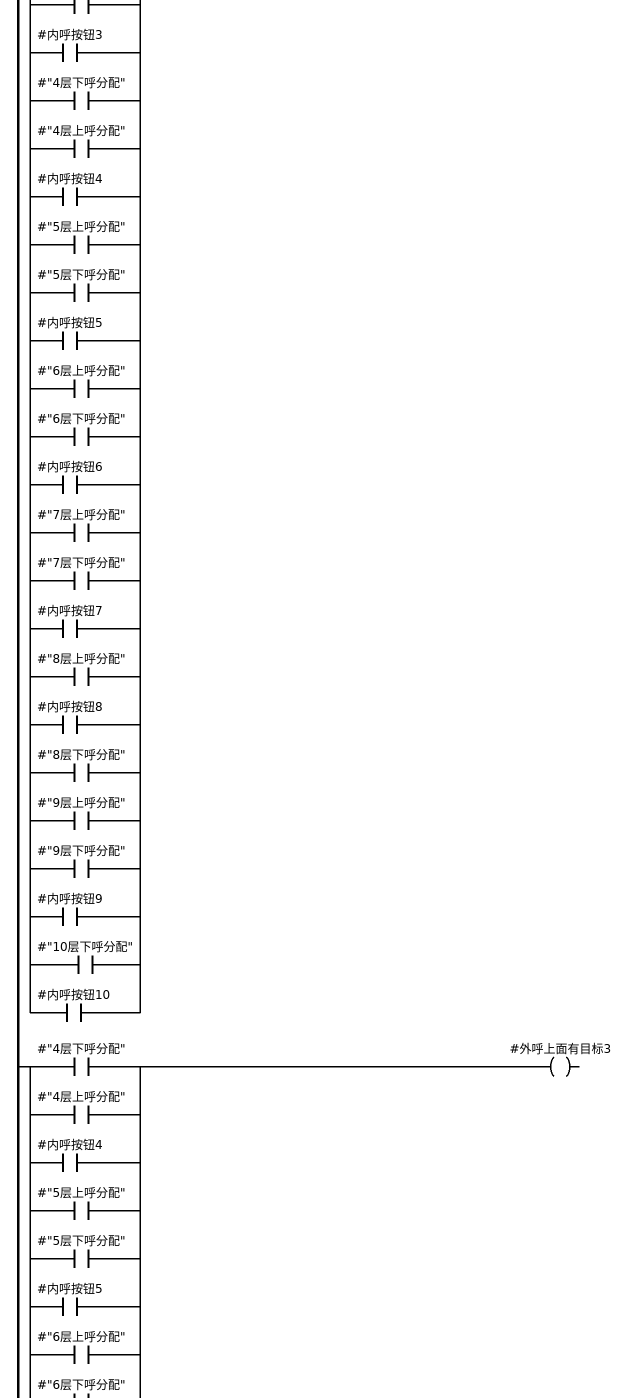
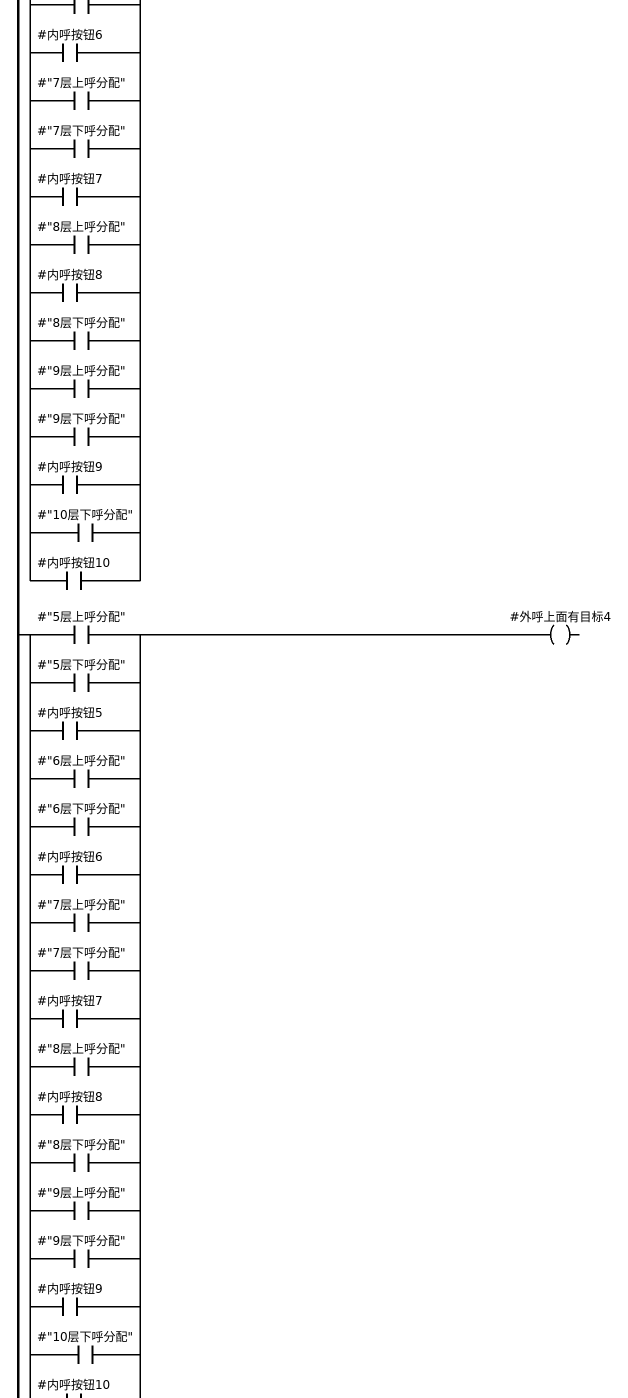
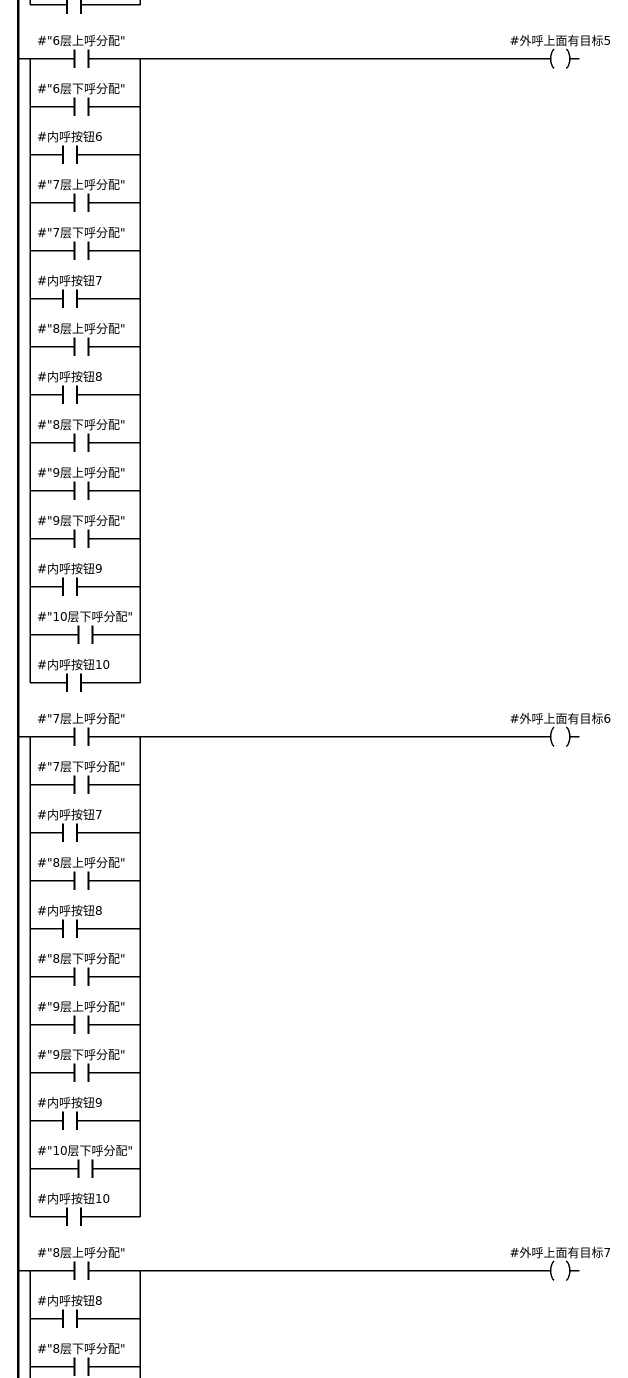
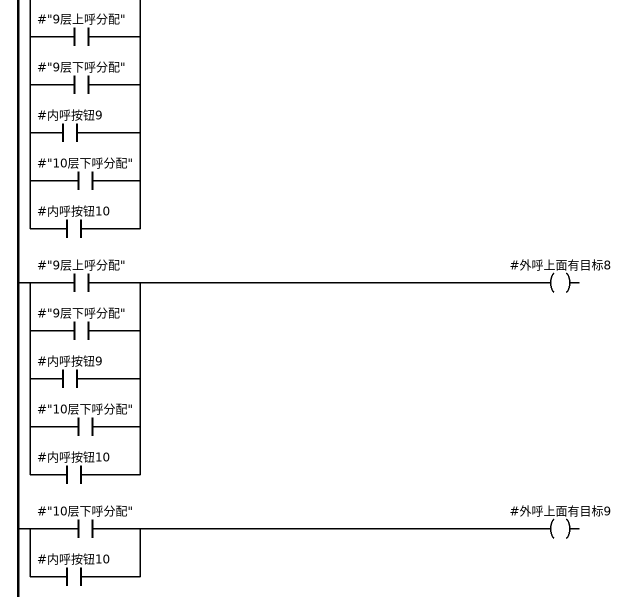
   RUNG wire#powerrail
      Contact( #"3层上呼分配" )
      wire#w1
      Coil( #外呼上面有目标2 )
   END_RUNG
   RUNG wire#powerrail
      Contact( #"3层下呼分配" )
   END_RUNG wire#w1
   RUNG wire#powerrail
      Contact( #内呼按钮3 )
   END_RUNG wire#w1
   RUNG wire#powerrail
      Contact( #"4层下呼分配" )
   END_RUNG wire#w1
   RUNG wire#powerrail
      Contact( #"4层上呼分配" )
   END_RUNG wire#w1
   RUNG wire#powerrail
      Contact( #内呼按钮4 )
   END_RUNG wire#w1
   RUNG wire#powerrail
      Contact( #"5层上呼分配" )
   END_RUNG wire#w1
   RUNG wire#powerrail
      Contact( #"5层下呼分配" )
   END_RUNG wire#w1
   RUNG wire#powerrail
      Contact( #内呼按钮5 )
   END_RUNG wire#w1
   RUNG wire#powerrail
      Contact( #"6层上呼分配" )
   END_RUNG wire#w1
   RUNG wire#powerrail
      Contact( #"6层下呼分配" )
   END_RUNG wire#w1
   RUNG wire#powerrail
      Contact( #内呼按钮6 )
   END_RUNG wire#w1
   RUNG wire#powerrail
      Contact( #"7层上呼分配" )
   END_RUNG wire#w1
   RUNG wire#powerrail
      Contact( #"7层下呼分配" )
   END_RUNG wire#w1
   RUNG wire#powerrail
      Contact( #内呼按钮7 )
   END_RUNG wire#w1
   RUNG wire#powerrail
      Contact( #"8层上呼分配" )
   END_RUNG wire#w1
   RUNG wire#powerrail
      Contact( #内呼按钮8 )
   END_RUNG wire#w1
   RUNG wire#powerrail
      Contact( #"8层下呼分配" )
   END_RUNG wire#w1
   RUNG wire#powerrail
      Contact( #"9层上呼分配" )
   END_RUNG wire#w1
   RUNG wire#powerrail
      Contact( #"9层下呼分配" )
   END_RUNG wire#w1
   RUNG wire#powerrail
      Contact( #内呼按钮9 )
   END_RUNG wire#w1
   RUNG wire#powerrail
      Contact( #"10层下呼分配" )
   END_RUNG wire#w1
   RUNG wire#powerrail
      Contact( #内呼按钮10 )
   END_RUNG wire#w1
   RUNG wire#powerrail
      Contact( #"3层上呼分配" )
      wire#w2
      Coil( #外呼上面有目标1 )
   END_RUNG
   RUNG wire#powerrail
      Contact( #"2层上呼分配" )
   END_RUNG wire#w2
   RUNG wire#powerrail
      Contact( #"2层下呼分配" )
   END_RUNG wire#w2
   RUNG wire#powerrail
      Contact( #内呼按钮2 )
   END_RUNG wire#w2
   RUNG wire#powerrail
      Contact( #"3层下呼分配" )
   END_RUNG wire#w2
   RUNG wire#powerrail
      Contact( #内呼按钮3 )
   END_RUNG wire#w2
   RUNG wire#powerrail
      Contact( #"4层下呼分配" )
   END_RUNG wire#w2
   RUNG wire#powerrail
      Contact( #"4层上呼分配" )
   END_RUNG wire#w2
   RUNG wire#powerrail
      Contact( #内呼按钮4 )
   END_RUNG wire#w2
   RUNG wire#powerrail
      Contact( #"5层上呼分配" )
   END_RUNG wire#w2
   RUNG wire#powerrail
      Contact( #"5层下呼分配" )
   END_RUNG wire#w2
   RUNG wire#powerrail
      Contact( #内呼按钮5 )
   END_RUNG wire#w2
   RUNG wire#powerrail
      Contact( #"6层上呼分配" )
   END_RUNG wire#w2
   RUNG wire#powerrail
      Contact( #"6层下呼分配" )
   END_RUNG wire#w2
   RUNG wire#powerrail
      Contact( #内呼按钮6 )
   END_RUNG wire#w2
   RUNG wire#powerrail
      Contact( #"7层上呼分配" )
   END_RUNG wire#w2
   RUNG wire#powerrail
      Contact( #"7层下呼分配" )
   END_RUNG wire#w2
   RUNG wire#powerrail
      Contact( #内呼按钮7 )
   END_RUNG wire#w2
   RUNG wire#powerrail
      Contact( #"8层上呼分配" )
   END_RUNG wire#w2
   RUNG wire#powerrail
      Contact( #内呼按钮8 )
   END_RUNG wire#w2
   RUNG wire#powerrail
      Contact( #"8层下呼分配" )
   END_RUNG wire#w2
   RUNG wire#powerrail
      Contact( #"9层上呼分配" )
   END_RUNG wire#w2
   RUNG wire#powerrail
      Contact( #"9层下呼分配" )
   END_RUNG wire#w2
   RUNG wire#powerrail
      Contact( #内呼按钮9 )
   END_RUNG wire#w2
   RUNG wire#powerrail
      Contact( #"10层下呼分配" )
   END_RUNG wire#w2
   RUNG wire#powerrail
      Contact( #内呼按钮10 )
   END_RUNG wire#w2
   RUNG wire#powerrail
      Contact( #"4层下呼分配" )
      wire#w3
      Coil( #外呼上面有目标3 )
   END_RUNG
   RUNG wire#powerrail
      Contact( #"4层上呼分配" )
   END_RUNG wire#w3
   RUNG wire#powerrail
      Contact( #内呼按钮4 )
   END_RUNG wire#w3
   RUNG wire#powerrail
      Contact( #"5层上呼分配" )
   END_RUNG wire#w3
   RUNG wire#powerrail
      Contact( #"5层下呼分配" )
   END_RUNG wire#w3
   RUNG wire#powerrail
      Contact( #内呼按钮5 )
   END_RUNG wire#w3
   RUNG wire#powerrail
      Contact( #"6层上呼分配" )
   END_RUNG wire#w3
   RUNG wire#powerrail
      Contact( #"6层下呼分配" )
   END_RUNG wire#w3
   RUNG wire#powerrail
      Contact( #内呼按钮6 )
   END_RUNG wire#w3
   RUNG wire#powerrail
      Contact( #"7层上呼分配" )
   END_RUNG wire#w3
   RUNG wire#powerrail
      Contact( #"7层下呼分配" )
   END_RUNG wire#w3
   RUNG wire#powerrail
      Contact( #内呼按钮7 )
   END_RUNG wire#w3
   RUNG wire#powerrail
      Contact( #"8层上呼分配" )
   END_RUNG wire#w3
   RUNG wire#powerrail
      Contact( #内呼按钮8 )
   END_RUNG wire#w3
   RUNG wire#powerrail
      Contact( #"8层下呼分配" )
   END_RUNG wire#w3
   RUNG wire#powerrail
      Contact( #"9层上呼分配" )
   END_RUNG wire#w3
   RUNG wire#powerrail
      Contact( #"9层下呼分配" )
   END_RUNG wire#w3
   RUNG wire#powerrail
      Contact( #内呼按钮9 )
   END_RUNG wire#w3
   RUNG wire#powerrail
      Contact( #"10层下呼分配" )
   END_RUNG wire#w3
   RUNG wire#powerrail
      Contact( #内呼按钮10 )
   END_RUNG wire#w3
   RUNG wire#powerrail
      Contact( #"5层上呼分配" )
      wire#w4
      Coil( #外呼上面有目标4 )
   END_RUNG
   RUNG wire#powerrail
      Contact( #"5层下呼分配" )
   END_RUNG wire#w4
   RUNG wire#powerrail
      Contact( #内呼按钮5 )
   END_RUNG wire#w4
   RUNG wire#powerrail
      Contact( #"6层上呼分配" )
   END_RUNG wire#w4
   RUNG wire#powerrail
      Contact( #"6层下呼分配" )
   END_RUNG wire#w4
   RUNG wire#powerrail
      Contact( #内呼按钮6 )
   END_RUNG wire#w4
   RUNG wire#powerrail
      Contact( #"7层上呼分配" )
   END_RUNG wire#w4
   RUNG wire#powerrail
      Contact( #"7层下呼分配" )
   END_RUNG wire#w4
   RUNG wire#powerrail
      Contact( #内呼按钮7 )
   END_RUNG wire#w4
   RUNG wire#powerrail
      Contact( #"8层上呼分配" )
   END_RUNG wire#w4
   RUNG wire#powerrail
      Contact( #内呼按钮8 )
   END_RUNG wire#w4
   RUNG wire#powerrail
      Contact( #"8层下呼分配" )
   END_RUNG wire#w4
   RUNG wire#powerrail
      Contact( #"9层上呼分配" )
   END_RUNG wire#w4
   RUNG wire#powerrail
      Contact( #"9层下呼分配" )
   END_RUNG wire#w4
   RUNG wire#powerrail
      Contact( #内呼按钮9 )
   END_RUNG wire#w4
   RUNG wire#powerrail
      Contact( #"10层下呼分配" )
   END_RUNG wire#w4
   RUNG wire#powerrail
      Contact( #内呼按钮10 )
   END_RUNG wire#w4
   RUNG wire#powerrail
      Contact( #"6层上呼分配" )
      wire#w5
      Coil( #外呼上面有目标5 )
   END_RUNG
   RUNG wire#powerrail
      Contact( #"6层下呼分配" )
   END_RUNG wire#w5
   RUNG wire#powerrail
      Contact( #内呼按钮6 )
   END_RUNG wire#w5
   RUNG wire#powerrail
      Contact( #"7层上呼分配" )
   END_RUNG wire#w5
   RUNG wire#powerrail
      Contact( #"7层下呼分配" )
   END_RUNG wire#w5
   RUNG wire#powerrail
      Contact( #内呼按钮7 )
   END_RUNG wire#w5
   RUNG wire#powerrail
      Contact( #"8层上呼分配" )
   END_RUNG wire#w5
   RUNG wire#powerrail
      Contact( #内呼按钮8 )
   END_RUNG wire#w5
   RUNG wire#powerrail
      Contact( #"8层下呼分配" )
   END_RUNG wire#w5
   RUNG wire#powerrail
      Contact( #"9层上呼分配" )
   END_RUNG wire#w5
   RUNG wire#powerrail
      Contact( #"9层下呼分配" )
   END_RUNG wire#w5
   RUNG wire#powerrail
      Contact( #内呼按钮9 )
   END_RUNG wire#w5
   RUNG wire#powerrail
      Contact( #"10层下呼分配" )
   END_RUNG wire#w5
   RUNG wire#powerrail
      Contact( #内呼按钮10 )
   END_RUNG wire#w5
   RUNG wire#powerrail
      Contact( #"7层上呼分配" )
      wire#w6
      Coil( #外呼上面有目标6 )
   END_RUNG
   RUNG wire#powerrail
      Contact( #"7层下呼分配" )
   END_RUNG wire#w6
   RUNG wire#powerrail
      Contact( #内呼按钮7 )
   END_RUNG wire#w6
   RUNG wire#powerrail
      Contact( #"8层上呼分配" )
   END_RUNG wire#w6
   RUNG wire#powerrail
      Contact( #内呼按钮8 )
   END_RUNG wire#w6
   RUNG wire#powerrail
      Contact( #"8层下呼分配" )
   END_RUNG wire#w6
   RUNG wire#powerrail
      Contact( #"9层上呼分配" )
   END_RUNG wire#w6
   RUNG wire#powerrail
      Contact( #"9层下呼分配" )
   END_RUNG wire#w6
   RUNG wire#powerrail
      Contact( #内呼按钮9 )
   END_RUNG wire#w6
   RUNG wire#powerrail
      Contact( #"10层下呼分配" )
   END_RUNG wire#w6
   RUNG wire#powerrail
      Contact( #内呼按钮10 )
   END_RUNG wire#w6
   RUNG wire#powerrail
      Contact( #"8层上呼分配" )
      wire#w7
      Coil( #外呼上面有目标7 )
   END_RUNG
   RUNG wire#powerrail
      Contact( #内呼按钮8 )
   END_RUNG wire#w7
   RUNG wire#powerrail
      Contact( #"8层下呼分配" )
   END_RUNG wire#w7
   RUNG wire#powerrail
      Contact( #"9层上呼分配" )
   END_RUNG wire#w7
   RUNG wire#powerrail
      Contact( #"9层下呼分配" )
   END_RUNG wire#w7
   RUNG wire#powerrail
      Contact( #内呼按钮9 )
   END_RUNG wire#w7
   RUNG wire#powerrail
      Contact( #"10层下呼分配" )
   END_RUNG wire#w7
   RUNG wire#powerrail
      Contact( #内呼按钮10 )
   END_RUNG wire#w7
   RUNG wire#powerrail
      Contact( #"9层上呼分配" )
      wire#w8
      Coil( #外呼上面有目标8 )
   END_RUNG
   RUNG wire#powerrail
      Contact( #"9层下呼分配" )
   END_RUNG wire#w8
   RUNG wire#powerrail
      Contact( #内呼按钮9 )
   END_RUNG wire#w8
   RUNG wire#powerrail
      Contact( #"10层下呼分配" )
   END_RUNG wire#w8
   RUNG wire#powerrail
      Contact( #内呼按钮10 )
   END_RUNG wire#w8
   RUNG wire#powerrail
      Contact( #"10层下呼分配" )
      wire#w9
      Coil( #外呼上面有目标9 )
   END_RUNG
   RUNG wire#powerrail
      Contact( #内呼按钮10 )
   END_RUNG wire#w9
   // the same network as SCL:
   #外呼上面有目标2 := #"3层上呼分配" OR #"3层下呼分配" OR #内呼按钮3 OR #"4层下呼分配" OR #"4层上呼分配" OR #内呼按钮4 OR #"5层上呼分配" OR #"5层下呼分配" OR #内呼按钮5 OR #"6层上呼分配" OR #"6层下呼分配" OR #内呼按钮6 OR #"7层上呼分配" OR #"7层下呼分配" OR #内呼按钮7 OR #"8层上呼分配" OR #内呼按钮8 OR #"8层下呼分配" OR #"9层上呼分配" OR #"9层下呼分配" OR #内呼按钮9 OR #"10层下呼分配" OR #内呼按钮10;
   #外呼上面有目标1 := #"3层上呼分配" OR #"2层上呼分配" OR #"2层下呼分配" OR #内呼按钮2 OR #"3层下呼分配" OR #内呼按钮3 OR #"4层下呼分配" OR #"4层上呼分配" OR #内呼按钮4 OR #"5层上呼分配" OR #"5层下呼分配" OR #内呼按钮5 OR #"6层上呼分配" OR #"6层下呼分配" OR #内呼按钮6 OR #"7层上呼分配" OR #"7层下呼分配" OR #内呼按钮7 OR #"8层上呼分配" OR #内呼按钮8 OR #"8层下呼分配" OR #"9层上呼分配" OR #"9层下呼分配" OR #内呼按钮9 OR #"10层下呼分配" OR #内呼按钮10;
   #外呼上面有目标3 := #"4层下呼分配" OR #"4层上呼分配" OR #内呼按钮4 OR #"5层上呼分配" OR #"5层下呼分配" OR #内呼按钮5 OR #"6层上呼分配" OR #"6层下呼分配" OR #内呼按钮6 OR #"7层上呼分配" OR #"7层下呼分配" OR #内呼按钮7 OR #"8层上呼分配" OR #内呼按钮8 OR #"8层下呼分配" OR #"9层上呼分配" OR #"9层下呼分配" OR #内呼按钮9 OR #"10层下呼分配" OR #内呼按钮10;
   #外呼上面有目标4 := #"5层上呼分配" OR #"5层下呼分配" OR #内呼按钮5 OR #"6层上呼分配" OR #"6层下呼分配" OR #内呼按钮6 OR #"7层上呼分配" OR #"7层下呼分配" OR #内呼按钮7 OR #"8层上呼分配" OR #内呼按钮8 OR #"8层下呼分配" OR #"9层上呼分配" OR #"9层下呼分配" OR #内呼按钮9 OR #"10层下呼分配" OR #内呼按钮10;
   #外呼上面有目标5 := #"6层上呼分配" OR #"6层下呼分配" OR #内呼按钮6 OR #"7层上呼分配" OR #"7层下呼分配" OR #内呼按钮7 OR #"8层上呼分配" OR #内呼按钮8 OR #"8层下呼分配" OR #"9层上呼分配" OR #"9层下呼分配" OR #内呼按钮9 OR #"10层下呼分配" OR #内呼按钮10;
   #外呼上面有目标6 := #"7层上呼分配" OR #"7层下呼分配" OR #内呼按钮7 OR #"8层上呼分配" OR #内呼按钮8 OR #"8层下呼分配" OR #"9层上呼分配" OR #"9层下呼分配" OR #内呼按钮9 OR #"10层下呼分配" OR #内呼按钮10;
   #外呼上面有目标7 := #"8层上呼分配" OR #内呼按钮8 OR #"8层下呼分配" OR #"9层上呼分配" OR #"9层下呼分配" OR #内呼按钮9 OR #"10层下呼分配" OR #内呼按钮10;
   #外呼上面有目标8 := #"9层上呼分配" OR #"9层下呼分配" OR #内呼按钮9 OR #"10层下呼分配" OR #内呼按钮10;
   #外呼上面有目标9 := #"10层下呼分配" OR #内呼按钮10;
END_REGION

